(* IEC 61131-3 sources: STAR-PLC-Agent/results/raw/batch_fresh_20261114/PUB015/functional/attempt_0001, 1 file *)

(* ---- test_program.st ---- *)
PROGRAM PLC_PRG
VAR
 BenchStep : UDINT := 0;
 BenchCalls : UDINT := 0;
 BenchDone : BOOL := FALSE;
 BenchUut0 : FB_Task;
 BenchUut1 : FB_Task;
 BenchUut2 : FB_Task;
 BenchUut3 : FB_Task;
 BenchUut4 : FB_Task;
 BenchUut5 : FB_Task;
 BenchUut6 : FB_Task;
 BenchUut7 : FB_Task;
 BenchUut8 : FB_Task;
 BenchUut9 : FB_Task;
 BenchUut10 : FB_Task;
 BenchUut11 : FB_Task;
 BenchUut12 : FB_Task;
 TraceIn_estop : ARRAY[0..126] OF BOOL;
 TraceIn_opeMode : ARRAY[0..126] OF BOOL;
 TraceIn_valveAStart : ARRAY[0..126] OF BOOL;
 TraceIn_valveBStart : ARRAY[0..126] OF BOOL;
 TraceIn_valveCStart : ARRAY[0..126] OF BOOL;
 TraceIn_valveDStart : ARRAY[0..126] OF BOOL;
 TraceIn_mixMotorStart : ARRAY[0..126] OF BOOL;
 TraceIn_autoStart : ARRAY[0..126] OF BOOL;
 TraceIn_processMode : ARRAY[0..126] OF BOOL;
 TraceIn_levelSensor : ARRAY[0..126] OF INT;
 TraceIn_mixMotorComplete : ARRAY[0..126] OF BOOL;
 TraceOut_valveARun : ARRAY[0..126] OF BOOL;
 TraceOut_valveBRun : ARRAY[0..126] OF BOOL;
 TraceOut_valveCRun : ARRAY[0..126] OF BOOL;
 TraceOut_valveDRun : ARRAY[0..126] OF BOOL;
 TraceOut_mixMotorRun : ARRAY[0..126] OF BOOL;
END_VAR

IF NOT BenchDone THEN
 CASE BenchStep OF
 0:
   BenchUut0.estop := TRUE;
   BenchUut0.opeMode := FALSE;
   BenchUut0.valveAStart := FALSE;
   BenchUut0.valveBStart := FALSE;
   BenchUut0.valveCStart := FALSE;
   BenchUut0.valveDStart := FALSE;
   BenchUut0.mixMotorStart := FALSE;
   BenchUut0.autoStart := FALSE;
   BenchUut0.processMode := FALSE;
   BenchUut0.levelSensor := INT#0;
   BenchUut0.mixMotorComplete := FALSE;
   TraceIn_estop[0] := BenchUut0.estop;
   TraceIn_opeMode[0] := BenchUut0.opeMode;
   TraceIn_valveAStart[0] := BenchUut0.valveAStart;
   TraceIn_valveBStart[0] := BenchUut0.valveBStart;
   TraceIn_valveCStart[0] := BenchUut0.valveCStart;
   TraceIn_valveDStart[0] := BenchUut0.valveDStart;
   TraceIn_mixMotorStart[0] := BenchUut0.mixMotorStart;
   TraceIn_autoStart[0] := BenchUut0.autoStart;
   TraceIn_processMode[0] := BenchUut0.processMode;
   TraceIn_levelSensor[0] := BenchUut0.levelSensor;
   TraceIn_mixMotorComplete[0] := BenchUut0.mixMotorComplete;
   BenchUut0();
   TraceOut_valveARun[0] := BenchUut0.valveARun;
   TraceOut_valveBRun[0] := BenchUut0.valveBRun;
   TraceOut_valveCRun[0] := BenchUut0.valveCRun;
   TraceOut_valveDRun[0] := BenchUut0.valveDRun;
   TraceOut_mixMotorRun[0] := BenchUut0.mixMotorRun;
   BenchCalls := BenchCalls + 1;
 1:
   BenchUut0.estop := TRUE;
   BenchUut0.opeMode := FALSE;
   BenchUut0.valveAStart := TRUE;
   BenchUut0.valveBStart := FALSE;
   BenchUut0.valveCStart := FALSE;
   BenchUut0.valveDStart := FALSE;
   BenchUut0.mixMotorStart := FALSE;
   BenchUut0.autoStart := FALSE;
   BenchUut0.processMode := FALSE;
   BenchUut0.levelSensor := INT#0;
   BenchUut0.mixMotorComplete := FALSE;
   TraceIn_estop[1] := BenchUut0.estop;
   TraceIn_opeMode[1] := BenchUut0.opeMode;
   TraceIn_valveAStart[1] := BenchUut0.valveAStart;
   TraceIn_valveBStart[1] := BenchUut0.valveBStart;
   TraceIn_valveCStart[1] := BenchUut0.valveCStart;
   TraceIn_valveDStart[1] := BenchUut0.valveDStart;
   TraceIn_mixMotorStart[1] := BenchUut0.mixMotorStart;
   TraceIn_autoStart[1] := BenchUut0.autoStart;
   TraceIn_processMode[1] := BenchUut0.processMode;
   TraceIn_levelSensor[1] := BenchUut0.levelSensor;
   TraceIn_mixMotorComplete[1] := BenchUut0.mixMotorComplete;
   BenchUut0();
   TraceOut_valveARun[1] := BenchUut0.valveARun;
   TraceOut_valveBRun[1] := BenchUut0.valveBRun;
   TraceOut_valveCRun[1] := BenchUut0.valveCRun;
   TraceOut_valveDRun[1] := BenchUut0.valveDRun;
   TraceOut_mixMotorRun[1] := BenchUut0.mixMotorRun;
   BenchCalls := BenchCalls + 1;
 2:
   BenchUut0.estop := TRUE;
   BenchUut0.opeMode := FALSE;
   BenchUut0.valveAStart := TRUE;
   BenchUut0.valveBStart := FALSE;
   BenchUut0.valveCStart := FALSE;
   BenchUut0.valveDStart := FALSE;
   BenchUut0.mixMotorStart := FALSE;
   BenchUut0.autoStart := FALSE;
   BenchUut0.processMode := FALSE;
   BenchUut0.levelSensor := INT#0;
   BenchUut0.mixMotorComplete := FALSE;
   TraceIn_estop[2] := BenchUut0.estop;
   TraceIn_opeMode[2] := BenchUut0.opeMode;
   TraceIn_valveAStart[2] := BenchUut0.valveAStart;
   TraceIn_valveBStart[2] := BenchUut0.valveBStart;
   TraceIn_valveCStart[2] := BenchUut0.valveCStart;
   TraceIn_valveDStart[2] := BenchUut0.valveDStart;
   TraceIn_mixMotorStart[2] := BenchUut0.mixMotorStart;
   TraceIn_autoStart[2] := BenchUut0.autoStart;
   TraceIn_processMode[2] := BenchUut0.processMode;
   TraceIn_levelSensor[2] := BenchUut0.levelSensor;
   TraceIn_mixMotorComplete[2] := BenchUut0.mixMotorComplete;
   BenchUut0();
   TraceOut_valveARun[2] := BenchUut0.valveARun;
   TraceOut_valveBRun[2] := BenchUut0.valveBRun;
   TraceOut_valveCRun[2] := BenchUut0.valveCRun;
   TraceOut_valveDRun[2] := BenchUut0.valveDRun;
   TraceOut_mixMotorRun[2] := BenchUut0.mixMotorRun;
   BenchCalls := BenchCalls + 1;
 3:
   BenchUut0.estop := TRUE;
   BenchUut0.opeMode := FALSE;
   BenchUut0.valveAStart := FALSE;
   BenchUut0.valveBStart := FALSE;
   BenchUut0.valveCStart := FALSE;
   BenchUut0.valveDStart := FALSE;
   BenchUut0.mixMotorStart := FALSE;
   BenchUut0.autoStart := FALSE;
   BenchUut0.processMode := FALSE;
   BenchUut0.levelSensor := INT#0;
   BenchUut0.mixMotorComplete := FALSE;
   TraceIn_estop[3] := BenchUut0.estop;
   TraceIn_opeMode[3] := BenchUut0.opeMode;
   TraceIn_valveAStart[3] := BenchUut0.valveAStart;
   TraceIn_valveBStart[3] := BenchUut0.valveBStart;
   TraceIn_valveCStart[3] := BenchUut0.valveCStart;
   TraceIn_valveDStart[3] := BenchUut0.valveDStart;
   TraceIn_mixMotorStart[3] := BenchUut0.mixMotorStart;
   TraceIn_autoStart[3] := BenchUut0.autoStart;
   TraceIn_processMode[3] := BenchUut0.processMode;
   TraceIn_levelSensor[3] := BenchUut0.levelSensor;
   TraceIn_mixMotorComplete[3] := BenchUut0.mixMotorComplete;
   BenchUut0();
   TraceOut_valveARun[3] := BenchUut0.valveARun;
   TraceOut_valveBRun[3] := BenchUut0.valveBRun;
   TraceOut_valveCRun[3] := BenchUut0.valveCRun;
   TraceOut_valveDRun[3] := BenchUut0.valveDRun;
   TraceOut_mixMotorRun[3] := BenchUut0.mixMotorRun;
   BenchCalls := BenchCalls + 1;
 4:
   BenchUut0.estop := TRUE;
   BenchUut0.opeMode := FALSE;
   BenchUut0.valveAStart := TRUE;
   BenchUut0.valveBStart := FALSE;
   BenchUut0.valveCStart := FALSE;
   BenchUut0.valveDStart := FALSE;
   BenchUut0.mixMotorStart := FALSE;
   BenchUut0.autoStart := FALSE;
   BenchUut0.processMode := FALSE;
   BenchUut0.levelSensor := INT#0;
   BenchUut0.mixMotorComplete := FALSE;
   TraceIn_estop[4] := BenchUut0.estop;
   TraceIn_opeMode[4] := BenchUut0.opeMode;
   TraceIn_valveAStart[4] := BenchUut0.valveAStart;
   TraceIn_valveBStart[4] := BenchUut0.valveBStart;
   TraceIn_valveCStart[4] := BenchUut0.valveCStart;
   TraceIn_valveDStart[4] := BenchUut0.valveDStart;
   TraceIn_mixMotorStart[4] := BenchUut0.mixMotorStart;
   TraceIn_autoStart[4] := BenchUut0.autoStart;
   TraceIn_processMode[4] := BenchUut0.processMode;
   TraceIn_levelSensor[4] := BenchUut0.levelSensor;
   TraceIn_mixMotorComplete[4] := BenchUut0.mixMotorComplete;
   BenchUut0();
   TraceOut_valveARun[4] := BenchUut0.valveARun;
   TraceOut_valveBRun[4] := BenchUut0.valveBRun;
   TraceOut_valveCRun[4] := BenchUut0.valveCRun;
   TraceOut_valveDRun[4] := BenchUut0.valveDRun;
   TraceOut_mixMotorRun[4] := BenchUut0.mixMotorRun;
   BenchCalls := BenchCalls + 1;
 5:
   BenchUut0.estop := TRUE;
   BenchUut0.opeMode := FALSE;
   BenchUut0.valveAStart := FALSE;
   BenchUut0.valveBStart := TRUE;
   BenchUut0.valveCStart := TRUE;
   BenchUut0.valveDStart := TRUE;
   BenchUut0.mixMotorStart := TRUE;
   BenchUut0.autoStart := FALSE;
   BenchUut0.processMode := FALSE;
   BenchUut0.levelSensor := INT#0;
   BenchUut0.mixMotorComplete := FALSE;
   TraceIn_estop[5] := BenchUut0.estop;
   TraceIn_opeMode[5] := BenchUut0.opeMode;
   TraceIn_valveAStart[5] := BenchUut0.valveAStart;
   TraceIn_valveBStart[5] := BenchUut0.valveBStart;
   TraceIn_valveCStart[5] := BenchUut0.valveCStart;
   TraceIn_valveDStart[5] := BenchUut0.valveDStart;
   TraceIn_mixMotorStart[5] := BenchUut0.mixMotorStart;
   TraceIn_autoStart[5] := BenchUut0.autoStart;
   TraceIn_processMode[5] := BenchUut0.processMode;
   TraceIn_levelSensor[5] := BenchUut0.levelSensor;
   TraceIn_mixMotorComplete[5] := BenchUut0.mixMotorComplete;
   BenchUut0();
   TraceOut_valveARun[5] := BenchUut0.valveARun;
   TraceOut_valveBRun[5] := BenchUut0.valveBRun;
   TraceOut_valveCRun[5] := BenchUut0.valveCRun;
   TraceOut_valveDRun[5] := BenchUut0.valveDRun;
   TraceOut_mixMotorRun[5] := BenchUut0.mixMotorRun;
   BenchCalls := BenchCalls + 1;
 6:
   BenchUut0.estop := FALSE;
   BenchUut0.opeMode := FALSE;
   BenchUut0.valveAStart := FALSE;
   BenchUut0.valveBStart := FALSE;
   BenchUut0.valveCStart := FALSE;
   BenchUut0.valveDStart := FALSE;
   BenchUut0.mixMotorStart := FALSE;
   BenchUut0.autoStart := FALSE;
   BenchUut0.processMode := FALSE;
   BenchUut0.levelSensor := INT#0;
   BenchUut0.mixMotorComplete := FALSE;
   TraceIn_estop[6] := BenchUut0.estop;
   TraceIn_opeMode[6] := BenchUut0.opeMode;
   TraceIn_valveAStart[6] := BenchUut0.valveAStart;
   TraceIn_valveBStart[6] := BenchUut0.valveBStart;
   TraceIn_valveCStart[6] := BenchUut0.valveCStart;
   TraceIn_valveDStart[6] := BenchUut0.valveDStart;
   TraceIn_mixMotorStart[6] := BenchUut0.mixMotorStart;
   TraceIn_autoStart[6] := BenchUut0.autoStart;
   TraceIn_processMode[6] := BenchUut0.processMode;
   TraceIn_levelSensor[6] := BenchUut0.levelSensor;
   TraceIn_mixMotorComplete[6] := BenchUut0.mixMotorComplete;
   BenchUut0();
   TraceOut_valveARun[6] := BenchUut0.valveARun;
   TraceOut_valveBRun[6] := BenchUut0.valveBRun;
   TraceOut_valveCRun[6] := BenchUut0.valveCRun;
   TraceOut_valveDRun[6] := BenchUut0.valveDRun;
   TraceOut_mixMotorRun[6] := BenchUut0.mixMotorRun;
   BenchCalls := BenchCalls + 1;
 7:
   BenchUut1.estop := TRUE;
   BenchUut1.opeMode := TRUE;
   BenchUut1.valveAStart := FALSE;
   BenchUut1.valveBStart := FALSE;
   BenchUut1.valveCStart := FALSE;
   BenchUut1.valveDStart := FALSE;
   BenchUut1.mixMotorStart := FALSE;
   BenchUut1.autoStart := FALSE;
   BenchUut1.processMode := FALSE;
   BenchUut1.levelSensor := INT#0;
   BenchUut1.mixMotorComplete := FALSE;
   TraceIn_estop[7] := BenchUut1.estop;
   TraceIn_opeMode[7] := BenchUut1.opeMode;
   TraceIn_valveAStart[7] := BenchUut1.valveAStart;
   TraceIn_valveBStart[7] := BenchUut1.valveBStart;
   TraceIn_valveCStart[7] := BenchUut1.valveCStart;
   TraceIn_valveDStart[7] := BenchUut1.valveDStart;
   TraceIn_mixMotorStart[7] := BenchUut1.mixMotorStart;
   TraceIn_autoStart[7] := BenchUut1.autoStart;
   TraceIn_processMode[7] := BenchUut1.processMode;
   TraceIn_levelSensor[7] := BenchUut1.levelSensor;
   TraceIn_mixMotorComplete[7] := BenchUut1.mixMotorComplete;
   BenchUut1();
   TraceOut_valveARun[7] := BenchUut1.valveARun;
   TraceOut_valveBRun[7] := BenchUut1.valveBRun;
   TraceOut_valveCRun[7] := BenchUut1.valveCRun;
   TraceOut_valveDRun[7] := BenchUut1.valveDRun;
   TraceOut_mixMotorRun[7] := BenchUut1.mixMotorRun;
   BenchCalls := BenchCalls + 1;
 8:
   BenchUut1.estop := TRUE;
   BenchUut1.opeMode := TRUE;
   BenchUut1.valveAStart := FALSE;
   BenchUut1.valveBStart := FALSE;
   BenchUut1.valveCStart := FALSE;
   BenchUut1.valveDStart := FALSE;
   BenchUut1.mixMotorStart := FALSE;
   BenchUut1.autoStart := TRUE;
   BenchUut1.processMode := FALSE;
   BenchUut1.levelSensor := INT#0;
   BenchUut1.mixMotorComplete := FALSE;
   TraceIn_estop[8] := BenchUut1.estop;
   TraceIn_opeMode[8] := BenchUut1.opeMode;
   TraceIn_valveAStart[8] := BenchUut1.valveAStart;
   TraceIn_valveBStart[8] := BenchUut1.valveBStart;
   TraceIn_valveCStart[8] := BenchUut1.valveCStart;
   TraceIn_valveDStart[8] := BenchUut1.valveDStart;
   TraceIn_mixMotorStart[8] := BenchUut1.mixMotorStart;
   TraceIn_autoStart[8] := BenchUut1.autoStart;
   TraceIn_processMode[8] := BenchUut1.processMode;
   TraceIn_levelSensor[8] := BenchUut1.levelSensor;
   TraceIn_mixMotorComplete[8] := BenchUut1.mixMotorComplete;
   BenchUut1();
   TraceOut_valveARun[8] := BenchUut1.valveARun;
   TraceOut_valveBRun[8] := BenchUut1.valveBRun;
   TraceOut_valveCRun[8] := BenchUut1.valveCRun;
   TraceOut_valveDRun[8] := BenchUut1.valveDRun;
   TraceOut_mixMotorRun[8] := BenchUut1.mixMotorRun;
   BenchCalls := BenchCalls + 1;
 9:
   BenchUut1.estop := TRUE;
   BenchUut1.opeMode := TRUE;
   BenchUut1.valveAStart := FALSE;
   BenchUut1.valveBStart := FALSE;
   BenchUut1.valveCStart := FALSE;
   BenchUut1.valveDStart := FALSE;
   BenchUut1.mixMotorStart := FALSE;
   BenchUut1.autoStart := FALSE;
   BenchUut1.processMode := FALSE;
   BenchUut1.levelSensor := INT#49;
   BenchUut1.mixMotorComplete := FALSE;
   TraceIn_estop[9] := BenchUut1.estop;
   TraceIn_opeMode[9] := BenchUut1.opeMode;
   TraceIn_valveAStart[9] := BenchUut1.valveAStart;
   TraceIn_valveBStart[9] := BenchUut1.valveBStart;
   TraceIn_valveCStart[9] := BenchUut1.valveCStart;
   TraceIn_valveDStart[9] := BenchUut1.valveDStart;
   TraceIn_mixMotorStart[9] := BenchUut1.mixMotorStart;
   TraceIn_autoStart[9] := BenchUut1.autoStart;
   TraceIn_processMode[9] := BenchUut1.processMode;
   TraceIn_levelSensor[9] := BenchUut1.levelSensor;
   TraceIn_mixMotorComplete[9] := BenchUut1.mixMotorComplete;
   BenchUut1();
   TraceOut_valveARun[9] := BenchUut1.valveARun;
   TraceOut_valveBRun[9] := BenchUut1.valveBRun;
   TraceOut_valveCRun[9] := BenchUut1.valveCRun;
   TraceOut_valveDRun[9] := BenchUut1.valveDRun;
   TraceOut_mixMotorRun[9] := BenchUut1.mixMotorRun;
   BenchCalls := BenchCalls + 1;
 10:
   BenchUut1.estop := TRUE;
   BenchUut1.opeMode := TRUE;
   BenchUut1.valveAStart := FALSE;
   BenchUut1.valveBStart := FALSE;
   BenchUut1.valveCStart := FALSE;
   BenchUut1.valveDStart := FALSE;
   BenchUut1.mixMotorStart := FALSE;
   BenchUut1.autoStart := FALSE;
   BenchUut1.processMode := FALSE;
   BenchUut1.levelSensor := INT#50;
   BenchUut1.mixMotorComplete := FALSE;
   TraceIn_estop[10] := BenchUut1.estop;
   TraceIn_opeMode[10] := BenchUut1.opeMode;
   TraceIn_valveAStart[10] := BenchUut1.valveAStart;
   TraceIn_valveBStart[10] := BenchUut1.valveBStart;
   TraceIn_valveCStart[10] := BenchUut1.valveCStart;
   TraceIn_valveDStart[10] := BenchUut1.valveDStart;
   TraceIn_mixMotorStart[10] := BenchUut1.mixMotorStart;
   TraceIn_autoStart[10] := BenchUut1.autoStart;
   TraceIn_processMode[10] := BenchUut1.processMode;
   TraceIn_levelSensor[10] := BenchUut1.levelSensor;
   TraceIn_mixMotorComplete[10] := BenchUut1.mixMotorComplete;
   BenchUut1();
   TraceOut_valveARun[10] := BenchUut1.valveARun;
   TraceOut_valveBRun[10] := BenchUut1.valveBRun;
   TraceOut_valveCRun[10] := BenchUut1.valveCRun;
   TraceOut_valveDRun[10] := BenchUut1.valveDRun;
   TraceOut_mixMotorRun[10] := BenchUut1.mixMotorRun;
   BenchCalls := BenchCalls + 1;
 11:
   BenchUut1.estop := TRUE;
   BenchUut1.opeMode := TRUE;
   BenchUut1.valveAStart := FALSE;
   BenchUut1.valveBStart := FALSE;
   BenchUut1.valveCStart := FALSE;
   BenchUut1.valveDStart := FALSE;
   BenchUut1.mixMotorStart := FALSE;
   BenchUut1.autoStart := FALSE;
   BenchUut1.processMode := FALSE;
   BenchUut1.levelSensor := INT#80;
   BenchUut1.mixMotorComplete := FALSE;
   TraceIn_estop[11] := BenchUut1.estop;
   TraceIn_opeMode[11] := BenchUut1.opeMode;
   TraceIn_valveAStart[11] := BenchUut1.valveAStart;
   TraceIn_valveBStart[11] := BenchUut1.valveBStart;
   TraceIn_valveCStart[11] := BenchUut1.valveCStart;
   TraceIn_valveDStart[11] := BenchUut1.valveDStart;
   TraceIn_mixMotorStart[11] := BenchUut1.mixMotorStart;
   TraceIn_autoStart[11] := BenchUut1.autoStart;
   TraceIn_processMode[11] := BenchUut1.processMode;
   TraceIn_levelSensor[11] := BenchUut1.levelSensor;
   TraceIn_mixMotorComplete[11] := BenchUut1.mixMotorComplete;
   BenchUut1();
   TraceOut_valveARun[11] := BenchUut1.valveARun;
   TraceOut_valveBRun[11] := BenchUut1.valveBRun;
   TraceOut_valveCRun[11] := BenchUut1.valveCRun;
   TraceOut_valveDRun[11] := BenchUut1.valveDRun;
   TraceOut_mixMotorRun[11] := BenchUut1.mixMotorRun;
   BenchCalls := BenchCalls + 1;
 12:
   BenchUut1.estop := TRUE;
   BenchUut1.opeMode := TRUE;
   BenchUut1.valveAStart := FALSE;
   BenchUut1.valveBStart := FALSE;
   BenchUut1.valveCStart := FALSE;
   BenchUut1.valveDStart := FALSE;
   BenchUut1.mixMotorStart := FALSE;
   BenchUut1.autoStart := FALSE;
   BenchUut1.processMode := FALSE;
   BenchUut1.levelSensor := INT#80;
   BenchUut1.mixMotorComplete := TRUE;
   TraceIn_estop[12] := BenchUut1.estop;
   TraceIn_opeMode[12] := BenchUut1.opeMode;
   TraceIn_valveAStart[12] := BenchUut1.valveAStart;
   TraceIn_valveBStart[12] := BenchUut1.valveBStart;
   TraceIn_valveCStart[12] := BenchUut1.valveCStart;
   TraceIn_valveDStart[12] := BenchUut1.valveDStart;
   TraceIn_mixMotorStart[12] := BenchUut1.mixMotorStart;
   TraceIn_autoStart[12] := BenchUut1.autoStart;
   TraceIn_processMode[12] := BenchUut1.processMode;
   TraceIn_levelSensor[12] := BenchUut1.levelSensor;
   TraceIn_mixMotorComplete[12] := BenchUut1.mixMotorComplete;
   BenchUut1();
   TraceOut_valveARun[12] := BenchUut1.valveARun;
   TraceOut_valveBRun[12] := BenchUut1.valveBRun;
   TraceOut_valveCRun[12] := BenchUut1.valveCRun;
   TraceOut_valveDRun[12] := BenchUut1.valveDRun;
   TraceOut_mixMotorRun[12] := BenchUut1.mixMotorRun;
   BenchCalls := BenchCalls + 1;
 13:
   BenchUut1.estop := FALSE;
   BenchUut1.opeMode := TRUE;
   BenchUut1.valveAStart := FALSE;
   BenchUut1.valveBStart := FALSE;
   BenchUut1.valveCStart := FALSE;
   BenchUut1.valveDStart := FALSE;
   BenchUut1.mixMotorStart := FALSE;
   BenchUut1.autoStart := FALSE;
   BenchUut1.processMode := FALSE;
   BenchUut1.levelSensor := INT#0;
   BenchUut1.mixMotorComplete := FALSE;
   TraceIn_estop[13] := BenchUut1.estop;
   TraceIn_opeMode[13] := BenchUut1.opeMode;
   TraceIn_valveAStart[13] := BenchUut1.valveAStart;
   TraceIn_valveBStart[13] := BenchUut1.valveBStart;
   TraceIn_valveCStart[13] := BenchUut1.valveCStart;
   TraceIn_valveDStart[13] := BenchUut1.valveDStart;
   TraceIn_mixMotorStart[13] := BenchUut1.mixMotorStart;
   TraceIn_autoStart[13] := BenchUut1.autoStart;
   TraceIn_processMode[13] := BenchUut1.processMode;
   TraceIn_levelSensor[13] := BenchUut1.levelSensor;
   TraceIn_mixMotorComplete[13] := BenchUut1.mixMotorComplete;
   BenchUut1();
   TraceOut_valveARun[13] := BenchUut1.valveARun;
   TraceOut_valveBRun[13] := BenchUut1.valveBRun;
   TraceOut_valveCRun[13] := BenchUut1.valveCRun;
   TraceOut_valveDRun[13] := BenchUut1.valveDRun;
   TraceOut_mixMotorRun[13] := BenchUut1.mixMotorRun;
   BenchCalls := BenchCalls + 1;
 14:
   BenchUut2.estop := TRUE;
   BenchUut2.opeMode := TRUE;
   BenchUut2.valveAStart := FALSE;
   BenchUut2.valveBStart := FALSE;
   BenchUut2.valveCStart := FALSE;
   BenchUut2.valveDStart := FALSE;
   BenchUut2.mixMotorStart := FALSE;
   BenchUut2.autoStart := FALSE;
   BenchUut2.processMode := FALSE;
   BenchUut2.levelSensor := INT#0;
   BenchUut2.mixMotorComplete := FALSE;
   TraceIn_estop[14] := BenchUut2.estop;
   TraceIn_opeMode[14] := BenchUut2.opeMode;
   TraceIn_valveAStart[14] := BenchUut2.valveAStart;
   TraceIn_valveBStart[14] := BenchUut2.valveBStart;
   TraceIn_valveCStart[14] := BenchUut2.valveCStart;
   TraceIn_valveDStart[14] := BenchUut2.valveDStart;
   TraceIn_mixMotorStart[14] := BenchUut2.mixMotorStart;
   TraceIn_autoStart[14] := BenchUut2.autoStart;
   TraceIn_processMode[14] := BenchUut2.processMode;
   TraceIn_levelSensor[14] := BenchUut2.levelSensor;
   TraceIn_mixMotorComplete[14] := BenchUut2.mixMotorComplete;
   BenchUut2();
   TraceOut_valveARun[14] := BenchUut2.valveARun;
   TraceOut_valveBRun[14] := BenchUut2.valveBRun;
   TraceOut_valveCRun[14] := BenchUut2.valveCRun;
   TraceOut_valveDRun[14] := BenchUut2.valveDRun;
   TraceOut_mixMotorRun[14] := BenchUut2.mixMotorRun;
   BenchCalls := BenchCalls + 1;
 15:
   BenchUut2.estop := TRUE;
   BenchUut2.opeMode := TRUE;
   BenchUut2.valveAStart := FALSE;
   BenchUut2.valveBStart := FALSE;
   BenchUut2.valveCStart := FALSE;
   BenchUut2.valveDStart := FALSE;
   BenchUut2.mixMotorStart := FALSE;
   BenchUut2.autoStart := TRUE;
   BenchUut2.processMode := TRUE;
   BenchUut2.levelSensor := INT#0;
   BenchUut2.mixMotorComplete := FALSE;
   TraceIn_estop[15] := BenchUut2.estop;
   TraceIn_opeMode[15] := BenchUut2.opeMode;
   TraceIn_valveAStart[15] := BenchUut2.valveAStart;
   TraceIn_valveBStart[15] := BenchUut2.valveBStart;
   TraceIn_valveCStart[15] := BenchUut2.valveCStart;
   TraceIn_valveDStart[15] := BenchUut2.valveDStart;
   TraceIn_mixMotorStart[15] := BenchUut2.mixMotorStart;
   TraceIn_autoStart[15] := BenchUut2.autoStart;
   TraceIn_processMode[15] := BenchUut2.processMode;
   TraceIn_levelSensor[15] := BenchUut2.levelSensor;
   TraceIn_mixMotorComplete[15] := BenchUut2.mixMotorComplete;
   BenchUut2();
   TraceOut_valveARun[15] := BenchUut2.valveARun;
   TraceOut_valveBRun[15] := BenchUut2.valveBRun;
   TraceOut_valveCRun[15] := BenchUut2.valveCRun;
   TraceOut_valveDRun[15] := BenchUut2.valveDRun;
   TraceOut_mixMotorRun[15] := BenchUut2.mixMotorRun;
   BenchCalls := BenchCalls + 1;
 16:
   BenchUut2.estop := TRUE;
   BenchUut2.opeMode := TRUE;
   BenchUut2.valveAStart := FALSE;
   BenchUut2.valveBStart := FALSE;
   BenchUut2.valveCStart := FALSE;
   BenchUut2.valveDStart := FALSE;
   BenchUut2.mixMotorStart := FALSE;
   BenchUut2.autoStart := FALSE;
   BenchUut2.processMode := TRUE;
   BenchUut2.levelSensor := INT#55;
   BenchUut2.mixMotorComplete := FALSE;
   TraceIn_estop[16] := BenchUut2.estop;
   TraceIn_opeMode[16] := BenchUut2.opeMode;
   TraceIn_valveAStart[16] := BenchUut2.valveAStart;
   TraceIn_valveBStart[16] := BenchUut2.valveBStart;
   TraceIn_valveCStart[16] := BenchUut2.valveCStart;
   TraceIn_valveDStart[16] := BenchUut2.valveDStart;
   TraceIn_mixMotorStart[16] := BenchUut2.mixMotorStart;
   TraceIn_autoStart[16] := BenchUut2.autoStart;
   TraceIn_processMode[16] := BenchUut2.processMode;
   TraceIn_levelSensor[16] := BenchUut2.levelSensor;
   TraceIn_mixMotorComplete[16] := BenchUut2.mixMotorComplete;
   BenchUut2();
   TraceOut_valveARun[16] := BenchUut2.valveARun;
   TraceOut_valveBRun[16] := BenchUut2.valveBRun;
   TraceOut_valveCRun[16] := BenchUut2.valveCRun;
   TraceOut_valveDRun[16] := BenchUut2.valveDRun;
   TraceOut_mixMotorRun[16] := BenchUut2.mixMotorRun;
   BenchCalls := BenchCalls + 1;
 17:
   BenchUut2.estop := TRUE;
   BenchUut2.opeMode := TRUE;
   BenchUut2.valveAStart := FALSE;
   BenchUut2.valveBStart := FALSE;
   BenchUut2.valveCStart := FALSE;
   BenchUut2.valveDStart := FALSE;
   BenchUut2.mixMotorStart := FALSE;
   BenchUut2.autoStart := FALSE;
   BenchUut2.processMode := TRUE;
   BenchUut2.levelSensor := INT#85;
   BenchUut2.mixMotorComplete := FALSE;
   TraceIn_estop[17] := BenchUut2.estop;
   TraceIn_opeMode[17] := BenchUut2.opeMode;
   TraceIn_valveAStart[17] := BenchUut2.valveAStart;
   TraceIn_valveBStart[17] := BenchUut2.valveBStart;
   TraceIn_valveCStart[17] := BenchUut2.valveCStart;
   TraceIn_valveDStart[17] := BenchUut2.valveDStart;
   TraceIn_mixMotorStart[17] := BenchUut2.mixMotorStart;
   TraceIn_autoStart[17] := BenchUut2.autoStart;
   TraceIn_processMode[17] := BenchUut2.processMode;
   TraceIn_levelSensor[17] := BenchUut2.levelSensor;
   TraceIn_mixMotorComplete[17] := BenchUut2.mixMotorComplete;
   BenchUut2();
   TraceOut_valveARun[17] := BenchUut2.valveARun;
   TraceOut_valveBRun[17] := BenchUut2.valveBRun;
   TraceOut_valveCRun[17] := BenchUut2.valveCRun;
   TraceOut_valveDRun[17] := BenchUut2.valveDRun;
   TraceOut_mixMotorRun[17] := BenchUut2.mixMotorRun;
   BenchCalls := BenchCalls + 1;
 18:
   BenchUut2.estop := TRUE;
   BenchUut2.opeMode := TRUE;
   BenchUut2.valveAStart := FALSE;
   BenchUut2.valveBStart := FALSE;
   BenchUut2.valveCStart := FALSE;
   BenchUut2.valveDStart := FALSE;
   BenchUut2.mixMotorStart := FALSE;
   BenchUut2.autoStart := FALSE;
   BenchUut2.processMode := TRUE;
   BenchUut2.levelSensor := INT#99;
   BenchUut2.mixMotorComplete := FALSE;
   TraceIn_estop[18] := BenchUut2.estop;
   TraceIn_opeMode[18] := BenchUut2.opeMode;
   TraceIn_valveAStart[18] := BenchUut2.valveAStart;
   TraceIn_valveBStart[18] := BenchUut2.valveBStart;
   TraceIn_valveCStart[18] := BenchUut2.valveCStart;
   TraceIn_valveDStart[18] := BenchUut2.valveDStart;
   TraceIn_mixMotorStart[18] := BenchUut2.mixMotorStart;
   TraceIn_autoStart[18] := BenchUut2.autoStart;
   TraceIn_processMode[18] := BenchUut2.processMode;
   TraceIn_levelSensor[18] := BenchUut2.levelSensor;
   TraceIn_mixMotorComplete[18] := BenchUut2.mixMotorComplete;
   BenchUut2();
   TraceOut_valveARun[18] := BenchUut2.valveARun;
   TraceOut_valveBRun[18] := BenchUut2.valveBRun;
   TraceOut_valveCRun[18] := BenchUut2.valveCRun;
   TraceOut_valveDRun[18] := BenchUut2.valveDRun;
   TraceOut_mixMotorRun[18] := BenchUut2.mixMotorRun;
   BenchCalls := BenchCalls + 1;
 19:
   BenchUut2.estop := TRUE;
   BenchUut2.opeMode := TRUE;
   BenchUut2.valveAStart := FALSE;
   BenchUut2.valveBStart := FALSE;
   BenchUut2.valveCStart := FALSE;
   BenchUut2.valveDStart := FALSE;
   BenchUut2.mixMotorStart := FALSE;
   BenchUut2.autoStart := FALSE;
   BenchUut2.processMode := TRUE;
   BenchUut2.levelSensor := INT#100;
   BenchUut2.mixMotorComplete := FALSE;
   TraceIn_estop[19] := BenchUut2.estop;
   TraceIn_opeMode[19] := BenchUut2.opeMode;
   TraceIn_valveAStart[19] := BenchUut2.valveAStart;
   TraceIn_valveBStart[19] := BenchUut2.valveBStart;
   TraceIn_valveCStart[19] := BenchUut2.valveCStart;
   TraceIn_valveDStart[19] := BenchUut2.valveDStart;
   TraceIn_mixMotorStart[19] := BenchUut2.mixMotorStart;
   TraceIn_autoStart[19] := BenchUut2.autoStart;
   TraceIn_processMode[19] := BenchUut2.processMode;
   TraceIn_levelSensor[19] := BenchUut2.levelSensor;
   TraceIn_mixMotorComplete[19] := BenchUut2.mixMotorComplete;
   BenchUut2();
   TraceOut_valveARun[19] := BenchUut2.valveARun;
   TraceOut_valveBRun[19] := BenchUut2.valveBRun;
   TraceOut_valveCRun[19] := BenchUut2.valveCRun;
   TraceOut_valveDRun[19] := BenchUut2.valveDRun;
   TraceOut_mixMotorRun[19] := BenchUut2.mixMotorRun;
   BenchCalls := BenchCalls + 1;
 20:
   BenchUut2.estop := FALSE;
   BenchUut2.opeMode := TRUE;
   BenchUut2.valveAStart := FALSE;
   BenchUut2.valveBStart := FALSE;
   BenchUut2.valveCStart := FALSE;
   BenchUut2.valveDStart := FALSE;
   BenchUut2.mixMotorStart := FALSE;
   BenchUut2.autoStart := FALSE;
   BenchUut2.processMode := TRUE;
   BenchUut2.levelSensor := INT#0;
   BenchUut2.mixMotorComplete := TRUE;
   TraceIn_estop[20] := BenchUut2.estop;
   TraceIn_opeMode[20] := BenchUut2.opeMode;
   TraceIn_valveAStart[20] := BenchUut2.valveAStart;
   TraceIn_valveBStart[20] := BenchUut2.valveBStart;
   TraceIn_valveCStart[20] := BenchUut2.valveCStart;
   TraceIn_valveDStart[20] := BenchUut2.valveDStart;
   TraceIn_mixMotorStart[20] := BenchUut2.mixMotorStart;
   TraceIn_autoStart[20] := BenchUut2.autoStart;
   TraceIn_processMode[20] := BenchUut2.processMode;
   TraceIn_levelSensor[20] := BenchUut2.levelSensor;
   TraceIn_mixMotorComplete[20] := BenchUut2.mixMotorComplete;
   BenchUut2();
   TraceOut_valveARun[20] := BenchUut2.valveARun;
   TraceOut_valveBRun[20] := BenchUut2.valveBRun;
   TraceOut_valveCRun[20] := BenchUut2.valveCRun;
   TraceOut_valveDRun[20] := BenchUut2.valveDRun;
   TraceOut_mixMotorRun[20] := BenchUut2.mixMotorRun;
   BenchCalls := BenchCalls + 1;
 21:
   BenchUut2.estop := TRUE;
   BenchUut2.opeMode := TRUE;
   BenchUut2.valveAStart := FALSE;
   BenchUut2.valveBStart := FALSE;
   BenchUut2.valveCStart := FALSE;
   BenchUut2.valveDStart := FALSE;
   BenchUut2.mixMotorStart := FALSE;
   BenchUut2.autoStart := FALSE;
   BenchUut2.processMode := TRUE;
   BenchUut2.levelSensor := INT#0;
   BenchUut2.mixMotorComplete := FALSE;
   TraceIn_estop[21] := BenchUut2.estop;
   TraceIn_opeMode[21] := BenchUut2.opeMode;
   TraceIn_valveAStart[21] := BenchUut2.valveAStart;
   TraceIn_valveBStart[21] := BenchUut2.valveBStart;
   TraceIn_valveCStart[21] := BenchUut2.valveCStart;
   TraceIn_valveDStart[21] := BenchUut2.valveDStart;
   TraceIn_mixMotorStart[21] := BenchUut2.mixMotorStart;
   TraceIn_autoStart[21] := BenchUut2.autoStart;
   TraceIn_processMode[21] := BenchUut2.processMode;
   TraceIn_levelSensor[21] := BenchUut2.levelSensor;
   TraceIn_mixMotorComplete[21] := BenchUut2.mixMotorComplete;
   BenchUut2();
   TraceOut_valveARun[21] := BenchUut2.valveARun;
   TraceOut_valveBRun[21] := BenchUut2.valveBRun;
   TraceOut_valveCRun[21] := BenchUut2.valveCRun;
   TraceOut_valveDRun[21] := BenchUut2.valveDRun;
   TraceOut_mixMotorRun[21] := BenchUut2.mixMotorRun;
   BenchCalls := BenchCalls + 1;
 22:
   BenchUut3.estop := TRUE;
   BenchUut3.opeMode := FALSE;
   BenchUut3.valveAStart := FALSE;
   BenchUut3.valveBStart := TRUE;
   BenchUut3.valveCStart := FALSE;
   BenchUut3.valveDStart := FALSE;
   BenchUut3.mixMotorStart := FALSE;
   BenchUut3.autoStart := FALSE;
   BenchUut3.processMode := FALSE;
   BenchUut3.levelSensor := INT#0;
   BenchUut3.mixMotorComplete := FALSE;
   TraceIn_estop[22] := BenchUut3.estop;
   TraceIn_opeMode[22] := BenchUut3.opeMode;
   TraceIn_valveAStart[22] := BenchUut3.valveAStart;
   TraceIn_valveBStart[22] := BenchUut3.valveBStart;
   TraceIn_valveCStart[22] := BenchUut3.valveCStart;
   TraceIn_valveDStart[22] := BenchUut3.valveDStart;
   TraceIn_mixMotorStart[22] := BenchUut3.mixMotorStart;
   TraceIn_autoStart[22] := BenchUut3.autoStart;
   TraceIn_processMode[22] := BenchUut3.processMode;
   TraceIn_levelSensor[22] := BenchUut3.levelSensor;
   TraceIn_mixMotorComplete[22] := BenchUut3.mixMotorComplete;
   BenchUut3();
   TraceOut_valveARun[22] := BenchUut3.valveARun;
   TraceOut_valveBRun[22] := BenchUut3.valveBRun;
   TraceOut_valveCRun[22] := BenchUut3.valveCRun;
   TraceOut_valveDRun[22] := BenchUut3.valveDRun;
   TraceOut_mixMotorRun[22] := BenchUut3.mixMotorRun;
   BenchCalls := BenchCalls + 1;
 23:
   BenchUut3.estop := TRUE;
   BenchUut3.opeMode := FALSE;
   BenchUut3.valveAStart := FALSE;
   BenchUut3.valveBStart := TRUE;
   BenchUut3.valveCStart := FALSE;
   BenchUut3.valveDStart := FALSE;
   BenchUut3.mixMotorStart := FALSE;
   BenchUut3.autoStart := FALSE;
   BenchUut3.processMode := FALSE;
   BenchUut3.levelSensor := INT#0;
   BenchUut3.mixMotorComplete := FALSE;
   TraceIn_estop[23] := BenchUut3.estop;
   TraceIn_opeMode[23] := BenchUut3.opeMode;
   TraceIn_valveAStart[23] := BenchUut3.valveAStart;
   TraceIn_valveBStart[23] := BenchUut3.valveBStart;
   TraceIn_valveCStart[23] := BenchUut3.valveCStart;
   TraceIn_valveDStart[23] := BenchUut3.valveDStart;
   TraceIn_mixMotorStart[23] := BenchUut3.mixMotorStart;
   TraceIn_autoStart[23] := BenchUut3.autoStart;
   TraceIn_processMode[23] := BenchUut3.processMode;
   TraceIn_levelSensor[23] := BenchUut3.levelSensor;
   TraceIn_mixMotorComplete[23] := BenchUut3.mixMotorComplete;
   BenchUut3();
   TraceOut_valveARun[23] := BenchUut3.valveARun;
   TraceOut_valveBRun[23] := BenchUut3.valveBRun;
   TraceOut_valveCRun[23] := BenchUut3.valveCRun;
   TraceOut_valveDRun[23] := BenchUut3.valveDRun;
   TraceOut_mixMotorRun[23] := BenchUut3.mixMotorRun;
   BenchCalls := BenchCalls + 1;
 24:
   BenchUut3.estop := TRUE;
   BenchUut3.opeMode := TRUE;
   BenchUut3.valveAStart := FALSE;
   BenchUut3.valveBStart := FALSE;
   BenchUut3.valveCStart := FALSE;
   BenchUut3.valveDStart := FALSE;
   BenchUut3.mixMotorStart := FALSE;
   BenchUut3.autoStart := TRUE;
   BenchUut3.processMode := FALSE;
   BenchUut3.levelSensor := INT#0;
   BenchUut3.mixMotorComplete := FALSE;
   TraceIn_estop[24] := BenchUut3.estop;
   TraceIn_opeMode[24] := BenchUut3.opeMode;
   TraceIn_valveAStart[24] := BenchUut3.valveAStart;
   TraceIn_valveBStart[24] := BenchUut3.valveBStart;
   TraceIn_valveCStart[24] := BenchUut3.valveCStart;
   TraceIn_valveDStart[24] := BenchUut3.valveDStart;
   TraceIn_mixMotorStart[24] := BenchUut3.mixMotorStart;
   TraceIn_autoStart[24] := BenchUut3.autoStart;
   TraceIn_processMode[24] := BenchUut3.processMode;
   TraceIn_levelSensor[24] := BenchUut3.levelSensor;
   TraceIn_mixMotorComplete[24] := BenchUut3.mixMotorComplete;
   BenchUut3();
   TraceOut_valveARun[24] := BenchUut3.valveARun;
   TraceOut_valveBRun[24] := BenchUut3.valveBRun;
   TraceOut_valveCRun[24] := BenchUut3.valveCRun;
   TraceOut_valveDRun[24] := BenchUut3.valveDRun;
   TraceOut_mixMotorRun[24] := BenchUut3.mixMotorRun;
   BenchCalls := BenchCalls + 1;
 25:
   BenchUut3.estop := TRUE;
   BenchUut3.opeMode := TRUE;
   BenchUut3.valveAStart := FALSE;
   BenchUut3.valveBStart := FALSE;
   BenchUut3.valveCStart := FALSE;
   BenchUut3.valveDStart := FALSE;
   BenchUut3.mixMotorStart := FALSE;
   BenchUut3.autoStart := TRUE;
   BenchUut3.processMode := FALSE;
   BenchUut3.levelSensor := INT#0;
   BenchUut3.mixMotorComplete := FALSE;
   TraceIn_estop[25] := BenchUut3.estop;
   TraceIn_opeMode[25] := BenchUut3.opeMode;
   TraceIn_valveAStart[25] := BenchUut3.valveAStart;
   TraceIn_valveBStart[25] := BenchUut3.valveBStart;
   TraceIn_valveCStart[25] := BenchUut3.valveCStart;
   TraceIn_valveDStart[25] := BenchUut3.valveDStart;
   TraceIn_mixMotorStart[25] := BenchUut3.mixMotorStart;
   TraceIn_autoStart[25] := BenchUut3.autoStart;
   TraceIn_processMode[25] := BenchUut3.processMode;
   TraceIn_levelSensor[25] := BenchUut3.levelSensor;
   TraceIn_mixMotorComplete[25] := BenchUut3.mixMotorComplete;
   BenchUut3();
   TraceOut_valveARun[25] := BenchUut3.valveARun;
   TraceOut_valveBRun[25] := BenchUut3.valveBRun;
   TraceOut_valveCRun[25] := BenchUut3.valveCRun;
   TraceOut_valveDRun[25] := BenchUut3.valveDRun;
   TraceOut_mixMotorRun[25] := BenchUut3.mixMotorRun;
   BenchCalls := BenchCalls + 1;
 26:
   BenchUut3.estop := TRUE;
   BenchUut3.opeMode := TRUE;
   BenchUut3.valveAStart := FALSE;
   BenchUut3.valveBStart := FALSE;
   BenchUut3.valveCStart := FALSE;
   BenchUut3.valveDStart := FALSE;
   BenchUut3.mixMotorStart := FALSE;
   BenchUut3.autoStart := FALSE;
   BenchUut3.processMode := FALSE;
   BenchUut3.levelSensor := INT#0;
   BenchUut3.mixMotorComplete := FALSE;
   TraceIn_estop[26] := BenchUut3.estop;
   TraceIn_opeMode[26] := BenchUut3.opeMode;
   TraceIn_valveAStart[26] := BenchUut3.valveAStart;
   TraceIn_valveBStart[26] := BenchUut3.valveBStart;
   TraceIn_valveCStart[26] := BenchUut3.valveCStart;
   TraceIn_valveDStart[26] := BenchUut3.valveDStart;
   TraceIn_mixMotorStart[26] := BenchUut3.mixMotorStart;
   TraceIn_autoStart[26] := BenchUut3.autoStart;
   TraceIn_processMode[26] := BenchUut3.processMode;
   TraceIn_levelSensor[26] := BenchUut3.levelSensor;
   TraceIn_mixMotorComplete[26] := BenchUut3.mixMotorComplete;
   BenchUut3();
   TraceOut_valveARun[26] := BenchUut3.valveARun;
   TraceOut_valveBRun[26] := BenchUut3.valveBRun;
   TraceOut_valveCRun[26] := BenchUut3.valveCRun;
   TraceOut_valveDRun[26] := BenchUut3.valveDRun;
   TraceOut_mixMotorRun[26] := BenchUut3.mixMotorRun;
   BenchCalls := BenchCalls + 1;
 27:
   BenchUut3.estop := TRUE;
   BenchUut3.opeMode := TRUE;
   BenchUut3.valveAStart := FALSE;
   BenchUut3.valveBStart := FALSE;
   BenchUut3.valveCStart := FALSE;
   BenchUut3.valveDStart := FALSE;
   BenchUut3.mixMotorStart := FALSE;
   BenchUut3.autoStart := TRUE;
   BenchUut3.processMode := FALSE;
   BenchUut3.levelSensor := INT#0;
   BenchUut3.mixMotorComplete := FALSE;
   TraceIn_estop[27] := BenchUut3.estop;
   TraceIn_opeMode[27] := BenchUut3.opeMode;
   TraceIn_valveAStart[27] := BenchUut3.valveAStart;
   TraceIn_valveBStart[27] := BenchUut3.valveBStart;
   TraceIn_valveCStart[27] := BenchUut3.valveCStart;
   TraceIn_valveDStart[27] := BenchUut3.valveDStart;
   TraceIn_mixMotorStart[27] := BenchUut3.mixMotorStart;
   TraceIn_autoStart[27] := BenchUut3.autoStart;
   TraceIn_processMode[27] := BenchUut3.processMode;
   TraceIn_levelSensor[27] := BenchUut3.levelSensor;
   TraceIn_mixMotorComplete[27] := BenchUut3.mixMotorComplete;
   BenchUut3();
   TraceOut_valveARun[27] := BenchUut3.valveARun;
   TraceOut_valveBRun[27] := BenchUut3.valveBRun;
   TraceOut_valveCRun[27] := BenchUut3.valveCRun;
   TraceOut_valveDRun[27] := BenchUut3.valveDRun;
   TraceOut_mixMotorRun[27] := BenchUut3.mixMotorRun;
   BenchCalls := BenchCalls + 1;
 28:
   BenchUut3.estop := TRUE;
   BenchUut3.opeMode := TRUE;
   BenchUut3.valveAStart := FALSE;
   BenchUut3.valveBStart := FALSE;
   BenchUut3.valveCStart := FALSE;
   BenchUut3.valveDStart := FALSE;
   BenchUut3.mixMotorStart := FALSE;
   BenchUut3.autoStart := FALSE;
   BenchUut3.processMode := FALSE;
   BenchUut3.levelSensor := INT#50;
   BenchUut3.mixMotorComplete := FALSE;
   TraceIn_estop[28] := BenchUut3.estop;
   TraceIn_opeMode[28] := BenchUut3.opeMode;
   TraceIn_valveAStart[28] := BenchUut3.valveAStart;
   TraceIn_valveBStart[28] := BenchUut3.valveBStart;
   TraceIn_valveCStart[28] := BenchUut3.valveCStart;
   TraceIn_valveDStart[28] := BenchUut3.valveDStart;
   TraceIn_mixMotorStart[28] := BenchUut3.mixMotorStart;
   TraceIn_autoStart[28] := BenchUut3.autoStart;
   TraceIn_processMode[28] := BenchUut3.processMode;
   TraceIn_levelSensor[28] := BenchUut3.levelSensor;
   TraceIn_mixMotorComplete[28] := BenchUut3.mixMotorComplete;
   BenchUut3();
   TraceOut_valveARun[28] := BenchUut3.valveARun;
   TraceOut_valveBRun[28] := BenchUut3.valveBRun;
   TraceOut_valveCRun[28] := BenchUut3.valveCRun;
   TraceOut_valveDRun[28] := BenchUut3.valveDRun;
   TraceOut_mixMotorRun[28] := BenchUut3.mixMotorRun;
   BenchCalls := BenchCalls + 1;
 29:
   BenchUut3.estop := TRUE;
   BenchUut3.opeMode := TRUE;
   BenchUut3.valveAStart := FALSE;
   BenchUut3.valveBStart := FALSE;
   BenchUut3.valveCStart := FALSE;
   BenchUut3.valveDStart := FALSE;
   BenchUut3.mixMotorStart := FALSE;
   BenchUut3.autoStart := FALSE;
   BenchUut3.processMode := FALSE;
   BenchUut3.levelSensor := INT#80;
   BenchUut3.mixMotorComplete := FALSE;
   TraceIn_estop[29] := BenchUut3.estop;
   TraceIn_opeMode[29] := BenchUut3.opeMode;
   TraceIn_valveAStart[29] := BenchUut3.valveAStart;
   TraceIn_valveBStart[29] := BenchUut3.valveBStart;
   TraceIn_valveCStart[29] := BenchUut3.valveCStart;
   TraceIn_valveDStart[29] := BenchUut3.valveDStart;
   TraceIn_mixMotorStart[29] := BenchUut3.mixMotorStart;
   TraceIn_autoStart[29] := BenchUut3.autoStart;
   TraceIn_processMode[29] := BenchUut3.processMode;
   TraceIn_levelSensor[29] := BenchUut3.levelSensor;
   TraceIn_mixMotorComplete[29] := BenchUut3.mixMotorComplete;
   BenchUut3();
   TraceOut_valveARun[29] := BenchUut3.valveARun;
   TraceOut_valveBRun[29] := BenchUut3.valveBRun;
   TraceOut_valveCRun[29] := BenchUut3.valveCRun;
   TraceOut_valveDRun[29] := BenchUut3.valveDRun;
   TraceOut_mixMotorRun[29] := BenchUut3.mixMotorRun;
   BenchCalls := BenchCalls + 1;
 30:
   BenchUut3.estop := TRUE;
   BenchUut3.opeMode := TRUE;
   BenchUut3.valveAStart := FALSE;
   BenchUut3.valveBStart := FALSE;
   BenchUut3.valveCStart := FALSE;
   BenchUut3.valveDStart := FALSE;
   BenchUut3.mixMotorStart := FALSE;
   BenchUut3.autoStart := FALSE;
   BenchUut3.processMode := FALSE;
   BenchUut3.levelSensor := INT#0;
   BenchUut3.mixMotorComplete := TRUE;
   TraceIn_estop[30] := BenchUut3.estop;
   TraceIn_opeMode[30] := BenchUut3.opeMode;
   TraceIn_valveAStart[30] := BenchUut3.valveAStart;
   TraceIn_valveBStart[30] := BenchUut3.valveBStart;
   TraceIn_valveCStart[30] := BenchUut3.valveCStart;
   TraceIn_valveDStart[30] := BenchUut3.valveDStart;
   TraceIn_mixMotorStart[30] := BenchUut3.mixMotorStart;
   TraceIn_autoStart[30] := BenchUut3.autoStart;
   TraceIn_processMode[30] := BenchUut3.processMode;
   TraceIn_levelSensor[30] := BenchUut3.levelSensor;
   TraceIn_mixMotorComplete[30] := BenchUut3.mixMotorComplete;
   BenchUut3();
   TraceOut_valveARun[30] := BenchUut3.valveARun;
   TraceOut_valveBRun[30] := BenchUut3.valveBRun;
   TraceOut_valveCRun[30] := BenchUut3.valveCRun;
   TraceOut_valveDRun[30] := BenchUut3.valveDRun;
   TraceOut_mixMotorRun[30] := BenchUut3.mixMotorRun;
   BenchCalls := BenchCalls + 1;
 31:
   BenchUut3.estop := TRUE;
   BenchUut3.opeMode := TRUE;
   BenchUut3.valveAStart := FALSE;
   BenchUut3.valveBStart := FALSE;
   BenchUut3.valveCStart := FALSE;
   BenchUut3.valveDStart := FALSE;
   BenchUut3.mixMotorStart := FALSE;
   BenchUut3.autoStart := FALSE;
   BenchUut3.processMode := FALSE;
   BenchUut3.levelSensor := INT#0;
   BenchUut3.mixMotorComplete := FALSE;
   TraceIn_estop[31] := BenchUut3.estop;
   TraceIn_opeMode[31] := BenchUut3.opeMode;
   TraceIn_valveAStart[31] := BenchUut3.valveAStart;
   TraceIn_valveBStart[31] := BenchUut3.valveBStart;
   TraceIn_valveCStart[31] := BenchUut3.valveCStart;
   TraceIn_valveDStart[31] := BenchUut3.valveDStart;
   TraceIn_mixMotorStart[31] := BenchUut3.mixMotorStart;
   TraceIn_autoStart[31] := BenchUut3.autoStart;
   TraceIn_processMode[31] := BenchUut3.processMode;
   TraceIn_levelSensor[31] := BenchUut3.levelSensor;
   TraceIn_mixMotorComplete[31] := BenchUut3.mixMotorComplete;
   BenchUut3();
   TraceOut_valveARun[31] := BenchUut3.valveARun;
   TraceOut_valveBRun[31] := BenchUut3.valveBRun;
   TraceOut_valveCRun[31] := BenchUut3.valveCRun;
   TraceOut_valveDRun[31] := BenchUut3.valveDRun;
   TraceOut_mixMotorRun[31] := BenchUut3.mixMotorRun;
   BenchCalls := BenchCalls + 1;
 32:
   BenchUut4.estop := TRUE;
   BenchUut4.opeMode := FALSE;
   BenchUut4.valveAStart := FALSE;
   BenchUut4.valveBStart := TRUE;
   BenchUut4.valveCStart := TRUE;
   BenchUut4.valveDStart := FALSE;
   BenchUut4.mixMotorStart := FALSE;
   BenchUut4.autoStart := FALSE;
   BenchUut4.processMode := FALSE;
   BenchUut4.levelSensor := INT#0;
   BenchUut4.mixMotorComplete := FALSE;
   TraceIn_estop[32] := BenchUut4.estop;
   TraceIn_opeMode[32] := BenchUut4.opeMode;
   TraceIn_valveAStart[32] := BenchUut4.valveAStart;
   TraceIn_valveBStart[32] := BenchUut4.valveBStart;
   TraceIn_valveCStart[32] := BenchUut4.valveCStart;
   TraceIn_valveDStart[32] := BenchUut4.valveDStart;
   TraceIn_mixMotorStart[32] := BenchUut4.mixMotorStart;
   TraceIn_autoStart[32] := BenchUut4.autoStart;
   TraceIn_processMode[32] := BenchUut4.processMode;
   TraceIn_levelSensor[32] := BenchUut4.levelSensor;
   TraceIn_mixMotorComplete[32] := BenchUut4.mixMotorComplete;
   BenchUut4();
   TraceOut_valveARun[32] := BenchUut4.valveARun;
   TraceOut_valveBRun[32] := BenchUut4.valveBRun;
   TraceOut_valveCRun[32] := BenchUut4.valveCRun;
   TraceOut_valveDRun[32] := BenchUut4.valveDRun;
   TraceOut_mixMotorRun[32] := BenchUut4.mixMotorRun;
   BenchCalls := BenchCalls + 1;
 33:
   BenchUut4.estop := TRUE;
   BenchUut4.opeMode := FALSE;
   BenchUut4.valveAStart := FALSE;
   BenchUut4.valveBStart := TRUE;
   BenchUut4.valveCStart := FALSE;
   BenchUut4.valveDStart := TRUE;
   BenchUut4.mixMotorStart := FALSE;
   BenchUut4.autoStart := FALSE;
   BenchUut4.processMode := FALSE;
   BenchUut4.levelSensor := INT#0;
   BenchUut4.mixMotorComplete := FALSE;
   TraceIn_estop[33] := BenchUut4.estop;
   TraceIn_opeMode[33] := BenchUut4.opeMode;
   TraceIn_valveAStart[33] := BenchUut4.valveAStart;
   TraceIn_valveBStart[33] := BenchUut4.valveBStart;
   TraceIn_valveCStart[33] := BenchUut4.valveCStart;
   TraceIn_valveDStart[33] := BenchUut4.valveDStart;
   TraceIn_mixMotorStart[33] := BenchUut4.mixMotorStart;
   TraceIn_autoStart[33] := BenchUut4.autoStart;
   TraceIn_processMode[33] := BenchUut4.processMode;
   TraceIn_levelSensor[33] := BenchUut4.levelSensor;
   TraceIn_mixMotorComplete[33] := BenchUut4.mixMotorComplete;
   BenchUut4();
   TraceOut_valveARun[33] := BenchUut4.valveARun;
   TraceOut_valveBRun[33] := BenchUut4.valveBRun;
   TraceOut_valveCRun[33] := BenchUut4.valveCRun;
   TraceOut_valveDRun[33] := BenchUut4.valveDRun;
   TraceOut_mixMotorRun[33] := BenchUut4.mixMotorRun;
   BenchCalls := BenchCalls + 1;
 34:
   BenchUut4.estop := TRUE;
   BenchUut4.opeMode := FALSE;
   BenchUut4.valveAStart := FALSE;
   BenchUut4.valveBStart := FALSE;
   BenchUut4.valveCStart := FALSE;
   BenchUut4.valveDStart := TRUE;
   BenchUut4.mixMotorStart := TRUE;
   BenchUut4.autoStart := FALSE;
   BenchUut4.processMode := FALSE;
   BenchUut4.levelSensor := INT#0;
   BenchUut4.mixMotorComplete := FALSE;
   TraceIn_estop[34] := BenchUut4.estop;
   TraceIn_opeMode[34] := BenchUut4.opeMode;
   TraceIn_valveAStart[34] := BenchUut4.valveAStart;
   TraceIn_valveBStart[34] := BenchUut4.valveBStart;
   TraceIn_valveCStart[34] := BenchUut4.valveCStart;
   TraceIn_valveDStart[34] := BenchUut4.valveDStart;
   TraceIn_mixMotorStart[34] := BenchUut4.mixMotorStart;
   TraceIn_autoStart[34] := BenchUut4.autoStart;
   TraceIn_processMode[34] := BenchUut4.processMode;
   TraceIn_levelSensor[34] := BenchUut4.levelSensor;
   TraceIn_mixMotorComplete[34] := BenchUut4.mixMotorComplete;
   BenchUut4();
   TraceOut_valveARun[34] := BenchUut4.valveARun;
   TraceOut_valveBRun[34] := BenchUut4.valveBRun;
   TraceOut_valveCRun[34] := BenchUut4.valveCRun;
   TraceOut_valveDRun[34] := BenchUut4.valveDRun;
   TraceOut_mixMotorRun[34] := BenchUut4.mixMotorRun;
   BenchCalls := BenchCalls + 1;
 35:
   BenchUut4.estop := TRUE;
   BenchUut4.opeMode := FALSE;
   BenchUut4.valveAStart := FALSE;
   BenchUut4.valveBStart := TRUE;
   BenchUut4.valveCStart := FALSE;
   BenchUut4.valveDStart := FALSE;
   BenchUut4.mixMotorStart := FALSE;
   BenchUut4.autoStart := FALSE;
   BenchUut4.processMode := FALSE;
   BenchUut4.levelSensor := INT#0;
   BenchUut4.mixMotorComplete := FALSE;
   TraceIn_estop[35] := BenchUut4.estop;
   TraceIn_opeMode[35] := BenchUut4.opeMode;
   TraceIn_valveAStart[35] := BenchUut4.valveAStart;
   TraceIn_valveBStart[35] := BenchUut4.valveBStart;
   TraceIn_valveCStart[35] := BenchUut4.valveCStart;
   TraceIn_valveDStart[35] := BenchUut4.valveDStart;
   TraceIn_mixMotorStart[35] := BenchUut4.mixMotorStart;
   TraceIn_autoStart[35] := BenchUut4.autoStart;
   TraceIn_processMode[35] := BenchUut4.processMode;
   TraceIn_levelSensor[35] := BenchUut4.levelSensor;
   TraceIn_mixMotorComplete[35] := BenchUut4.mixMotorComplete;
   BenchUut4();
   TraceOut_valveARun[35] := BenchUut4.valveARun;
   TraceOut_valveBRun[35] := BenchUut4.valveBRun;
   TraceOut_valveCRun[35] := BenchUut4.valveCRun;
   TraceOut_valveDRun[35] := BenchUut4.valveDRun;
   TraceOut_mixMotorRun[35] := BenchUut4.mixMotorRun;
   BenchCalls := BenchCalls + 1;
 36:
   BenchUut4.estop := TRUE;
   BenchUut4.opeMode := TRUE;
   BenchUut4.valveAStart := FALSE;
   BenchUut4.valveBStart := FALSE;
   BenchUut4.valveCStart := FALSE;
   BenchUut4.valveDStart := FALSE;
   BenchUut4.mixMotorStart := FALSE;
   BenchUut4.autoStart := FALSE;
   BenchUut4.processMode := TRUE;
   BenchUut4.levelSensor := INT#0;
   BenchUut4.mixMotorComplete := FALSE;
   TraceIn_estop[36] := BenchUut4.estop;
   TraceIn_opeMode[36] := BenchUut4.opeMode;
   TraceIn_valveAStart[36] := BenchUut4.valveAStart;
   TraceIn_valveBStart[36] := BenchUut4.valveBStart;
   TraceIn_valveCStart[36] := BenchUut4.valveCStart;
   TraceIn_valveDStart[36] := BenchUut4.valveDStart;
   TraceIn_mixMotorStart[36] := BenchUut4.mixMotorStart;
   TraceIn_autoStart[36] := BenchUut4.autoStart;
   TraceIn_processMode[36] := BenchUut4.processMode;
   TraceIn_levelSensor[36] := BenchUut4.levelSensor;
   TraceIn_mixMotorComplete[36] := BenchUut4.mixMotorComplete;
   BenchUut4();
   TraceOut_valveARun[36] := BenchUut4.valveARun;
   TraceOut_valveBRun[36] := BenchUut4.valveBRun;
   TraceOut_valveCRun[36] := BenchUut4.valveCRun;
   TraceOut_valveDRun[36] := BenchUut4.valveDRun;
   TraceOut_mixMotorRun[36] := BenchUut4.mixMotorRun;
   BenchCalls := BenchCalls + 1;
 37:
   BenchUut4.estop := TRUE;
   BenchUut4.opeMode := TRUE;
   BenchUut4.valveAStart := FALSE;
   BenchUut4.valveBStart := FALSE;
   BenchUut4.valveCStart := FALSE;
   BenchUut4.valveDStart := FALSE;
   BenchUut4.mixMotorStart := FALSE;
   BenchUut4.autoStart := TRUE;
   BenchUut4.processMode := TRUE;
   BenchUut4.levelSensor := INT#120;
   BenchUut4.mixMotorComplete := FALSE;
   TraceIn_estop[37] := BenchUut4.estop;
   TraceIn_opeMode[37] := BenchUut4.opeMode;
   TraceIn_valveAStart[37] := BenchUut4.valveAStart;
   TraceIn_valveBStart[37] := BenchUut4.valveBStart;
   TraceIn_valveCStart[37] := BenchUut4.valveCStart;
   TraceIn_valveDStart[37] := BenchUut4.valveDStart;
   TraceIn_mixMotorStart[37] := BenchUut4.mixMotorStart;
   TraceIn_autoStart[37] := BenchUut4.autoStart;
   TraceIn_processMode[37] := BenchUut4.processMode;
   TraceIn_levelSensor[37] := BenchUut4.levelSensor;
   TraceIn_mixMotorComplete[37] := BenchUut4.mixMotorComplete;
   BenchUut4();
   TraceOut_valveARun[37] := BenchUut4.valveARun;
   TraceOut_valveBRun[37] := BenchUut4.valveBRun;
   TraceOut_valveCRun[37] := BenchUut4.valveCRun;
   TraceOut_valveDRun[37] := BenchUut4.valveDRun;
   TraceOut_mixMotorRun[37] := BenchUut4.mixMotorRun;
   BenchCalls := BenchCalls + 1;
 38:
   BenchUut4.estop := TRUE;
   BenchUut4.opeMode := TRUE;
   BenchUut4.valveAStart := FALSE;
   BenchUut4.valveBStart := FALSE;
   BenchUut4.valveCStart := FALSE;
   BenchUut4.valveDStart := FALSE;
   BenchUut4.mixMotorStart := FALSE;
   BenchUut4.autoStart := TRUE;
   BenchUut4.processMode := TRUE;
   BenchUut4.levelSensor := INT#120;
   BenchUut4.mixMotorComplete := FALSE;
   TraceIn_estop[38] := BenchUut4.estop;
   TraceIn_opeMode[38] := BenchUut4.opeMode;
   TraceIn_valveAStart[38] := BenchUut4.valveAStart;
   TraceIn_valveBStart[38] := BenchUut4.valveBStart;
   TraceIn_valveCStart[38] := BenchUut4.valveCStart;
   TraceIn_valveDStart[38] := BenchUut4.valveDStart;
   TraceIn_mixMotorStart[38] := BenchUut4.mixMotorStart;
   TraceIn_autoStart[38] := BenchUut4.autoStart;
   TraceIn_processMode[38] := BenchUut4.processMode;
   TraceIn_levelSensor[38] := BenchUut4.levelSensor;
   TraceIn_mixMotorComplete[38] := BenchUut4.mixMotorComplete;
   BenchUut4();
   TraceOut_valveARun[38] := BenchUut4.valveARun;
   TraceOut_valveBRun[38] := BenchUut4.valveBRun;
   TraceOut_valveCRun[38] := BenchUut4.valveCRun;
   TraceOut_valveDRun[38] := BenchUut4.valveDRun;
   TraceOut_mixMotorRun[38] := BenchUut4.mixMotorRun;
   BenchCalls := BenchCalls + 1;
 39:
   BenchUut4.estop := TRUE;
   BenchUut4.opeMode := TRUE;
   BenchUut4.valveAStart := FALSE;
   BenchUut4.valveBStart := FALSE;
   BenchUut4.valveCStart := FALSE;
   BenchUut4.valveDStart := FALSE;
   BenchUut4.mixMotorStart := FALSE;
   BenchUut4.autoStart := FALSE;
   BenchUut4.processMode := TRUE;
   BenchUut4.levelSensor := INT#120;
   BenchUut4.mixMotorComplete := FALSE;
   TraceIn_estop[39] := BenchUut4.estop;
   TraceIn_opeMode[39] := BenchUut4.opeMode;
   TraceIn_valveAStart[39] := BenchUut4.valveAStart;
   TraceIn_valveBStart[39] := BenchUut4.valveBStart;
   TraceIn_valveCStart[39] := BenchUut4.valveCStart;
   TraceIn_valveDStart[39] := BenchUut4.valveDStart;
   TraceIn_mixMotorStart[39] := BenchUut4.mixMotorStart;
   TraceIn_autoStart[39] := BenchUut4.autoStart;
   TraceIn_processMode[39] := BenchUut4.processMode;
   TraceIn_levelSensor[39] := BenchUut4.levelSensor;
   TraceIn_mixMotorComplete[39] := BenchUut4.mixMotorComplete;
   BenchUut4();
   TraceOut_valveARun[39] := BenchUut4.valveARun;
   TraceOut_valveBRun[39] := BenchUut4.valveBRun;
   TraceOut_valveCRun[39] := BenchUut4.valveCRun;
   TraceOut_valveDRun[39] := BenchUut4.valveDRun;
   TraceOut_mixMotorRun[39] := BenchUut4.mixMotorRun;
   BenchCalls := BenchCalls + 1;
 40:
   BenchUut4.estop := TRUE;
   BenchUut4.opeMode := TRUE;
   BenchUut4.valveAStart := FALSE;
   BenchUut4.valveBStart := FALSE;
   BenchUut4.valveCStart := FALSE;
   BenchUut4.valveDStart := FALSE;
   BenchUut4.mixMotorStart := FALSE;
   BenchUut4.autoStart := FALSE;
   BenchUut4.processMode := TRUE;
   BenchUut4.levelSensor := INT#120;
   BenchUut4.mixMotorComplete := FALSE;
   TraceIn_estop[40] := BenchUut4.estop;
   TraceIn_opeMode[40] := BenchUut4.opeMode;
   TraceIn_valveAStart[40] := BenchUut4.valveAStart;
   TraceIn_valveBStart[40] := BenchUut4.valveBStart;
   TraceIn_valveCStart[40] := BenchUut4.valveCStart;
   TraceIn_valveDStart[40] := BenchUut4.valveDStart;
   TraceIn_mixMotorStart[40] := BenchUut4.mixMotorStart;
   TraceIn_autoStart[40] := BenchUut4.autoStart;
   TraceIn_processMode[40] := BenchUut4.processMode;
   TraceIn_levelSensor[40] := BenchUut4.levelSensor;
   TraceIn_mixMotorComplete[40] := BenchUut4.mixMotorComplete;
   BenchUut4();
   TraceOut_valveARun[40] := BenchUut4.valveARun;
   TraceOut_valveBRun[40] := BenchUut4.valveBRun;
   TraceOut_valveCRun[40] := BenchUut4.valveCRun;
   TraceOut_valveDRun[40] := BenchUut4.valveDRun;
   TraceOut_mixMotorRun[40] := BenchUut4.mixMotorRun;
   BenchCalls := BenchCalls + 1;
 41:
   BenchUut4.estop := TRUE;
   BenchUut4.opeMode := TRUE;
   BenchUut4.valveAStart := FALSE;
   BenchUut4.valveBStart := FALSE;
   BenchUut4.valveCStart := FALSE;
   BenchUut4.valveDStart := FALSE;
   BenchUut4.mixMotorStart := FALSE;
   BenchUut4.autoStart := FALSE;
   BenchUut4.processMode := TRUE;
   BenchUut4.levelSensor := INT#120;
   BenchUut4.mixMotorComplete := TRUE;
   TraceIn_estop[41] := BenchUut4.estop;
   TraceIn_opeMode[41] := BenchUut4.opeMode;
   TraceIn_valveAStart[41] := BenchUut4.valveAStart;
   TraceIn_valveBStart[41] := BenchUut4.valveBStart;
   TraceIn_valveCStart[41] := BenchUut4.valveCStart;
   TraceIn_valveDStart[41] := BenchUut4.valveDStart;
   TraceIn_mixMotorStart[41] := BenchUut4.mixMotorStart;
   TraceIn_autoStart[41] := BenchUut4.autoStart;
   TraceIn_processMode[41] := BenchUut4.processMode;
   TraceIn_levelSensor[41] := BenchUut4.levelSensor;
   TraceIn_mixMotorComplete[41] := BenchUut4.mixMotorComplete;
   BenchUut4();
   TraceOut_valveARun[41] := BenchUut4.valveARun;
   TraceOut_valveBRun[41] := BenchUut4.valveBRun;
   TraceOut_valveCRun[41] := BenchUut4.valveCRun;
   TraceOut_valveDRun[41] := BenchUut4.valveDRun;
   TraceOut_mixMotorRun[41] := BenchUut4.mixMotorRun;
   BenchCalls := BenchCalls + 1;
 42:
   BenchUut4.estop := TRUE;
   BenchUut4.opeMode := TRUE;
   BenchUut4.valveAStart := FALSE;
   BenchUut4.valveBStart := FALSE;
   BenchUut4.valveCStart := FALSE;
   BenchUut4.valveDStart := FALSE;
   BenchUut4.mixMotorStart := FALSE;
   BenchUut4.autoStart := FALSE;
   BenchUut4.processMode := TRUE;
   BenchUut4.levelSensor := INT#0;
   BenchUut4.mixMotorComplete := FALSE;
   TraceIn_estop[42] := BenchUut4.estop;
   TraceIn_opeMode[42] := BenchUut4.opeMode;
   TraceIn_valveAStart[42] := BenchUut4.valveAStart;
   TraceIn_valveBStart[42] := BenchUut4.valveBStart;
   TraceIn_valveCStart[42] := BenchUut4.valveCStart;
   TraceIn_valveDStart[42] := BenchUut4.valveDStart;
   TraceIn_mixMotorStart[42] := BenchUut4.mixMotorStart;
   TraceIn_autoStart[42] := BenchUut4.autoStart;
   TraceIn_processMode[42] := BenchUut4.processMode;
   TraceIn_levelSensor[42] := BenchUut4.levelSensor;
   TraceIn_mixMotorComplete[42] := BenchUut4.mixMotorComplete;
   BenchUut4();
   TraceOut_valveARun[42] := BenchUut4.valveARun;
   TraceOut_valveBRun[42] := BenchUut4.valveBRun;
   TraceOut_valveCRun[42] := BenchUut4.valveCRun;
   TraceOut_valveDRun[42] := BenchUut4.valveDRun;
   TraceOut_mixMotorRun[42] := BenchUut4.mixMotorRun;
   BenchCalls := BenchCalls + 1;
 43:
   BenchUut4.estop := TRUE;
   BenchUut4.opeMode := TRUE;
   BenchUut4.valveAStart := FALSE;
   BenchUut4.valveBStart := FALSE;
   BenchUut4.valveCStart := FALSE;
   BenchUut4.valveDStart := FALSE;
   BenchUut4.mixMotorStart := FALSE;
   BenchUut4.autoStart := TRUE;
   BenchUut4.processMode := FALSE;
   BenchUut4.levelSensor := INT#0;
   BenchUut4.mixMotorComplete := FALSE;
   TraceIn_estop[43] := BenchUut4.estop;
   TraceIn_opeMode[43] := BenchUut4.opeMode;
   TraceIn_valveAStart[43] := BenchUut4.valveAStart;
   TraceIn_valveBStart[43] := BenchUut4.valveBStart;
   TraceIn_valveCStart[43] := BenchUut4.valveCStart;
   TraceIn_valveDStart[43] := BenchUut4.valveDStart;
   TraceIn_mixMotorStart[43] := BenchUut4.mixMotorStart;
   TraceIn_autoStart[43] := BenchUut4.autoStart;
   TraceIn_processMode[43] := BenchUut4.processMode;
   TraceIn_levelSensor[43] := BenchUut4.levelSensor;
   TraceIn_mixMotorComplete[43] := BenchUut4.mixMotorComplete;
   BenchUut4();
   TraceOut_valveARun[43] := BenchUut4.valveARun;
   TraceOut_valveBRun[43] := BenchUut4.valveBRun;
   TraceOut_valveCRun[43] := BenchUut4.valveCRun;
   TraceOut_valveDRun[43] := BenchUut4.valveDRun;
   TraceOut_mixMotorRun[43] := BenchUut4.mixMotorRun;
   BenchCalls := BenchCalls + 1;
 44:
   BenchUut4.estop := FALSE;
   BenchUut4.opeMode := TRUE;
   BenchUut4.valveAStart := FALSE;
   BenchUut4.valveBStart := FALSE;
   BenchUut4.valveCStart := FALSE;
   BenchUut4.valveDStart := FALSE;
   BenchUut4.mixMotorStart := FALSE;
   BenchUut4.autoStart := FALSE;
   BenchUut4.processMode := FALSE;
   BenchUut4.levelSensor := INT#50;
   BenchUut4.mixMotorComplete := FALSE;
   TraceIn_estop[44] := BenchUut4.estop;
   TraceIn_opeMode[44] := BenchUut4.opeMode;
   TraceIn_valveAStart[44] := BenchUut4.valveAStart;
   TraceIn_valveBStart[44] := BenchUut4.valveBStart;
   TraceIn_valveCStart[44] := BenchUut4.valveCStart;
   TraceIn_valveDStart[44] := BenchUut4.valveDStart;
   TraceIn_mixMotorStart[44] := BenchUut4.mixMotorStart;
   TraceIn_autoStart[44] := BenchUut4.autoStart;
   TraceIn_processMode[44] := BenchUut4.processMode;
   TraceIn_levelSensor[44] := BenchUut4.levelSensor;
   TraceIn_mixMotorComplete[44] := BenchUut4.mixMotorComplete;
   BenchUut4();
   TraceOut_valveARun[44] := BenchUut4.valveARun;
   TraceOut_valveBRun[44] := BenchUut4.valveBRun;
   TraceOut_valveCRun[44] := BenchUut4.valveCRun;
   TraceOut_valveDRun[44] := BenchUut4.valveDRun;
   TraceOut_mixMotorRun[44] := BenchUut4.mixMotorRun;
   BenchCalls := BenchCalls + 1;
 45:
   BenchUut4.estop := TRUE;
   BenchUut4.opeMode := TRUE;
   BenchUut4.valveAStart := FALSE;
   BenchUut4.valveBStart := FALSE;
   BenchUut4.valveCStart := FALSE;
   BenchUut4.valveDStart := FALSE;
   BenchUut4.mixMotorStart := FALSE;
   BenchUut4.autoStart := FALSE;
   BenchUut4.processMode := FALSE;
   BenchUut4.levelSensor := INT#0;
   BenchUut4.mixMotorComplete := FALSE;
   TraceIn_estop[45] := BenchUut4.estop;
   TraceIn_opeMode[45] := BenchUut4.opeMode;
   TraceIn_valveAStart[45] := BenchUut4.valveAStart;
   TraceIn_valveBStart[45] := BenchUut4.valveBStart;
   TraceIn_valveCStart[45] := BenchUut4.valveCStart;
   TraceIn_valveDStart[45] := BenchUut4.valveDStart;
   TraceIn_mixMotorStart[45] := BenchUut4.mixMotorStart;
   TraceIn_autoStart[45] := BenchUut4.autoStart;
   TraceIn_processMode[45] := BenchUut4.processMode;
   TraceIn_levelSensor[45] := BenchUut4.levelSensor;
   TraceIn_mixMotorComplete[45] := BenchUut4.mixMotorComplete;
   BenchUut4();
   TraceOut_valveARun[45] := BenchUut4.valveARun;
   TraceOut_valveBRun[45] := BenchUut4.valveBRun;
   TraceOut_valveCRun[45] := BenchUut4.valveCRun;
   TraceOut_valveDRun[45] := BenchUut4.valveDRun;
   TraceOut_mixMotorRun[45] := BenchUut4.mixMotorRun;
   BenchCalls := BenchCalls + 1;
 46:
   BenchUut5.estop := TRUE;
   BenchUut5.opeMode := FALSE;
   BenchUut5.valveAStart := FALSE;
   BenchUut5.valveBStart := FALSE;
   BenchUut5.valveCStart := FALSE;
   BenchUut5.valveDStart := FALSE;
   BenchUut5.mixMotorStart := FALSE;
   BenchUut5.autoStart := FALSE;
   BenchUut5.processMode := FALSE;
   BenchUut5.levelSensor := INT#0;
   BenchUut5.mixMotorComplete := FALSE;
   TraceIn_estop[46] := BenchUut5.estop;
   TraceIn_opeMode[46] := BenchUut5.opeMode;
   TraceIn_valveAStart[46] := BenchUut5.valveAStart;
   TraceIn_valveBStart[46] := BenchUut5.valveBStart;
   TraceIn_valveCStart[46] := BenchUut5.valveCStart;
   TraceIn_valveDStart[46] := BenchUut5.valveDStart;
   TraceIn_mixMotorStart[46] := BenchUut5.mixMotorStart;
   TraceIn_autoStart[46] := BenchUut5.autoStart;
   TraceIn_processMode[46] := BenchUut5.processMode;
   TraceIn_levelSensor[46] := BenchUut5.levelSensor;
   TraceIn_mixMotorComplete[46] := BenchUut5.mixMotorComplete;
   BenchUut5();
   TraceOut_valveARun[46] := BenchUut5.valveARun;
   TraceOut_valveBRun[46] := BenchUut5.valveBRun;
   TraceOut_valveCRun[46] := BenchUut5.valveCRun;
   TraceOut_valveDRun[46] := BenchUut5.valveDRun;
   TraceOut_mixMotorRun[46] := BenchUut5.mixMotorRun;
   BenchCalls := BenchCalls + 1;
 47:
   BenchUut5.estop := TRUE;
   BenchUut5.opeMode := FALSE;
   BenchUut5.valveAStart := TRUE;
   BenchUut5.valveBStart := FALSE;
   BenchUut5.valveCStart := FALSE;
   BenchUut5.valveDStart := FALSE;
   BenchUut5.mixMotorStart := FALSE;
   BenchUut5.autoStart := FALSE;
   BenchUut5.processMode := FALSE;
   BenchUut5.levelSensor := INT#0;
   BenchUut5.mixMotorComplete := FALSE;
   TraceIn_estop[47] := BenchUut5.estop;
   TraceIn_opeMode[47] := BenchUut5.opeMode;
   TraceIn_valveAStart[47] := BenchUut5.valveAStart;
   TraceIn_valveBStart[47] := BenchUut5.valveBStart;
   TraceIn_valveCStart[47] := BenchUut5.valveCStart;
   TraceIn_valveDStart[47] := BenchUut5.valveDStart;
   TraceIn_mixMotorStart[47] := BenchUut5.mixMotorStart;
   TraceIn_autoStart[47] := BenchUut5.autoStart;
   TraceIn_processMode[47] := BenchUut5.processMode;
   TraceIn_levelSensor[47] := BenchUut5.levelSensor;
   TraceIn_mixMotorComplete[47] := BenchUut5.mixMotorComplete;
   BenchUut5();
   TraceOut_valveARun[47] := BenchUut5.valveARun;
   TraceOut_valveBRun[47] := BenchUut5.valveBRun;
   TraceOut_valveCRun[47] := BenchUut5.valveCRun;
   TraceOut_valveDRun[47] := BenchUut5.valveDRun;
   TraceOut_mixMotorRun[47] := BenchUut5.mixMotorRun;
   BenchCalls := BenchCalls + 1;
 48:
   BenchUut5.estop := TRUE;
   BenchUut5.opeMode := FALSE;
   BenchUut5.valveAStart := TRUE;
   BenchUut5.valveBStart := FALSE;
   BenchUut5.valveCStart := FALSE;
   BenchUut5.valveDStart := FALSE;
   BenchUut5.mixMotorStart := FALSE;
   BenchUut5.autoStart := FALSE;
   BenchUut5.processMode := FALSE;
   BenchUut5.levelSensor := INT#0;
   BenchUut5.mixMotorComplete := FALSE;
   TraceIn_estop[48] := BenchUut5.estop;
   TraceIn_opeMode[48] := BenchUut5.opeMode;
   TraceIn_valveAStart[48] := BenchUut5.valveAStart;
   TraceIn_valveBStart[48] := BenchUut5.valveBStart;
   TraceIn_valveCStart[48] := BenchUut5.valveCStart;
   TraceIn_valveDStart[48] := BenchUut5.valveDStart;
   TraceIn_mixMotorStart[48] := BenchUut5.mixMotorStart;
   TraceIn_autoStart[48] := BenchUut5.autoStart;
   TraceIn_processMode[48] := BenchUut5.processMode;
   TraceIn_levelSensor[48] := BenchUut5.levelSensor;
   TraceIn_mixMotorComplete[48] := BenchUut5.mixMotorComplete;
   BenchUut5();
   TraceOut_valveARun[48] := BenchUut5.valveARun;
   TraceOut_valveBRun[48] := BenchUut5.valveBRun;
   TraceOut_valveCRun[48] := BenchUut5.valveCRun;
   TraceOut_valveDRun[48] := BenchUut5.valveDRun;
   TraceOut_mixMotorRun[48] := BenchUut5.mixMotorRun;
   BenchCalls := BenchCalls + 1;
 49:
   BenchUut5.estop := TRUE;
   BenchUut5.opeMode := FALSE;
   BenchUut5.valveAStart := FALSE;
   BenchUut5.valveBStart := FALSE;
   BenchUut5.valveCStart := FALSE;
   BenchUut5.valveDStart := FALSE;
   BenchUut5.mixMotorStart := FALSE;
   BenchUut5.autoStart := FALSE;
   BenchUut5.processMode := FALSE;
   BenchUut5.levelSensor := INT#0;
   BenchUut5.mixMotorComplete := FALSE;
   TraceIn_estop[49] := BenchUut5.estop;
   TraceIn_opeMode[49] := BenchUut5.opeMode;
   TraceIn_valveAStart[49] := BenchUut5.valveAStart;
   TraceIn_valveBStart[49] := BenchUut5.valveBStart;
   TraceIn_valveCStart[49] := BenchUut5.valveCStart;
   TraceIn_valveDStart[49] := BenchUut5.valveDStart;
   TraceIn_mixMotorStart[49] := BenchUut5.mixMotorStart;
   TraceIn_autoStart[49] := BenchUut5.autoStart;
   TraceIn_processMode[49] := BenchUut5.processMode;
   TraceIn_levelSensor[49] := BenchUut5.levelSensor;
   TraceIn_mixMotorComplete[49] := BenchUut5.mixMotorComplete;
   BenchUut5();
   TraceOut_valveARun[49] := BenchUut5.valveARun;
   TraceOut_valveBRun[49] := BenchUut5.valveBRun;
   TraceOut_valveCRun[49] := BenchUut5.valveCRun;
   TraceOut_valveDRun[49] := BenchUut5.valveDRun;
   TraceOut_mixMotorRun[49] := BenchUut5.mixMotorRun;
   BenchCalls := BenchCalls + 1;
 50:
   BenchUut5.estop := TRUE;
   BenchUut5.opeMode := FALSE;
   BenchUut5.valveAStart := TRUE;
   BenchUut5.valveBStart := FALSE;
   BenchUut5.valveCStart := FALSE;
   BenchUut5.valveDStart := FALSE;
   BenchUut5.mixMotorStart := FALSE;
   BenchUut5.autoStart := FALSE;
   BenchUut5.processMode := FALSE;
   BenchUut5.levelSensor := INT#0;
   BenchUut5.mixMotorComplete := FALSE;
   TraceIn_estop[50] := BenchUut5.estop;
   TraceIn_opeMode[50] := BenchUut5.opeMode;
   TraceIn_valveAStart[50] := BenchUut5.valveAStart;
   TraceIn_valveBStart[50] := BenchUut5.valveBStart;
   TraceIn_valveCStart[50] := BenchUut5.valveCStart;
   TraceIn_valveDStart[50] := BenchUut5.valveDStart;
   TraceIn_mixMotorStart[50] := BenchUut5.mixMotorStart;
   TraceIn_autoStart[50] := BenchUut5.autoStart;
   TraceIn_processMode[50] := BenchUut5.processMode;
   TraceIn_levelSensor[50] := BenchUut5.levelSensor;
   TraceIn_mixMotorComplete[50] := BenchUut5.mixMotorComplete;
   BenchUut5();
   TraceOut_valveARun[50] := BenchUut5.valveARun;
   TraceOut_valveBRun[50] := BenchUut5.valveBRun;
   TraceOut_valveCRun[50] := BenchUut5.valveCRun;
   TraceOut_valveDRun[50] := BenchUut5.valveDRun;
   TraceOut_mixMotorRun[50] := BenchUut5.mixMotorRun;
   BenchCalls := BenchCalls + 1;
 51:
   BenchUut5.estop := TRUE;
   BenchUut5.opeMode := FALSE;
   BenchUut5.valveAStart := FALSE;
   BenchUut5.valveBStart := TRUE;
   BenchUut5.valveCStart := TRUE;
   BenchUut5.valveDStart := TRUE;
   BenchUut5.mixMotorStart := TRUE;
   BenchUut5.autoStart := FALSE;
   BenchUut5.processMode := FALSE;
   BenchUut5.levelSensor := INT#0;
   BenchUut5.mixMotorComplete := FALSE;
   TraceIn_estop[51] := BenchUut5.estop;
   TraceIn_opeMode[51] := BenchUut5.opeMode;
   TraceIn_valveAStart[51] := BenchUut5.valveAStart;
   TraceIn_valveBStart[51] := BenchUut5.valveBStart;
   TraceIn_valveCStart[51] := BenchUut5.valveCStart;
   TraceIn_valveDStart[51] := BenchUut5.valveDStart;
   TraceIn_mixMotorStart[51] := BenchUut5.mixMotorStart;
   TraceIn_autoStart[51] := BenchUut5.autoStart;
   TraceIn_processMode[51] := BenchUut5.processMode;
   TraceIn_levelSensor[51] := BenchUut5.levelSensor;
   TraceIn_mixMotorComplete[51] := BenchUut5.mixMotorComplete;
   BenchUut5();
   TraceOut_valveARun[51] := BenchUut5.valveARun;
   TraceOut_valveBRun[51] := BenchUut5.valveBRun;
   TraceOut_valveCRun[51] := BenchUut5.valveCRun;
   TraceOut_valveDRun[51] := BenchUut5.valveDRun;
   TraceOut_mixMotorRun[51] := BenchUut5.mixMotorRun;
   BenchCalls := BenchCalls + 1;
 52:
   BenchUut5.estop := TRUE;
   BenchUut5.opeMode := FALSE;
   BenchUut5.valveAStart := FALSE;
   BenchUut5.valveBStart := TRUE;
   BenchUut5.valveCStart := TRUE;
   BenchUut5.valveDStart := TRUE;
   BenchUut5.mixMotorStart := TRUE;
   BenchUut5.autoStart := FALSE;
   BenchUut5.processMode := FALSE;
   BenchUut5.levelSensor := INT#0;
   BenchUut5.mixMotorComplete := FALSE;
   TraceIn_estop[52] := BenchUut5.estop;
   TraceIn_opeMode[52] := BenchUut5.opeMode;
   TraceIn_valveAStart[52] := BenchUut5.valveAStart;
   TraceIn_valveBStart[52] := BenchUut5.valveBStart;
   TraceIn_valveCStart[52] := BenchUut5.valveCStart;
   TraceIn_valveDStart[52] := BenchUut5.valveDStart;
   TraceIn_mixMotorStart[52] := BenchUut5.mixMotorStart;
   TraceIn_autoStart[52] := BenchUut5.autoStart;
   TraceIn_processMode[52] := BenchUut5.processMode;
   TraceIn_levelSensor[52] := BenchUut5.levelSensor;
   TraceIn_mixMotorComplete[52] := BenchUut5.mixMotorComplete;
   BenchUut5();
   TraceOut_valveARun[52] := BenchUut5.valveARun;
   TraceOut_valveBRun[52] := BenchUut5.valveBRun;
   TraceOut_valveCRun[52] := BenchUut5.valveCRun;
   TraceOut_valveDRun[52] := BenchUut5.valveDRun;
   TraceOut_mixMotorRun[52] := BenchUut5.mixMotorRun;
   BenchCalls := BenchCalls + 1;
 53:
   BenchUut6.estop := TRUE;
   BenchUut6.opeMode := FALSE;
   BenchUut6.valveAStart := FALSE;
   BenchUut6.valveBStart := FALSE;
   BenchUut6.valveCStart := FALSE;
   BenchUut6.valveDStart := FALSE;
   BenchUut6.mixMotorStart := FALSE;
   BenchUut6.autoStart := FALSE;
   BenchUut6.processMode := FALSE;
   BenchUut6.levelSensor := INT#0;
   BenchUut6.mixMotorComplete := FALSE;
   TraceIn_estop[53] := BenchUut6.estop;
   TraceIn_opeMode[53] := BenchUut6.opeMode;
   TraceIn_valveAStart[53] := BenchUut6.valveAStart;
   TraceIn_valveBStart[53] := BenchUut6.valveBStart;
   TraceIn_valveCStart[53] := BenchUut6.valveCStart;
   TraceIn_valveDStart[53] := BenchUut6.valveDStart;
   TraceIn_mixMotorStart[53] := BenchUut6.mixMotorStart;
   TraceIn_autoStart[53] := BenchUut6.autoStart;
   TraceIn_processMode[53] := BenchUut6.processMode;
   TraceIn_levelSensor[53] := BenchUut6.levelSensor;
   TraceIn_mixMotorComplete[53] := BenchUut6.mixMotorComplete;
   BenchUut6();
   TraceOut_valveARun[53] := BenchUut6.valveARun;
   TraceOut_valveBRun[53] := BenchUut6.valveBRun;
   TraceOut_valveCRun[53] := BenchUut6.valveCRun;
   TraceOut_valveDRun[53] := BenchUut6.valveDRun;
   TraceOut_mixMotorRun[53] := BenchUut6.mixMotorRun;
   BenchCalls := BenchCalls + 1;
 54:
   BenchUut6.estop := TRUE;
   BenchUut6.opeMode := FALSE;
   BenchUut6.valveAStart := TRUE;
   BenchUut6.valveBStart := FALSE;
   BenchUut6.valveCStart := FALSE;
   BenchUut6.valveDStart := FALSE;
   BenchUut6.mixMotorStart := FALSE;
   BenchUut6.autoStart := FALSE;
   BenchUut6.processMode := FALSE;
   BenchUut6.levelSensor := INT#0;
   BenchUut6.mixMotorComplete := FALSE;
   TraceIn_estop[54] := BenchUut6.estop;
   TraceIn_opeMode[54] := BenchUut6.opeMode;
   TraceIn_valveAStart[54] := BenchUut6.valveAStart;
   TraceIn_valveBStart[54] := BenchUut6.valveBStart;
   TraceIn_valveCStart[54] := BenchUut6.valveCStart;
   TraceIn_valveDStart[54] := BenchUut6.valveDStart;
   TraceIn_mixMotorStart[54] := BenchUut6.mixMotorStart;
   TraceIn_autoStart[54] := BenchUut6.autoStart;
   TraceIn_processMode[54] := BenchUut6.processMode;
   TraceIn_levelSensor[54] := BenchUut6.levelSensor;
   TraceIn_mixMotorComplete[54] := BenchUut6.mixMotorComplete;
   BenchUut6();
   TraceOut_valveARun[54] := BenchUut6.valveARun;
   TraceOut_valveBRun[54] := BenchUut6.valveBRun;
   TraceOut_valveCRun[54] := BenchUut6.valveCRun;
   TraceOut_valveDRun[54] := BenchUut6.valveDRun;
   TraceOut_mixMotorRun[54] := BenchUut6.mixMotorRun;
   BenchCalls := BenchCalls + 1;
 55:
   BenchUut6.estop := TRUE;
   BenchUut6.opeMode := FALSE;
   BenchUut6.valveAStart := TRUE;
   BenchUut6.valveBStart := FALSE;
   BenchUut6.valveCStart := FALSE;
   BenchUut6.valveDStart := FALSE;
   BenchUut6.mixMotorStart := FALSE;
   BenchUut6.autoStart := FALSE;
   BenchUut6.processMode := FALSE;
   BenchUut6.levelSensor := INT#0;
   BenchUut6.mixMotorComplete := FALSE;
   TraceIn_estop[55] := BenchUut6.estop;
   TraceIn_opeMode[55] := BenchUut6.opeMode;
   TraceIn_valveAStart[55] := BenchUut6.valveAStart;
   TraceIn_valveBStart[55] := BenchUut6.valveBStart;
   TraceIn_valveCStart[55] := BenchUut6.valveCStart;
   TraceIn_valveDStart[55] := BenchUut6.valveDStart;
   TraceIn_mixMotorStart[55] := BenchUut6.mixMotorStart;
   TraceIn_autoStart[55] := BenchUut6.autoStart;
   TraceIn_processMode[55] := BenchUut6.processMode;
   TraceIn_levelSensor[55] := BenchUut6.levelSensor;
   TraceIn_mixMotorComplete[55] := BenchUut6.mixMotorComplete;
   BenchUut6();
   TraceOut_valveARun[55] := BenchUut6.valveARun;
   TraceOut_valveBRun[55] := BenchUut6.valveBRun;
   TraceOut_valveCRun[55] := BenchUut6.valveCRun;
   TraceOut_valveDRun[55] := BenchUut6.valveDRun;
   TraceOut_mixMotorRun[55] := BenchUut6.mixMotorRun;
   BenchCalls := BenchCalls + 1;
 56:
   BenchUut6.estop := TRUE;
   BenchUut6.opeMode := FALSE;
   BenchUut6.valveAStart := FALSE;
   BenchUut6.valveBStart := FALSE;
   BenchUut6.valveCStart := FALSE;
   BenchUut6.valveDStart := FALSE;
   BenchUut6.mixMotorStart := FALSE;
   BenchUut6.autoStart := FALSE;
   BenchUut6.processMode := FALSE;
   BenchUut6.levelSensor := INT#0;
   BenchUut6.mixMotorComplete := FALSE;
   TraceIn_estop[56] := BenchUut6.estop;
   TraceIn_opeMode[56] := BenchUut6.opeMode;
   TraceIn_valveAStart[56] := BenchUut6.valveAStart;
   TraceIn_valveBStart[56] := BenchUut6.valveBStart;
   TraceIn_valveCStart[56] := BenchUut6.valveCStart;
   TraceIn_valveDStart[56] := BenchUut6.valveDStart;
   TraceIn_mixMotorStart[56] := BenchUut6.mixMotorStart;
   TraceIn_autoStart[56] := BenchUut6.autoStart;
   TraceIn_processMode[56] := BenchUut6.processMode;
   TraceIn_levelSensor[56] := BenchUut6.levelSensor;
   TraceIn_mixMotorComplete[56] := BenchUut6.mixMotorComplete;
   BenchUut6();
   TraceOut_valveARun[56] := BenchUut6.valveARun;
   TraceOut_valveBRun[56] := BenchUut6.valveBRun;
   TraceOut_valveCRun[56] := BenchUut6.valveCRun;
   TraceOut_valveDRun[56] := BenchUut6.valveDRun;
   TraceOut_mixMotorRun[56] := BenchUut6.mixMotorRun;
   BenchCalls := BenchCalls + 1;
 57:
   BenchUut6.estop := TRUE;
   BenchUut6.opeMode := FALSE;
   BenchUut6.valveAStart := FALSE;
   BenchUut6.valveBStart := FALSE;
   BenchUut6.valveCStart := FALSE;
   BenchUut6.valveDStart := FALSE;
   BenchUut6.mixMotorStart := FALSE;
   BenchUut6.autoStart := FALSE;
   BenchUut6.processMode := FALSE;
   BenchUut6.levelSensor := INT#0;
   BenchUut6.mixMotorComplete := FALSE;
   TraceIn_estop[57] := BenchUut6.estop;
   TraceIn_opeMode[57] := BenchUut6.opeMode;
   TraceIn_valveAStart[57] := BenchUut6.valveAStart;
   TraceIn_valveBStart[57] := BenchUut6.valveBStart;
   TraceIn_valveCStart[57] := BenchUut6.valveCStart;
   TraceIn_valveDStart[57] := BenchUut6.valveDStart;
   TraceIn_mixMotorStart[57] := BenchUut6.mixMotorStart;
   TraceIn_autoStart[57] := BenchUut6.autoStart;
   TraceIn_processMode[57] := BenchUut6.processMode;
   TraceIn_levelSensor[57] := BenchUut6.levelSensor;
   TraceIn_mixMotorComplete[57] := BenchUut6.mixMotorComplete;
   BenchUut6();
   TraceOut_valveARun[57] := BenchUut6.valveARun;
   TraceOut_valveBRun[57] := BenchUut6.valveBRun;
   TraceOut_valveCRun[57] := BenchUut6.valveCRun;
   TraceOut_valveDRun[57] := BenchUut6.valveDRun;
   TraceOut_mixMotorRun[57] := BenchUut6.mixMotorRun;
   BenchCalls := BenchCalls + 1;
 58:
   BenchUut6.estop := TRUE;
   BenchUut6.opeMode := FALSE;
   BenchUut6.valveAStart := TRUE;
   BenchUut6.valveBStart := FALSE;
   BenchUut6.valveCStart := FALSE;
   BenchUut6.valveDStart := FALSE;
   BenchUut6.mixMotorStart := FALSE;
   BenchUut6.autoStart := FALSE;
   BenchUut6.processMode := FALSE;
   BenchUut6.levelSensor := INT#0;
   BenchUut6.mixMotorComplete := FALSE;
   TraceIn_estop[58] := BenchUut6.estop;
   TraceIn_opeMode[58] := BenchUut6.opeMode;
   TraceIn_valveAStart[58] := BenchUut6.valveAStart;
   TraceIn_valveBStart[58] := BenchUut6.valveBStart;
   TraceIn_valveCStart[58] := BenchUut6.valveCStart;
   TraceIn_valveDStart[58] := BenchUut6.valveDStart;
   TraceIn_mixMotorStart[58] := BenchUut6.mixMotorStart;
   TraceIn_autoStart[58] := BenchUut6.autoStart;
   TraceIn_processMode[58] := BenchUut6.processMode;
   TraceIn_levelSensor[58] := BenchUut6.levelSensor;
   TraceIn_mixMotorComplete[58] := BenchUut6.mixMotorComplete;
   BenchUut6();
   TraceOut_valveARun[58] := BenchUut6.valveARun;
   TraceOut_valveBRun[58] := BenchUut6.valveBRun;
   TraceOut_valveCRun[58] := BenchUut6.valveCRun;
   TraceOut_valveDRun[58] := BenchUut6.valveDRun;
   TraceOut_mixMotorRun[58] := BenchUut6.mixMotorRun;
   BenchCalls := BenchCalls + 1;
 59:
   BenchUut6.estop := TRUE;
   BenchUut6.opeMode := FALSE;
   BenchUut6.valveAStart := TRUE;
   BenchUut6.valveBStart := FALSE;
   BenchUut6.valveCStart := FALSE;
   BenchUut6.valveDStart := FALSE;
   BenchUut6.mixMotorStart := FALSE;
   BenchUut6.autoStart := FALSE;
   BenchUut6.processMode := FALSE;
   BenchUut6.levelSensor := INT#0;
   BenchUut6.mixMotorComplete := FALSE;
   TraceIn_estop[59] := BenchUut6.estop;
   TraceIn_opeMode[59] := BenchUut6.opeMode;
   TraceIn_valveAStart[59] := BenchUut6.valveAStart;
   TraceIn_valveBStart[59] := BenchUut6.valveBStart;
   TraceIn_valveCStart[59] := BenchUut6.valveCStart;
   TraceIn_valveDStart[59] := BenchUut6.valveDStart;
   TraceIn_mixMotorStart[59] := BenchUut6.mixMotorStart;
   TraceIn_autoStart[59] := BenchUut6.autoStart;
   TraceIn_processMode[59] := BenchUut6.processMode;
   TraceIn_levelSensor[59] := BenchUut6.levelSensor;
   TraceIn_mixMotorComplete[59] := BenchUut6.mixMotorComplete;
   BenchUut6();
   TraceOut_valveARun[59] := BenchUut6.valveARun;
   TraceOut_valveBRun[59] := BenchUut6.valveBRun;
   TraceOut_valveCRun[59] := BenchUut6.valveCRun;
   TraceOut_valveDRun[59] := BenchUut6.valveDRun;
   TraceOut_mixMotorRun[59] := BenchUut6.mixMotorRun;
   BenchCalls := BenchCalls + 1;
 60:
   BenchUut6.estop := TRUE;
   BenchUut6.opeMode := FALSE;
   BenchUut6.valveAStart := FALSE;
   BenchUut6.valveBStart := FALSE;
   BenchUut6.valveCStart := FALSE;
   BenchUut6.valveDStart := FALSE;
   BenchUut6.mixMotorStart := FALSE;
   BenchUut6.autoStart := FALSE;
   BenchUut6.processMode := FALSE;
   BenchUut6.levelSensor := INT#0;
   BenchUut6.mixMotorComplete := FALSE;
   TraceIn_estop[60] := BenchUut6.estop;
   TraceIn_opeMode[60] := BenchUut6.opeMode;
   TraceIn_valveAStart[60] := BenchUut6.valveAStart;
   TraceIn_valveBStart[60] := BenchUut6.valveBStart;
   TraceIn_valveCStart[60] := BenchUut6.valveCStart;
   TraceIn_valveDStart[60] := BenchUut6.valveDStart;
   TraceIn_mixMotorStart[60] := BenchUut6.mixMotorStart;
   TraceIn_autoStart[60] := BenchUut6.autoStart;
   TraceIn_processMode[60] := BenchUut6.processMode;
   TraceIn_levelSensor[60] := BenchUut6.levelSensor;
   TraceIn_mixMotorComplete[60] := BenchUut6.mixMotorComplete;
   BenchUut6();
   TraceOut_valveARun[60] := BenchUut6.valveARun;
   TraceOut_valveBRun[60] := BenchUut6.valveBRun;
   TraceOut_valveCRun[60] := BenchUut6.valveCRun;
   TraceOut_valveDRun[60] := BenchUut6.valveDRun;
   TraceOut_mixMotorRun[60] := BenchUut6.mixMotorRun;
   BenchCalls := BenchCalls + 1;
 61:
   BenchUut7.estop := TRUE;
   BenchUut7.opeMode := FALSE;
   BenchUut7.valveAStart := FALSE;
   BenchUut7.valveBStart := FALSE;
   BenchUut7.valveCStart := FALSE;
   BenchUut7.valveDStart := FALSE;
   BenchUut7.mixMotorStart := FALSE;
   BenchUut7.autoStart := FALSE;
   BenchUut7.processMode := FALSE;
   BenchUut7.levelSensor := INT#0;
   BenchUut7.mixMotorComplete := FALSE;
   TraceIn_estop[61] := BenchUut7.estop;
   TraceIn_opeMode[61] := BenchUut7.opeMode;
   TraceIn_valveAStart[61] := BenchUut7.valveAStart;
   TraceIn_valveBStart[61] := BenchUut7.valveBStart;
   TraceIn_valveCStart[61] := BenchUut7.valveCStart;
   TraceIn_valveDStart[61] := BenchUut7.valveDStart;
   TraceIn_mixMotorStart[61] := BenchUut7.mixMotorStart;
   TraceIn_autoStart[61] := BenchUut7.autoStart;
   TraceIn_processMode[61] := BenchUut7.processMode;
   TraceIn_levelSensor[61] := BenchUut7.levelSensor;
   TraceIn_mixMotorComplete[61] := BenchUut7.mixMotorComplete;
   BenchUut7();
   TraceOut_valveARun[61] := BenchUut7.valveARun;
   TraceOut_valveBRun[61] := BenchUut7.valveBRun;
   TraceOut_valveCRun[61] := BenchUut7.valveCRun;
   TraceOut_valveDRun[61] := BenchUut7.valveDRun;
   TraceOut_mixMotorRun[61] := BenchUut7.mixMotorRun;
   BenchCalls := BenchCalls + 1;
 62:
   BenchUut7.estop := TRUE;
   BenchUut7.opeMode := FALSE;
   BenchUut7.valveAStart := FALSE;
   BenchUut7.valveBStart := TRUE;
   BenchUut7.valveCStart := FALSE;
   BenchUut7.valveDStart := FALSE;
   BenchUut7.mixMotorStart := FALSE;
   BenchUut7.autoStart := FALSE;
   BenchUut7.processMode := FALSE;
   BenchUut7.levelSensor := INT#0;
   BenchUut7.mixMotorComplete := FALSE;
   TraceIn_estop[62] := BenchUut7.estop;
   TraceIn_opeMode[62] := BenchUut7.opeMode;
   TraceIn_valveAStart[62] := BenchUut7.valveAStart;
   TraceIn_valveBStart[62] := BenchUut7.valveBStart;
   TraceIn_valveCStart[62] := BenchUut7.valveCStart;
   TraceIn_valveDStart[62] := BenchUut7.valveDStart;
   TraceIn_mixMotorStart[62] := BenchUut7.mixMotorStart;
   TraceIn_autoStart[62] := BenchUut7.autoStart;
   TraceIn_processMode[62] := BenchUut7.processMode;
   TraceIn_levelSensor[62] := BenchUut7.levelSensor;
   TraceIn_mixMotorComplete[62] := BenchUut7.mixMotorComplete;
   BenchUut7();
   TraceOut_valveARun[62] := BenchUut7.valveARun;
   TraceOut_valveBRun[62] := BenchUut7.valveBRun;
   TraceOut_valveCRun[62] := BenchUut7.valveCRun;
   TraceOut_valveDRun[62] := BenchUut7.valveDRun;
   TraceOut_mixMotorRun[62] := BenchUut7.mixMotorRun;
   BenchCalls := BenchCalls + 1;
 63:
   BenchUut7.estop := TRUE;
   BenchUut7.opeMode := FALSE;
   BenchUut7.valveAStart := FALSE;
   BenchUut7.valveBStart := TRUE;
   BenchUut7.valveCStart := FALSE;
   BenchUut7.valveDStart := FALSE;
   BenchUut7.mixMotorStart := FALSE;
   BenchUut7.autoStart := FALSE;
   BenchUut7.processMode := FALSE;
   BenchUut7.levelSensor := INT#0;
   BenchUut7.mixMotorComplete := FALSE;
   TraceIn_estop[63] := BenchUut7.estop;
   TraceIn_opeMode[63] := BenchUut7.opeMode;
   TraceIn_valveAStart[63] := BenchUut7.valveAStart;
   TraceIn_valveBStart[63] := BenchUut7.valveBStart;
   TraceIn_valveCStart[63] := BenchUut7.valveCStart;
   TraceIn_valveDStart[63] := BenchUut7.valveDStart;
   TraceIn_mixMotorStart[63] := BenchUut7.mixMotorStart;
   TraceIn_autoStart[63] := BenchUut7.autoStart;
   TraceIn_processMode[63] := BenchUut7.processMode;
   TraceIn_levelSensor[63] := BenchUut7.levelSensor;
   TraceIn_mixMotorComplete[63] := BenchUut7.mixMotorComplete;
   BenchUut7();
   TraceOut_valveARun[63] := BenchUut7.valveARun;
   TraceOut_valveBRun[63] := BenchUut7.valveBRun;
   TraceOut_valveCRun[63] := BenchUut7.valveCRun;
   TraceOut_valveDRun[63] := BenchUut7.valveDRun;
   TraceOut_mixMotorRun[63] := BenchUut7.mixMotorRun;
   BenchCalls := BenchCalls + 1;
 64:
   BenchUut7.estop := TRUE;
   BenchUut7.opeMode := FALSE;
   BenchUut7.valveAStart := FALSE;
   BenchUut7.valveBStart := FALSE;
   BenchUut7.valveCStart := FALSE;
   BenchUut7.valveDStart := FALSE;
   BenchUut7.mixMotorStart := FALSE;
   BenchUut7.autoStart := FALSE;
   BenchUut7.processMode := FALSE;
   BenchUut7.levelSensor := INT#0;
   BenchUut7.mixMotorComplete := FALSE;
   TraceIn_estop[64] := BenchUut7.estop;
   TraceIn_opeMode[64] := BenchUut7.opeMode;
   TraceIn_valveAStart[64] := BenchUut7.valveAStart;
   TraceIn_valveBStart[64] := BenchUut7.valveBStart;
   TraceIn_valveCStart[64] := BenchUut7.valveCStart;
   TraceIn_valveDStart[64] := BenchUut7.valveDStart;
   TraceIn_mixMotorStart[64] := BenchUut7.mixMotorStart;
   TraceIn_autoStart[64] := BenchUut7.autoStart;
   TraceIn_processMode[64] := BenchUut7.processMode;
   TraceIn_levelSensor[64] := BenchUut7.levelSensor;
   TraceIn_mixMotorComplete[64] := BenchUut7.mixMotorComplete;
   BenchUut7();
   TraceOut_valveARun[64] := BenchUut7.valveARun;
   TraceOut_valveBRun[64] := BenchUut7.valveBRun;
   TraceOut_valveCRun[64] := BenchUut7.valveCRun;
   TraceOut_valveDRun[64] := BenchUut7.valveDRun;
   TraceOut_mixMotorRun[64] := BenchUut7.mixMotorRun;
   BenchCalls := BenchCalls + 1;
 65:
   BenchUut7.estop := TRUE;
   BenchUut7.opeMode := FALSE;
   BenchUut7.valveAStart := FALSE;
   BenchUut7.valveBStart := FALSE;
   BenchUut7.valveCStart := FALSE;
   BenchUut7.valveDStart := FALSE;
   BenchUut7.mixMotorStart := FALSE;
   BenchUut7.autoStart := FALSE;
   BenchUut7.processMode := FALSE;
   BenchUut7.levelSensor := INT#0;
   BenchUut7.mixMotorComplete := FALSE;
   TraceIn_estop[65] := BenchUut7.estop;
   TraceIn_opeMode[65] := BenchUut7.opeMode;
   TraceIn_valveAStart[65] := BenchUut7.valveAStart;
   TraceIn_valveBStart[65] := BenchUut7.valveBStart;
   TraceIn_valveCStart[65] := BenchUut7.valveCStart;
   TraceIn_valveDStart[65] := BenchUut7.valveDStart;
   TraceIn_mixMotorStart[65] := BenchUut7.mixMotorStart;
   TraceIn_autoStart[65] := BenchUut7.autoStart;
   TraceIn_processMode[65] := BenchUut7.processMode;
   TraceIn_levelSensor[65] := BenchUut7.levelSensor;
   TraceIn_mixMotorComplete[65] := BenchUut7.mixMotorComplete;
   BenchUut7();
   TraceOut_valveARun[65] := BenchUut7.valveARun;
   TraceOut_valveBRun[65] := BenchUut7.valveBRun;
   TraceOut_valveCRun[65] := BenchUut7.valveCRun;
   TraceOut_valveDRun[65] := BenchUut7.valveDRun;
   TraceOut_mixMotorRun[65] := BenchUut7.mixMotorRun;
   BenchCalls := BenchCalls + 1;
 66:
   BenchUut7.estop := TRUE;
   BenchUut7.opeMode := FALSE;
   BenchUut7.valveAStart := FALSE;
   BenchUut7.valveBStart := TRUE;
   BenchUut7.valveCStart := FALSE;
   BenchUut7.valveDStart := FALSE;
   BenchUut7.mixMotorStart := FALSE;
   BenchUut7.autoStart := FALSE;
   BenchUut7.processMode := FALSE;
   BenchUut7.levelSensor := INT#0;
   BenchUut7.mixMotorComplete := FALSE;
   TraceIn_estop[66] := BenchUut7.estop;
   TraceIn_opeMode[66] := BenchUut7.opeMode;
   TraceIn_valveAStart[66] := BenchUut7.valveAStart;
   TraceIn_valveBStart[66] := BenchUut7.valveBStart;
   TraceIn_valveCStart[66] := BenchUut7.valveCStart;
   TraceIn_valveDStart[66] := BenchUut7.valveDStart;
   TraceIn_mixMotorStart[66] := BenchUut7.mixMotorStart;
   TraceIn_autoStart[66] := BenchUut7.autoStart;
   TraceIn_processMode[66] := BenchUut7.processMode;
   TraceIn_levelSensor[66] := BenchUut7.levelSensor;
   TraceIn_mixMotorComplete[66] := BenchUut7.mixMotorComplete;
   BenchUut7();
   TraceOut_valveARun[66] := BenchUut7.valveARun;
   TraceOut_valveBRun[66] := BenchUut7.valveBRun;
   TraceOut_valveCRun[66] := BenchUut7.valveCRun;
   TraceOut_valveDRun[66] := BenchUut7.valveDRun;
   TraceOut_mixMotorRun[66] := BenchUut7.mixMotorRun;
   BenchCalls := BenchCalls + 1;
 67:
   BenchUut7.estop := TRUE;
   BenchUut7.opeMode := FALSE;
   BenchUut7.valveAStart := FALSE;
   BenchUut7.valveBStart := TRUE;
   BenchUut7.valveCStart := FALSE;
   BenchUut7.valveDStart := FALSE;
   BenchUut7.mixMotorStart := FALSE;
   BenchUut7.autoStart := FALSE;
   BenchUut7.processMode := FALSE;
   BenchUut7.levelSensor := INT#0;
   BenchUut7.mixMotorComplete := FALSE;
   TraceIn_estop[67] := BenchUut7.estop;
   TraceIn_opeMode[67] := BenchUut7.opeMode;
   TraceIn_valveAStart[67] := BenchUut7.valveAStart;
   TraceIn_valveBStart[67] := BenchUut7.valveBStart;
   TraceIn_valveCStart[67] := BenchUut7.valveCStart;
   TraceIn_valveDStart[67] := BenchUut7.valveDStart;
   TraceIn_mixMotorStart[67] := BenchUut7.mixMotorStart;
   TraceIn_autoStart[67] := BenchUut7.autoStart;
   TraceIn_processMode[67] := BenchUut7.processMode;
   TraceIn_levelSensor[67] := BenchUut7.levelSensor;
   TraceIn_mixMotorComplete[67] := BenchUut7.mixMotorComplete;
   BenchUut7();
   TraceOut_valveARun[67] := BenchUut7.valveARun;
   TraceOut_valveBRun[67] := BenchUut7.valveBRun;
   TraceOut_valveCRun[67] := BenchUut7.valveCRun;
   TraceOut_valveDRun[67] := BenchUut7.valveDRun;
   TraceOut_mixMotorRun[67] := BenchUut7.mixMotorRun;
   BenchCalls := BenchCalls + 1;
 68:
   BenchUut7.estop := TRUE;
   BenchUut7.opeMode := FALSE;
   BenchUut7.valveAStart := FALSE;
   BenchUut7.valveBStart := FALSE;
   BenchUut7.valveCStart := FALSE;
   BenchUut7.valveDStart := FALSE;
   BenchUut7.mixMotorStart := FALSE;
   BenchUut7.autoStart := FALSE;
   BenchUut7.processMode := FALSE;
   BenchUut7.levelSensor := INT#0;
   BenchUut7.mixMotorComplete := FALSE;
   TraceIn_estop[68] := BenchUut7.estop;
   TraceIn_opeMode[68] := BenchUut7.opeMode;
   TraceIn_valveAStart[68] := BenchUut7.valveAStart;
   TraceIn_valveBStart[68] := BenchUut7.valveBStart;
   TraceIn_valveCStart[68] := BenchUut7.valveCStart;
   TraceIn_valveDStart[68] := BenchUut7.valveDStart;
   TraceIn_mixMotorStart[68] := BenchUut7.mixMotorStart;
   TraceIn_autoStart[68] := BenchUut7.autoStart;
   TraceIn_processMode[68] := BenchUut7.processMode;
   TraceIn_levelSensor[68] := BenchUut7.levelSensor;
   TraceIn_mixMotorComplete[68] := BenchUut7.mixMotorComplete;
   BenchUut7();
   TraceOut_valveARun[68] := BenchUut7.valveARun;
   TraceOut_valveBRun[68] := BenchUut7.valveBRun;
   TraceOut_valveCRun[68] := BenchUut7.valveCRun;
   TraceOut_valveDRun[68] := BenchUut7.valveDRun;
   TraceOut_mixMotorRun[68] := BenchUut7.mixMotorRun;
   BenchCalls := BenchCalls + 1;
 69:
   BenchUut8.estop := TRUE;
   BenchUut8.opeMode := FALSE;
   BenchUut8.valveAStart := FALSE;
   BenchUut8.valveBStart := FALSE;
   BenchUut8.valveCStart := FALSE;
   BenchUut8.valveDStart := FALSE;
   BenchUut8.mixMotorStart := FALSE;
   BenchUut8.autoStart := FALSE;
   BenchUut8.processMode := FALSE;
   BenchUut8.levelSensor := INT#0;
   BenchUut8.mixMotorComplete := FALSE;
   TraceIn_estop[69] := BenchUut8.estop;
   TraceIn_opeMode[69] := BenchUut8.opeMode;
   TraceIn_valveAStart[69] := BenchUut8.valveAStart;
   TraceIn_valveBStart[69] := BenchUut8.valveBStart;
   TraceIn_valveCStart[69] := BenchUut8.valveCStart;
   TraceIn_valveDStart[69] := BenchUut8.valveDStart;
   TraceIn_mixMotorStart[69] := BenchUut8.mixMotorStart;
   TraceIn_autoStart[69] := BenchUut8.autoStart;
   TraceIn_processMode[69] := BenchUut8.processMode;
   TraceIn_levelSensor[69] := BenchUut8.levelSensor;
   TraceIn_mixMotorComplete[69] := BenchUut8.mixMotorComplete;
   BenchUut8();
   TraceOut_valveARun[69] := BenchUut8.valveARun;
   TraceOut_valveBRun[69] := BenchUut8.valveBRun;
   TraceOut_valveCRun[69] := BenchUut8.valveCRun;
   TraceOut_valveDRun[69] := BenchUut8.valveDRun;
   TraceOut_mixMotorRun[69] := BenchUut8.mixMotorRun;
   BenchCalls := BenchCalls + 1;
 70:
   BenchUut8.estop := TRUE;
   BenchUut8.opeMode := FALSE;
   BenchUut8.valveAStart := FALSE;
   BenchUut8.valveBStart := FALSE;
   BenchUut8.valveCStart := TRUE;
   BenchUut8.valveDStart := FALSE;
   BenchUut8.mixMotorStart := FALSE;
   BenchUut8.autoStart := FALSE;
   BenchUut8.processMode := FALSE;
   BenchUut8.levelSensor := INT#0;
   BenchUut8.mixMotorComplete := FALSE;
   TraceIn_estop[70] := BenchUut8.estop;
   TraceIn_opeMode[70] := BenchUut8.opeMode;
   TraceIn_valveAStart[70] := BenchUut8.valveAStart;
   TraceIn_valveBStart[70] := BenchUut8.valveBStart;
   TraceIn_valveCStart[70] := BenchUut8.valveCStart;
   TraceIn_valveDStart[70] := BenchUut8.valveDStart;
   TraceIn_mixMotorStart[70] := BenchUut8.mixMotorStart;
   TraceIn_autoStart[70] := BenchUut8.autoStart;
   TraceIn_processMode[70] := BenchUut8.processMode;
   TraceIn_levelSensor[70] := BenchUut8.levelSensor;
   TraceIn_mixMotorComplete[70] := BenchUut8.mixMotorComplete;
   BenchUut8();
   TraceOut_valveARun[70] := BenchUut8.valveARun;
   TraceOut_valveBRun[70] := BenchUut8.valveBRun;
   TraceOut_valveCRun[70] := BenchUut8.valveCRun;
   TraceOut_valveDRun[70] := BenchUut8.valveDRun;
   TraceOut_mixMotorRun[70] := BenchUut8.mixMotorRun;
   BenchCalls := BenchCalls + 1;
 71:
   BenchUut8.estop := TRUE;
   BenchUut8.opeMode := FALSE;
   BenchUut8.valveAStart := FALSE;
   BenchUut8.valveBStart := FALSE;
   BenchUut8.valveCStart := TRUE;
   BenchUut8.valveDStart := FALSE;
   BenchUut8.mixMotorStart := FALSE;
   BenchUut8.autoStart := FALSE;
   BenchUut8.processMode := FALSE;
   BenchUut8.levelSensor := INT#0;
   BenchUut8.mixMotorComplete := FALSE;
   TraceIn_estop[71] := BenchUut8.estop;
   TraceIn_opeMode[71] := BenchUut8.opeMode;
   TraceIn_valveAStart[71] := BenchUut8.valveAStart;
   TraceIn_valveBStart[71] := BenchUut8.valveBStart;
   TraceIn_valveCStart[71] := BenchUut8.valveCStart;
   TraceIn_valveDStart[71] := BenchUut8.valveDStart;
   TraceIn_mixMotorStart[71] := BenchUut8.mixMotorStart;
   TraceIn_autoStart[71] := BenchUut8.autoStart;
   TraceIn_processMode[71] := BenchUut8.processMode;
   TraceIn_levelSensor[71] := BenchUut8.levelSensor;
   TraceIn_mixMotorComplete[71] := BenchUut8.mixMotorComplete;
   BenchUut8();
   TraceOut_valveARun[71] := BenchUut8.valveARun;
   TraceOut_valveBRun[71] := BenchUut8.valveBRun;
   TraceOut_valveCRun[71] := BenchUut8.valveCRun;
   TraceOut_valveDRun[71] := BenchUut8.valveDRun;
   TraceOut_mixMotorRun[71] := BenchUut8.mixMotorRun;
   BenchCalls := BenchCalls + 1;
 72:
   BenchUut8.estop := TRUE;
   BenchUut8.opeMode := FALSE;
   BenchUut8.valveAStart := FALSE;
   BenchUut8.valveBStart := FALSE;
   BenchUut8.valveCStart := FALSE;
   BenchUut8.valveDStart := FALSE;
   BenchUut8.mixMotorStart := FALSE;
   BenchUut8.autoStart := FALSE;
   BenchUut8.processMode := FALSE;
   BenchUut8.levelSensor := INT#0;
   BenchUut8.mixMotorComplete := FALSE;
   TraceIn_estop[72] := BenchUut8.estop;
   TraceIn_opeMode[72] := BenchUut8.opeMode;
   TraceIn_valveAStart[72] := BenchUut8.valveAStart;
   TraceIn_valveBStart[72] := BenchUut8.valveBStart;
   TraceIn_valveCStart[72] := BenchUut8.valveCStart;
   TraceIn_valveDStart[72] := BenchUut8.valveDStart;
   TraceIn_mixMotorStart[72] := BenchUut8.mixMotorStart;
   TraceIn_autoStart[72] := BenchUut8.autoStart;
   TraceIn_processMode[72] := BenchUut8.processMode;
   TraceIn_levelSensor[72] := BenchUut8.levelSensor;
   TraceIn_mixMotorComplete[72] := BenchUut8.mixMotorComplete;
   BenchUut8();
   TraceOut_valveARun[72] := BenchUut8.valveARun;
   TraceOut_valveBRun[72] := BenchUut8.valveBRun;
   TraceOut_valveCRun[72] := BenchUut8.valveCRun;
   TraceOut_valveDRun[72] := BenchUut8.valveDRun;
   TraceOut_mixMotorRun[72] := BenchUut8.mixMotorRun;
   BenchCalls := BenchCalls + 1;
 73:
   BenchUut8.estop := TRUE;
   BenchUut8.opeMode := FALSE;
   BenchUut8.valveAStart := FALSE;
   BenchUut8.valveBStart := FALSE;
   BenchUut8.valveCStart := FALSE;
   BenchUut8.valveDStart := FALSE;
   BenchUut8.mixMotorStart := FALSE;
   BenchUut8.autoStart := FALSE;
   BenchUut8.processMode := FALSE;
   BenchUut8.levelSensor := INT#0;
   BenchUut8.mixMotorComplete := FALSE;
   TraceIn_estop[73] := BenchUut8.estop;
   TraceIn_opeMode[73] := BenchUut8.opeMode;
   TraceIn_valveAStart[73] := BenchUut8.valveAStart;
   TraceIn_valveBStart[73] := BenchUut8.valveBStart;
   TraceIn_valveCStart[73] := BenchUut8.valveCStart;
   TraceIn_valveDStart[73] := BenchUut8.valveDStart;
   TraceIn_mixMotorStart[73] := BenchUut8.mixMotorStart;
   TraceIn_autoStart[73] := BenchUut8.autoStart;
   TraceIn_processMode[73] := BenchUut8.processMode;
   TraceIn_levelSensor[73] := BenchUut8.levelSensor;
   TraceIn_mixMotorComplete[73] := BenchUut8.mixMotorComplete;
   BenchUut8();
   TraceOut_valveARun[73] := BenchUut8.valveARun;
   TraceOut_valveBRun[73] := BenchUut8.valveBRun;
   TraceOut_valveCRun[73] := BenchUut8.valveCRun;
   TraceOut_valveDRun[73] := BenchUut8.valveDRun;
   TraceOut_mixMotorRun[73] := BenchUut8.mixMotorRun;
   BenchCalls := BenchCalls + 1;
 74:
   BenchUut8.estop := TRUE;
   BenchUut8.opeMode := FALSE;
   BenchUut8.valveAStart := FALSE;
   BenchUut8.valveBStart := FALSE;
   BenchUut8.valveCStart := TRUE;
   BenchUut8.valveDStart := FALSE;
   BenchUut8.mixMotorStart := FALSE;
   BenchUut8.autoStart := FALSE;
   BenchUut8.processMode := FALSE;
   BenchUut8.levelSensor := INT#0;
   BenchUut8.mixMotorComplete := FALSE;
   TraceIn_estop[74] := BenchUut8.estop;
   TraceIn_opeMode[74] := BenchUut8.opeMode;
   TraceIn_valveAStart[74] := BenchUut8.valveAStart;
   TraceIn_valveBStart[74] := BenchUut8.valveBStart;
   TraceIn_valveCStart[74] := BenchUut8.valveCStart;
   TraceIn_valveDStart[74] := BenchUut8.valveDStart;
   TraceIn_mixMotorStart[74] := BenchUut8.mixMotorStart;
   TraceIn_autoStart[74] := BenchUut8.autoStart;
   TraceIn_processMode[74] := BenchUut8.processMode;
   TraceIn_levelSensor[74] := BenchUut8.levelSensor;
   TraceIn_mixMotorComplete[74] := BenchUut8.mixMotorComplete;
   BenchUut8();
   TraceOut_valveARun[74] := BenchUut8.valveARun;
   TraceOut_valveBRun[74] := BenchUut8.valveBRun;
   TraceOut_valveCRun[74] := BenchUut8.valveCRun;
   TraceOut_valveDRun[74] := BenchUut8.valveDRun;
   TraceOut_mixMotorRun[74] := BenchUut8.mixMotorRun;
   BenchCalls := BenchCalls + 1;
 75:
   BenchUut8.estop := TRUE;
   BenchUut8.opeMode := FALSE;
   BenchUut8.valveAStart := FALSE;
   BenchUut8.valveBStart := FALSE;
   BenchUut8.valveCStart := TRUE;
   BenchUut8.valveDStart := FALSE;
   BenchUut8.mixMotorStart := FALSE;
   BenchUut8.autoStart := FALSE;
   BenchUut8.processMode := FALSE;
   BenchUut8.levelSensor := INT#0;
   BenchUut8.mixMotorComplete := FALSE;
   TraceIn_estop[75] := BenchUut8.estop;
   TraceIn_opeMode[75] := BenchUut8.opeMode;
   TraceIn_valveAStart[75] := BenchUut8.valveAStart;
   TraceIn_valveBStart[75] := BenchUut8.valveBStart;
   TraceIn_valveCStart[75] := BenchUut8.valveCStart;
   TraceIn_valveDStart[75] := BenchUut8.valveDStart;
   TraceIn_mixMotorStart[75] := BenchUut8.mixMotorStart;
   TraceIn_autoStart[75] := BenchUut8.autoStart;
   TraceIn_processMode[75] := BenchUut8.processMode;
   TraceIn_levelSensor[75] := BenchUut8.levelSensor;
   TraceIn_mixMotorComplete[75] := BenchUut8.mixMotorComplete;
   BenchUut8();
   TraceOut_valveARun[75] := BenchUut8.valveARun;
   TraceOut_valveBRun[75] := BenchUut8.valveBRun;
   TraceOut_valveCRun[75] := BenchUut8.valveCRun;
   TraceOut_valveDRun[75] := BenchUut8.valveDRun;
   TraceOut_mixMotorRun[75] := BenchUut8.mixMotorRun;
   BenchCalls := BenchCalls + 1;
 76:
   BenchUut8.estop := TRUE;
   BenchUut8.opeMode := FALSE;
   BenchUut8.valveAStart := FALSE;
   BenchUut8.valveBStart := FALSE;
   BenchUut8.valveCStart := FALSE;
   BenchUut8.valveDStart := FALSE;
   BenchUut8.mixMotorStart := FALSE;
   BenchUut8.autoStart := FALSE;
   BenchUut8.processMode := FALSE;
   BenchUut8.levelSensor := INT#0;
   BenchUut8.mixMotorComplete := FALSE;
   TraceIn_estop[76] := BenchUut8.estop;
   TraceIn_opeMode[76] := BenchUut8.opeMode;
   TraceIn_valveAStart[76] := BenchUut8.valveAStart;
   TraceIn_valveBStart[76] := BenchUut8.valveBStart;
   TraceIn_valveCStart[76] := BenchUut8.valveCStart;
   TraceIn_valveDStart[76] := BenchUut8.valveDStart;
   TraceIn_mixMotorStart[76] := BenchUut8.mixMotorStart;
   TraceIn_autoStart[76] := BenchUut8.autoStart;
   TraceIn_processMode[76] := BenchUut8.processMode;
   TraceIn_levelSensor[76] := BenchUut8.levelSensor;
   TraceIn_mixMotorComplete[76] := BenchUut8.mixMotorComplete;
   BenchUut8();
   TraceOut_valveARun[76] := BenchUut8.valveARun;
   TraceOut_valveBRun[76] := BenchUut8.valveBRun;
   TraceOut_valveCRun[76] := BenchUut8.valveCRun;
   TraceOut_valveDRun[76] := BenchUut8.valveDRun;
   TraceOut_mixMotorRun[76] := BenchUut8.mixMotorRun;
   BenchCalls := BenchCalls + 1;
 77:
   BenchUut9.estop := TRUE;
   BenchUut9.opeMode := FALSE;
   BenchUut9.valveAStart := FALSE;
   BenchUut9.valveBStart := FALSE;
   BenchUut9.valveCStart := FALSE;
   BenchUut9.valveDStart := FALSE;
   BenchUut9.mixMotorStart := FALSE;
   BenchUut9.autoStart := FALSE;
   BenchUut9.processMode := FALSE;
   BenchUut9.levelSensor := INT#0;
   BenchUut9.mixMotorComplete := FALSE;
   TraceIn_estop[77] := BenchUut9.estop;
   TraceIn_opeMode[77] := BenchUut9.opeMode;
   TraceIn_valveAStart[77] := BenchUut9.valveAStart;
   TraceIn_valveBStart[77] := BenchUut9.valveBStart;
   TraceIn_valveCStart[77] := BenchUut9.valveCStart;
   TraceIn_valveDStart[77] := BenchUut9.valveDStart;
   TraceIn_mixMotorStart[77] := BenchUut9.mixMotorStart;
   TraceIn_autoStart[77] := BenchUut9.autoStart;
   TraceIn_processMode[77] := BenchUut9.processMode;
   TraceIn_levelSensor[77] := BenchUut9.levelSensor;
   TraceIn_mixMotorComplete[77] := BenchUut9.mixMotorComplete;
   BenchUut9();
   TraceOut_valveARun[77] := BenchUut9.valveARun;
   TraceOut_valveBRun[77] := BenchUut9.valveBRun;
   TraceOut_valveCRun[77] := BenchUut9.valveCRun;
   TraceOut_valveDRun[77] := BenchUut9.valveDRun;
   TraceOut_mixMotorRun[77] := BenchUut9.mixMotorRun;
   BenchCalls := BenchCalls + 1;
 78:
   BenchUut9.estop := TRUE;
   BenchUut9.opeMode := FALSE;
   BenchUut9.valveAStart := FALSE;
   BenchUut9.valveBStart := FALSE;
   BenchUut9.valveCStart := FALSE;
   BenchUut9.valveDStart := TRUE;
   BenchUut9.mixMotorStart := FALSE;
   BenchUut9.autoStart := FALSE;
   BenchUut9.processMode := FALSE;
   BenchUut9.levelSensor := INT#0;
   BenchUut9.mixMotorComplete := FALSE;
   TraceIn_estop[78] := BenchUut9.estop;
   TraceIn_opeMode[78] := BenchUut9.opeMode;
   TraceIn_valveAStart[78] := BenchUut9.valveAStart;
   TraceIn_valveBStart[78] := BenchUut9.valveBStart;
   TraceIn_valveCStart[78] := BenchUut9.valveCStart;
   TraceIn_valveDStart[78] := BenchUut9.valveDStart;
   TraceIn_mixMotorStart[78] := BenchUut9.mixMotorStart;
   TraceIn_autoStart[78] := BenchUut9.autoStart;
   TraceIn_processMode[78] := BenchUut9.processMode;
   TraceIn_levelSensor[78] := BenchUut9.levelSensor;
   TraceIn_mixMotorComplete[78] := BenchUut9.mixMotorComplete;
   BenchUut9();
   TraceOut_valveARun[78] := BenchUut9.valveARun;
   TraceOut_valveBRun[78] := BenchUut9.valveBRun;
   TraceOut_valveCRun[78] := BenchUut9.valveCRun;
   TraceOut_valveDRun[78] := BenchUut9.valveDRun;
   TraceOut_mixMotorRun[78] := BenchUut9.mixMotorRun;
   BenchCalls := BenchCalls + 1;
 79:
   BenchUut9.estop := TRUE;
   BenchUut9.opeMode := FALSE;
   BenchUut9.valveAStart := FALSE;
   BenchUut9.valveBStart := FALSE;
   BenchUut9.valveCStart := FALSE;
   BenchUut9.valveDStart := TRUE;
   BenchUut9.mixMotorStart := FALSE;
   BenchUut9.autoStart := FALSE;
   BenchUut9.processMode := FALSE;
   BenchUut9.levelSensor := INT#0;
   BenchUut9.mixMotorComplete := FALSE;
   TraceIn_estop[79] := BenchUut9.estop;
   TraceIn_opeMode[79] := BenchUut9.opeMode;
   TraceIn_valveAStart[79] := BenchUut9.valveAStart;
   TraceIn_valveBStart[79] := BenchUut9.valveBStart;
   TraceIn_valveCStart[79] := BenchUut9.valveCStart;
   TraceIn_valveDStart[79] := BenchUut9.valveDStart;
   TraceIn_mixMotorStart[79] := BenchUut9.mixMotorStart;
   TraceIn_autoStart[79] := BenchUut9.autoStart;
   TraceIn_processMode[79] := BenchUut9.processMode;
   TraceIn_levelSensor[79] := BenchUut9.levelSensor;
   TraceIn_mixMotorComplete[79] := BenchUut9.mixMotorComplete;
   BenchUut9();
   TraceOut_valveARun[79] := BenchUut9.valveARun;
   TraceOut_valveBRun[79] := BenchUut9.valveBRun;
   TraceOut_valveCRun[79] := BenchUut9.valveCRun;
   TraceOut_valveDRun[79] := BenchUut9.valveDRun;
   TraceOut_mixMotorRun[79] := BenchUut9.mixMotorRun;
   BenchCalls := BenchCalls + 1;
 80:
   BenchUut9.estop := TRUE;
   BenchUut9.opeMode := FALSE;
   BenchUut9.valveAStart := FALSE;
   BenchUut9.valveBStart := FALSE;
   BenchUut9.valveCStart := FALSE;
   BenchUut9.valveDStart := FALSE;
   BenchUut9.mixMotorStart := FALSE;
   BenchUut9.autoStart := FALSE;
   BenchUut9.processMode := FALSE;
   BenchUut9.levelSensor := INT#0;
   BenchUut9.mixMotorComplete := FALSE;
   TraceIn_estop[80] := BenchUut9.estop;
   TraceIn_opeMode[80] := BenchUut9.opeMode;
   TraceIn_valveAStart[80] := BenchUut9.valveAStart;
   TraceIn_valveBStart[80] := BenchUut9.valveBStart;
   TraceIn_valveCStart[80] := BenchUut9.valveCStart;
   TraceIn_valveDStart[80] := BenchUut9.valveDStart;
   TraceIn_mixMotorStart[80] := BenchUut9.mixMotorStart;
   TraceIn_autoStart[80] := BenchUut9.autoStart;
   TraceIn_processMode[80] := BenchUut9.processMode;
   TraceIn_levelSensor[80] := BenchUut9.levelSensor;
   TraceIn_mixMotorComplete[80] := BenchUut9.mixMotorComplete;
   BenchUut9();
   TraceOut_valveARun[80] := BenchUut9.valveARun;
   TraceOut_valveBRun[80] := BenchUut9.valveBRun;
   TraceOut_valveCRun[80] := BenchUut9.valveCRun;
   TraceOut_valveDRun[80] := BenchUut9.valveDRun;
   TraceOut_mixMotorRun[80] := BenchUut9.mixMotorRun;
   BenchCalls := BenchCalls + 1;
 81:
   BenchUut9.estop := TRUE;
   BenchUut9.opeMode := FALSE;
   BenchUut9.valveAStart := FALSE;
   BenchUut9.valveBStart := FALSE;
   BenchUut9.valveCStart := FALSE;
   BenchUut9.valveDStart := FALSE;
   BenchUut9.mixMotorStart := FALSE;
   BenchUut9.autoStart := FALSE;
   BenchUut9.processMode := FALSE;
   BenchUut9.levelSensor := INT#0;
   BenchUut9.mixMotorComplete := FALSE;
   TraceIn_estop[81] := BenchUut9.estop;
   TraceIn_opeMode[81] := BenchUut9.opeMode;
   TraceIn_valveAStart[81] := BenchUut9.valveAStart;
   TraceIn_valveBStart[81] := BenchUut9.valveBStart;
   TraceIn_valveCStart[81] := BenchUut9.valveCStart;
   TraceIn_valveDStart[81] := BenchUut9.valveDStart;
   TraceIn_mixMotorStart[81] := BenchUut9.mixMotorStart;
   TraceIn_autoStart[81] := BenchUut9.autoStart;
   TraceIn_processMode[81] := BenchUut9.processMode;
   TraceIn_levelSensor[81] := BenchUut9.levelSensor;
   TraceIn_mixMotorComplete[81] := BenchUut9.mixMotorComplete;
   BenchUut9();
   TraceOut_valveARun[81] := BenchUut9.valveARun;
   TraceOut_valveBRun[81] := BenchUut9.valveBRun;
   TraceOut_valveCRun[81] := BenchUut9.valveCRun;
   TraceOut_valveDRun[81] := BenchUut9.valveDRun;
   TraceOut_mixMotorRun[81] := BenchUut9.mixMotorRun;
   BenchCalls := BenchCalls + 1;
 82:
   BenchUut9.estop := TRUE;
   BenchUut9.opeMode := FALSE;
   BenchUut9.valveAStart := FALSE;
   BenchUut9.valveBStart := FALSE;
   BenchUut9.valveCStart := FALSE;
   BenchUut9.valveDStart := TRUE;
   BenchUut9.mixMotorStart := FALSE;
   BenchUut9.autoStart := FALSE;
   BenchUut9.processMode := FALSE;
   BenchUut9.levelSensor := INT#0;
   BenchUut9.mixMotorComplete := FALSE;
   TraceIn_estop[82] := BenchUut9.estop;
   TraceIn_opeMode[82] := BenchUut9.opeMode;
   TraceIn_valveAStart[82] := BenchUut9.valveAStart;
   TraceIn_valveBStart[82] := BenchUut9.valveBStart;
   TraceIn_valveCStart[82] := BenchUut9.valveCStart;
   TraceIn_valveDStart[82] := BenchUut9.valveDStart;
   TraceIn_mixMotorStart[82] := BenchUut9.mixMotorStart;
   TraceIn_autoStart[82] := BenchUut9.autoStart;
   TraceIn_processMode[82] := BenchUut9.processMode;
   TraceIn_levelSensor[82] := BenchUut9.levelSensor;
   TraceIn_mixMotorComplete[82] := BenchUut9.mixMotorComplete;
   BenchUut9();
   TraceOut_valveARun[82] := BenchUut9.valveARun;
   TraceOut_valveBRun[82] := BenchUut9.valveBRun;
   TraceOut_valveCRun[82] := BenchUut9.valveCRun;
   TraceOut_valveDRun[82] := BenchUut9.valveDRun;
   TraceOut_mixMotorRun[82] := BenchUut9.mixMotorRun;
   BenchCalls := BenchCalls + 1;
 83:
   BenchUut9.estop := TRUE;
   BenchUut9.opeMode := FALSE;
   BenchUut9.valveAStart := FALSE;
   BenchUut9.valveBStart := FALSE;
   BenchUut9.valveCStart := FALSE;
   BenchUut9.valveDStart := TRUE;
   BenchUut9.mixMotorStart := FALSE;
   BenchUut9.autoStart := FALSE;
   BenchUut9.processMode := FALSE;
   BenchUut9.levelSensor := INT#0;
   BenchUut9.mixMotorComplete := FALSE;
   TraceIn_estop[83] := BenchUut9.estop;
   TraceIn_opeMode[83] := BenchUut9.opeMode;
   TraceIn_valveAStart[83] := BenchUut9.valveAStart;
   TraceIn_valveBStart[83] := BenchUut9.valveBStart;
   TraceIn_valveCStart[83] := BenchUut9.valveCStart;
   TraceIn_valveDStart[83] := BenchUut9.valveDStart;
   TraceIn_mixMotorStart[83] := BenchUut9.mixMotorStart;
   TraceIn_autoStart[83] := BenchUut9.autoStart;
   TraceIn_processMode[83] := BenchUut9.processMode;
   TraceIn_levelSensor[83] := BenchUut9.levelSensor;
   TraceIn_mixMotorComplete[83] := BenchUut9.mixMotorComplete;
   BenchUut9();
   TraceOut_valveARun[83] := BenchUut9.valveARun;
   TraceOut_valveBRun[83] := BenchUut9.valveBRun;
   TraceOut_valveCRun[83] := BenchUut9.valveCRun;
   TraceOut_valveDRun[83] := BenchUut9.valveDRun;
   TraceOut_mixMotorRun[83] := BenchUut9.mixMotorRun;
   BenchCalls := BenchCalls + 1;
 84:
   BenchUut9.estop := TRUE;
   BenchUut9.opeMode := FALSE;
   BenchUut9.valveAStart := FALSE;
   BenchUut9.valveBStart := FALSE;
   BenchUut9.valveCStart := FALSE;
   BenchUut9.valveDStart := FALSE;
   BenchUut9.mixMotorStart := FALSE;
   BenchUut9.autoStart := FALSE;
   BenchUut9.processMode := FALSE;
   BenchUut9.levelSensor := INT#0;
   BenchUut9.mixMotorComplete := FALSE;
   TraceIn_estop[84] := BenchUut9.estop;
   TraceIn_opeMode[84] := BenchUut9.opeMode;
   TraceIn_valveAStart[84] := BenchUut9.valveAStart;
   TraceIn_valveBStart[84] := BenchUut9.valveBStart;
   TraceIn_valveCStart[84] := BenchUut9.valveCStart;
   TraceIn_valveDStart[84] := BenchUut9.valveDStart;
   TraceIn_mixMotorStart[84] := BenchUut9.mixMotorStart;
   TraceIn_autoStart[84] := BenchUut9.autoStart;
   TraceIn_processMode[84] := BenchUut9.processMode;
   TraceIn_levelSensor[84] := BenchUut9.levelSensor;
   TraceIn_mixMotorComplete[84] := BenchUut9.mixMotorComplete;
   BenchUut9();
   TraceOut_valveARun[84] := BenchUut9.valveARun;
   TraceOut_valveBRun[84] := BenchUut9.valveBRun;
   TraceOut_valveCRun[84] := BenchUut9.valveCRun;
   TraceOut_valveDRun[84] := BenchUut9.valveDRun;
   TraceOut_mixMotorRun[84] := BenchUut9.mixMotorRun;
   BenchCalls := BenchCalls + 1;
 85:
   BenchUut10.estop := TRUE;
   BenchUut10.opeMode := FALSE;
   BenchUut10.valveAStart := FALSE;
   BenchUut10.valveBStart := FALSE;
   BenchUut10.valveCStart := FALSE;
   BenchUut10.valveDStart := FALSE;
   BenchUut10.mixMotorStart := FALSE;
   BenchUut10.autoStart := FALSE;
   BenchUut10.processMode := FALSE;
   BenchUut10.levelSensor := INT#0;
   BenchUut10.mixMotorComplete := FALSE;
   TraceIn_estop[85] := BenchUut10.estop;
   TraceIn_opeMode[85] := BenchUut10.opeMode;
   TraceIn_valveAStart[85] := BenchUut10.valveAStart;
   TraceIn_valveBStart[85] := BenchUut10.valveBStart;
   TraceIn_valveCStart[85] := BenchUut10.valveCStart;
   TraceIn_valveDStart[85] := BenchUut10.valveDStart;
   TraceIn_mixMotorStart[85] := BenchUut10.mixMotorStart;
   TraceIn_autoStart[85] := BenchUut10.autoStart;
   TraceIn_processMode[85] := BenchUut10.processMode;
   TraceIn_levelSensor[85] := BenchUut10.levelSensor;
   TraceIn_mixMotorComplete[85] := BenchUut10.mixMotorComplete;
   BenchUut10();
   TraceOut_valveARun[85] := BenchUut10.valveARun;
   TraceOut_valveBRun[85] := BenchUut10.valveBRun;
   TraceOut_valveCRun[85] := BenchUut10.valveCRun;
   TraceOut_valveDRun[85] := BenchUut10.valveDRun;
   TraceOut_mixMotorRun[85] := BenchUut10.mixMotorRun;
   BenchCalls := BenchCalls + 1;
 86:
   BenchUut10.estop := TRUE;
   BenchUut10.opeMode := FALSE;
   BenchUut10.valveAStart := FALSE;
   BenchUut10.valveBStart := FALSE;
   BenchUut10.valveCStart := FALSE;
   BenchUut10.valveDStart := FALSE;
   BenchUut10.mixMotorStart := TRUE;
   BenchUut10.autoStart := FALSE;
   BenchUut10.processMode := FALSE;
   BenchUut10.levelSensor := INT#0;
   BenchUut10.mixMotorComplete := FALSE;
   TraceIn_estop[86] := BenchUut10.estop;
   TraceIn_opeMode[86] := BenchUut10.opeMode;
   TraceIn_valveAStart[86] := BenchUut10.valveAStart;
   TraceIn_valveBStart[86] := BenchUut10.valveBStart;
   TraceIn_valveCStart[86] := BenchUut10.valveCStart;
   TraceIn_valveDStart[86] := BenchUut10.valveDStart;
   TraceIn_mixMotorStart[86] := BenchUut10.mixMotorStart;
   TraceIn_autoStart[86] := BenchUut10.autoStart;
   TraceIn_processMode[86] := BenchUut10.processMode;
   TraceIn_levelSensor[86] := BenchUut10.levelSensor;
   TraceIn_mixMotorComplete[86] := BenchUut10.mixMotorComplete;
   BenchUut10();
   TraceOut_valveARun[86] := BenchUut10.valveARun;
   TraceOut_valveBRun[86] := BenchUut10.valveBRun;
   TraceOut_valveCRun[86] := BenchUut10.valveCRun;
   TraceOut_valveDRun[86] := BenchUut10.valveDRun;
   TraceOut_mixMotorRun[86] := BenchUut10.mixMotorRun;
   BenchCalls := BenchCalls + 1;
 87:
   BenchUut10.estop := TRUE;
   BenchUut10.opeMode := FALSE;
   BenchUut10.valveAStart := FALSE;
   BenchUut10.valveBStart := FALSE;
   BenchUut10.valveCStart := FALSE;
   BenchUut10.valveDStart := FALSE;
   BenchUut10.mixMotorStart := TRUE;
   BenchUut10.autoStart := FALSE;
   BenchUut10.processMode := FALSE;
   BenchUut10.levelSensor := INT#0;
   BenchUut10.mixMotorComplete := FALSE;
   TraceIn_estop[87] := BenchUut10.estop;
   TraceIn_opeMode[87] := BenchUut10.opeMode;
   TraceIn_valveAStart[87] := BenchUut10.valveAStart;
   TraceIn_valveBStart[87] := BenchUut10.valveBStart;
   TraceIn_valveCStart[87] := BenchUut10.valveCStart;
   TraceIn_valveDStart[87] := BenchUut10.valveDStart;
   TraceIn_mixMotorStart[87] := BenchUut10.mixMotorStart;
   TraceIn_autoStart[87] := BenchUut10.autoStart;
   TraceIn_processMode[87] := BenchUut10.processMode;
   TraceIn_levelSensor[87] := BenchUut10.levelSensor;
   TraceIn_mixMotorComplete[87] := BenchUut10.mixMotorComplete;
   BenchUut10();
   TraceOut_valveARun[87] := BenchUut10.valveARun;
   TraceOut_valveBRun[87] := BenchUut10.valveBRun;
   TraceOut_valveCRun[87] := BenchUut10.valveCRun;
   TraceOut_valveDRun[87] := BenchUut10.valveDRun;
   TraceOut_mixMotorRun[87] := BenchUut10.mixMotorRun;
   BenchCalls := BenchCalls + 1;
 88:
   BenchUut10.estop := TRUE;
   BenchUut10.opeMode := FALSE;
   BenchUut10.valveAStart := FALSE;
   BenchUut10.valveBStart := FALSE;
   BenchUut10.valveCStart := FALSE;
   BenchUut10.valveDStart := FALSE;
   BenchUut10.mixMotorStart := FALSE;
   BenchUut10.autoStart := FALSE;
   BenchUut10.processMode := FALSE;
   BenchUut10.levelSensor := INT#0;
   BenchUut10.mixMotorComplete := FALSE;
   TraceIn_estop[88] := BenchUut10.estop;
   TraceIn_opeMode[88] := BenchUut10.opeMode;
   TraceIn_valveAStart[88] := BenchUut10.valveAStart;
   TraceIn_valveBStart[88] := BenchUut10.valveBStart;
   TraceIn_valveCStart[88] := BenchUut10.valveCStart;
   TraceIn_valveDStart[88] := BenchUut10.valveDStart;
   TraceIn_mixMotorStart[88] := BenchUut10.mixMotorStart;
   TraceIn_autoStart[88] := BenchUut10.autoStart;
   TraceIn_processMode[88] := BenchUut10.processMode;
   TraceIn_levelSensor[88] := BenchUut10.levelSensor;
   TraceIn_mixMotorComplete[88] := BenchUut10.mixMotorComplete;
   BenchUut10();
   TraceOut_valveARun[88] := BenchUut10.valveARun;
   TraceOut_valveBRun[88] := BenchUut10.valveBRun;
   TraceOut_valveCRun[88] := BenchUut10.valveCRun;
   TraceOut_valveDRun[88] := BenchUut10.valveDRun;
   TraceOut_mixMotorRun[88] := BenchUut10.mixMotorRun;
   BenchCalls := BenchCalls + 1;
 89:
   BenchUut10.estop := TRUE;
   BenchUut10.opeMode := FALSE;
   BenchUut10.valveAStart := FALSE;
   BenchUut10.valveBStart := FALSE;
   BenchUut10.valveCStart := FALSE;
   BenchUut10.valveDStart := FALSE;
   BenchUut10.mixMotorStart := FALSE;
   BenchUut10.autoStart := FALSE;
   BenchUut10.processMode := FALSE;
   BenchUut10.levelSensor := INT#0;
   BenchUut10.mixMotorComplete := FALSE;
   TraceIn_estop[89] := BenchUut10.estop;
   TraceIn_opeMode[89] := BenchUut10.opeMode;
   TraceIn_valveAStart[89] := BenchUut10.valveAStart;
   TraceIn_valveBStart[89] := BenchUut10.valveBStart;
   TraceIn_valveCStart[89] := BenchUut10.valveCStart;
   TraceIn_valveDStart[89] := BenchUut10.valveDStart;
   TraceIn_mixMotorStart[89] := BenchUut10.mixMotorStart;
   TraceIn_autoStart[89] := BenchUut10.autoStart;
   TraceIn_processMode[89] := BenchUut10.processMode;
   TraceIn_levelSensor[89] := BenchUut10.levelSensor;
   TraceIn_mixMotorComplete[89] := BenchUut10.mixMotorComplete;
   BenchUut10();
   TraceOut_valveARun[89] := BenchUut10.valveARun;
   TraceOut_valveBRun[89] := BenchUut10.valveBRun;
   TraceOut_valveCRun[89] := BenchUut10.valveCRun;
   TraceOut_valveDRun[89] := BenchUut10.valveDRun;
   TraceOut_mixMotorRun[89] := BenchUut10.mixMotorRun;
   BenchCalls := BenchCalls + 1;
 90:
   BenchUut10.estop := TRUE;
   BenchUut10.opeMode := FALSE;
   BenchUut10.valveAStart := FALSE;
   BenchUut10.valveBStart := FALSE;
   BenchUut10.valveCStart := FALSE;
   BenchUut10.valveDStart := FALSE;
   BenchUut10.mixMotorStart := TRUE;
   BenchUut10.autoStart := FALSE;
   BenchUut10.processMode := FALSE;
   BenchUut10.levelSensor := INT#0;
   BenchUut10.mixMotorComplete := FALSE;
   TraceIn_estop[90] := BenchUut10.estop;
   TraceIn_opeMode[90] := BenchUut10.opeMode;
   TraceIn_valveAStart[90] := BenchUut10.valveAStart;
   TraceIn_valveBStart[90] := BenchUut10.valveBStart;
   TraceIn_valveCStart[90] := BenchUut10.valveCStart;
   TraceIn_valveDStart[90] := BenchUut10.valveDStart;
   TraceIn_mixMotorStart[90] := BenchUut10.mixMotorStart;
   TraceIn_autoStart[90] := BenchUut10.autoStart;
   TraceIn_processMode[90] := BenchUut10.processMode;
   TraceIn_levelSensor[90] := BenchUut10.levelSensor;
   TraceIn_mixMotorComplete[90] := BenchUut10.mixMotorComplete;
   BenchUut10();
   TraceOut_valveARun[90] := BenchUut10.valveARun;
   TraceOut_valveBRun[90] := BenchUut10.valveBRun;
   TraceOut_valveCRun[90] := BenchUut10.valveCRun;
   TraceOut_valveDRun[90] := BenchUut10.valveDRun;
   TraceOut_mixMotorRun[90] := BenchUut10.mixMotorRun;
   BenchCalls := BenchCalls + 1;
 91:
   BenchUut10.estop := TRUE;
   BenchUut10.opeMode := FALSE;
   BenchUut10.valveAStart := FALSE;
   BenchUut10.valveBStart := FALSE;
   BenchUut10.valveCStart := FALSE;
   BenchUut10.valveDStart := FALSE;
   BenchUut10.mixMotorStart := TRUE;
   BenchUut10.autoStart := FALSE;
   BenchUut10.processMode := FALSE;
   BenchUut10.levelSensor := INT#0;
   BenchUut10.mixMotorComplete := FALSE;
   TraceIn_estop[91] := BenchUut10.estop;
   TraceIn_opeMode[91] := BenchUut10.opeMode;
   TraceIn_valveAStart[91] := BenchUut10.valveAStart;
   TraceIn_valveBStart[91] := BenchUut10.valveBStart;
   TraceIn_valveCStart[91] := BenchUut10.valveCStart;
   TraceIn_valveDStart[91] := BenchUut10.valveDStart;
   TraceIn_mixMotorStart[91] := BenchUut10.mixMotorStart;
   TraceIn_autoStart[91] := BenchUut10.autoStart;
   TraceIn_processMode[91] := BenchUut10.processMode;
   TraceIn_levelSensor[91] := BenchUut10.levelSensor;
   TraceIn_mixMotorComplete[91] := BenchUut10.mixMotorComplete;
   BenchUut10();
   TraceOut_valveARun[91] := BenchUut10.valveARun;
   TraceOut_valveBRun[91] := BenchUut10.valveBRun;
   TraceOut_valveCRun[91] := BenchUut10.valveCRun;
   TraceOut_valveDRun[91] := BenchUut10.valveDRun;
   TraceOut_mixMotorRun[91] := BenchUut10.mixMotorRun;
   BenchCalls := BenchCalls + 1;
 92:
   BenchUut10.estop := TRUE;
   BenchUut10.opeMode := FALSE;
   BenchUut10.valveAStart := FALSE;
   BenchUut10.valveBStart := FALSE;
   BenchUut10.valveCStart := FALSE;
   BenchUut10.valveDStart := FALSE;
   BenchUut10.mixMotorStart := FALSE;
   BenchUut10.autoStart := FALSE;
   BenchUut10.processMode := FALSE;
   BenchUut10.levelSensor := INT#0;
   BenchUut10.mixMotorComplete := FALSE;
   TraceIn_estop[92] := BenchUut10.estop;
   TraceIn_opeMode[92] := BenchUut10.opeMode;
   TraceIn_valveAStart[92] := BenchUut10.valveAStart;
   TraceIn_valveBStart[92] := BenchUut10.valveBStart;
   TraceIn_valveCStart[92] := BenchUut10.valveCStart;
   TraceIn_valveDStart[92] := BenchUut10.valveDStart;
   TraceIn_mixMotorStart[92] := BenchUut10.mixMotorStart;
   TraceIn_autoStart[92] := BenchUut10.autoStart;
   TraceIn_processMode[92] := BenchUut10.processMode;
   TraceIn_levelSensor[92] := BenchUut10.levelSensor;
   TraceIn_mixMotorComplete[92] := BenchUut10.mixMotorComplete;
   BenchUut10();
   TraceOut_valveARun[92] := BenchUut10.valveARun;
   TraceOut_valveBRun[92] := BenchUut10.valveBRun;
   TraceOut_valveCRun[92] := BenchUut10.valveCRun;
   TraceOut_valveDRun[92] := BenchUut10.valveDRun;
   TraceOut_mixMotorRun[92] := BenchUut10.mixMotorRun;
   BenchCalls := BenchCalls + 1;
 93:
   BenchUut11.estop := TRUE;
   BenchUut11.opeMode := TRUE;
   BenchUut11.valveAStart := FALSE;
   BenchUut11.valveBStart := FALSE;
   BenchUut11.valveCStart := FALSE;
   BenchUut11.valveDStart := FALSE;
   BenchUut11.mixMotorStart := FALSE;
   BenchUut11.autoStart := FALSE;
   BenchUut11.processMode := FALSE;
   BenchUut11.levelSensor := INT#0;
   BenchUut11.mixMotorComplete := FALSE;
   TraceIn_estop[93] := BenchUut11.estop;
   TraceIn_opeMode[93] := BenchUut11.opeMode;
   TraceIn_valveAStart[93] := BenchUut11.valveAStart;
   TraceIn_valveBStart[93] := BenchUut11.valveBStart;
   TraceIn_valveCStart[93] := BenchUut11.valveCStart;
   TraceIn_valveDStart[93] := BenchUut11.valveDStart;
   TraceIn_mixMotorStart[93] := BenchUut11.mixMotorStart;
   TraceIn_autoStart[93] := BenchUut11.autoStart;
   TraceIn_processMode[93] := BenchUut11.processMode;
   TraceIn_levelSensor[93] := BenchUut11.levelSensor;
   TraceIn_mixMotorComplete[93] := BenchUut11.mixMotorComplete;
   BenchUut11();
   TraceOut_valveARun[93] := BenchUut11.valveARun;
   TraceOut_valveBRun[93] := BenchUut11.valveBRun;
   TraceOut_valveCRun[93] := BenchUut11.valveCRun;
   TraceOut_valveDRun[93] := BenchUut11.valveDRun;
   TraceOut_mixMotorRun[93] := BenchUut11.mixMotorRun;
   BenchCalls := BenchCalls + 1;
 94:
   BenchUut11.estop := TRUE;
   BenchUut11.opeMode := TRUE;
   BenchUut11.valveAStart := FALSE;
   BenchUut11.valveBStart := FALSE;
   BenchUut11.valveCStart := FALSE;
   BenchUut11.valveDStart := FALSE;
   BenchUut11.mixMotorStart := FALSE;
   BenchUut11.autoStart := TRUE;
   BenchUut11.processMode := FALSE;
   BenchUut11.levelSensor := INT#0;
   BenchUut11.mixMotorComplete := FALSE;
   TraceIn_estop[94] := BenchUut11.estop;
   TraceIn_opeMode[94] := BenchUut11.opeMode;
   TraceIn_valveAStart[94] := BenchUut11.valveAStart;
   TraceIn_valveBStart[94] := BenchUut11.valveBStart;
   TraceIn_valveCStart[94] := BenchUut11.valveCStart;
   TraceIn_valveDStart[94] := BenchUut11.valveDStart;
   TraceIn_mixMotorStart[94] := BenchUut11.mixMotorStart;
   TraceIn_autoStart[94] := BenchUut11.autoStart;
   TraceIn_processMode[94] := BenchUut11.processMode;
   TraceIn_levelSensor[94] := BenchUut11.levelSensor;
   TraceIn_mixMotorComplete[94] := BenchUut11.mixMotorComplete;
   BenchUut11();
   TraceOut_valveARun[94] := BenchUut11.valveARun;
   TraceOut_valveBRun[94] := BenchUut11.valveBRun;
   TraceOut_valveCRun[94] := BenchUut11.valveCRun;
   TraceOut_valveDRun[94] := BenchUut11.valveDRun;
   TraceOut_mixMotorRun[94] := BenchUut11.mixMotorRun;
   BenchCalls := BenchCalls + 1;
 95:
   BenchUut11.estop := TRUE;
   BenchUut11.opeMode := TRUE;
   BenchUut11.valveAStart := FALSE;
   BenchUut11.valveBStart := FALSE;
   BenchUut11.valveCStart := FALSE;
   BenchUut11.valveDStart := FALSE;
   BenchUut11.mixMotorStart := FALSE;
   BenchUut11.autoStart := FALSE;
   BenchUut11.processMode := FALSE;
   BenchUut11.levelSensor := INT#0;
   BenchUut11.mixMotorComplete := FALSE;
   TraceIn_estop[95] := BenchUut11.estop;
   TraceIn_opeMode[95] := BenchUut11.opeMode;
   TraceIn_valveAStart[95] := BenchUut11.valveAStart;
   TraceIn_valveBStart[95] := BenchUut11.valveBStart;
   TraceIn_valveCStart[95] := BenchUut11.valveCStart;
   TraceIn_valveDStart[95] := BenchUut11.valveDStart;
   TraceIn_mixMotorStart[95] := BenchUut11.mixMotorStart;
   TraceIn_autoStart[95] := BenchUut11.autoStart;
   TraceIn_processMode[95] := BenchUut11.processMode;
   TraceIn_levelSensor[95] := BenchUut11.levelSensor;
   TraceIn_mixMotorComplete[95] := BenchUut11.mixMotorComplete;
   BenchUut11();
   TraceOut_valveARun[95] := BenchUut11.valveARun;
   TraceOut_valveBRun[95] := BenchUut11.valveBRun;
   TraceOut_valveCRun[95] := BenchUut11.valveCRun;
   TraceOut_valveDRun[95] := BenchUut11.valveDRun;
   TraceOut_mixMotorRun[95] := BenchUut11.mixMotorRun;
   BenchCalls := BenchCalls + 1;
 96:
   BenchUut11.estop := TRUE;
   BenchUut11.opeMode := TRUE;
   BenchUut11.valveAStart := FALSE;
   BenchUut11.valveBStart := FALSE;
   BenchUut11.valveCStart := FALSE;
   BenchUut11.valveDStart := FALSE;
   BenchUut11.mixMotorStart := FALSE;
   BenchUut11.autoStart := FALSE;
   BenchUut11.processMode := FALSE;
   BenchUut11.levelSensor := INT#0;
   BenchUut11.mixMotorComplete := FALSE;
   TraceIn_estop[96] := BenchUut11.estop;
   TraceIn_opeMode[96] := BenchUut11.opeMode;
   TraceIn_valveAStart[96] := BenchUut11.valveAStart;
   TraceIn_valveBStart[96] := BenchUut11.valveBStart;
   TraceIn_valveCStart[96] := BenchUut11.valveCStart;
   TraceIn_valveDStart[96] := BenchUut11.valveDStart;
   TraceIn_mixMotorStart[96] := BenchUut11.mixMotorStart;
   TraceIn_autoStart[96] := BenchUut11.autoStart;
   TraceIn_processMode[96] := BenchUut11.processMode;
   TraceIn_levelSensor[96] := BenchUut11.levelSensor;
   TraceIn_mixMotorComplete[96] := BenchUut11.mixMotorComplete;
   BenchUut11();
   TraceOut_valveARun[96] := BenchUut11.valveARun;
   TraceOut_valveBRun[96] := BenchUut11.valveBRun;
   TraceOut_valveCRun[96] := BenchUut11.valveCRun;
   TraceOut_valveDRun[96] := BenchUut11.valveDRun;
   TraceOut_mixMotorRun[96] := BenchUut11.mixMotorRun;
   BenchCalls := BenchCalls + 1;
 97:
   BenchUut11.estop := TRUE;
   BenchUut11.opeMode := TRUE;
   BenchUut11.valveAStart := FALSE;
   BenchUut11.valveBStart := FALSE;
   BenchUut11.valveCStart := FALSE;
   BenchUut11.valveDStart := FALSE;
   BenchUut11.mixMotorStart := FALSE;
   BenchUut11.autoStart := FALSE;
   BenchUut11.processMode := FALSE;
   BenchUut11.levelSensor := INT#50;
   BenchUut11.mixMotorComplete := FALSE;
   TraceIn_estop[97] := BenchUut11.estop;
   TraceIn_opeMode[97] := BenchUut11.opeMode;
   TraceIn_valveAStart[97] := BenchUut11.valveAStart;
   TraceIn_valveBStart[97] := BenchUut11.valveBStart;
   TraceIn_valveCStart[97] := BenchUut11.valveCStart;
   TraceIn_valveDStart[97] := BenchUut11.valveDStart;
   TraceIn_mixMotorStart[97] := BenchUut11.mixMotorStart;
   TraceIn_autoStart[97] := BenchUut11.autoStart;
   TraceIn_processMode[97] := BenchUut11.processMode;
   TraceIn_levelSensor[97] := BenchUut11.levelSensor;
   TraceIn_mixMotorComplete[97] := BenchUut11.mixMotorComplete;
   BenchUut11();
   TraceOut_valveARun[97] := BenchUut11.valveARun;
   TraceOut_valveBRun[97] := BenchUut11.valveBRun;
   TraceOut_valveCRun[97] := BenchUut11.valveCRun;
   TraceOut_valveDRun[97] := BenchUut11.valveDRun;
   TraceOut_mixMotorRun[97] := BenchUut11.mixMotorRun;
   BenchCalls := BenchCalls + 1;
 98:
   BenchUut11.estop := TRUE;
   BenchUut11.opeMode := TRUE;
   BenchUut11.valveAStart := FALSE;
   BenchUut11.valveBStart := FALSE;
   BenchUut11.valveCStart := FALSE;
   BenchUut11.valveDStart := FALSE;
   BenchUut11.mixMotorStart := FALSE;
   BenchUut11.autoStart := FALSE;
   BenchUut11.processMode := FALSE;
   BenchUut11.levelSensor := INT#50;
   BenchUut11.mixMotorComplete := FALSE;
   TraceIn_estop[98] := BenchUut11.estop;
   TraceIn_opeMode[98] := BenchUut11.opeMode;
   TraceIn_valveAStart[98] := BenchUut11.valveAStart;
   TraceIn_valveBStart[98] := BenchUut11.valveBStart;
   TraceIn_valveCStart[98] := BenchUut11.valveCStart;
   TraceIn_valveDStart[98] := BenchUut11.valveDStart;
   TraceIn_mixMotorStart[98] := BenchUut11.mixMotorStart;
   TraceIn_autoStart[98] := BenchUut11.autoStart;
   TraceIn_processMode[98] := BenchUut11.processMode;
   TraceIn_levelSensor[98] := BenchUut11.levelSensor;
   TraceIn_mixMotorComplete[98] := BenchUut11.mixMotorComplete;
   BenchUut11();
   TraceOut_valveARun[98] := BenchUut11.valveARun;
   TraceOut_valveBRun[98] := BenchUut11.valveBRun;
   TraceOut_valveCRun[98] := BenchUut11.valveCRun;
   TraceOut_valveDRun[98] := BenchUut11.valveDRun;
   TraceOut_mixMotorRun[98] := BenchUut11.mixMotorRun;
   BenchCalls := BenchCalls + 1;
 99:
   BenchUut11.estop := TRUE;
   BenchUut11.opeMode := TRUE;
   BenchUut11.valveAStart := FALSE;
   BenchUut11.valveBStart := FALSE;
   BenchUut11.valveCStart := FALSE;
   BenchUut11.valveDStart := FALSE;
   BenchUut11.mixMotorStart := FALSE;
   BenchUut11.autoStart := FALSE;
   BenchUut11.processMode := FALSE;
   BenchUut11.levelSensor := INT#80;
   BenchUut11.mixMotorComplete := FALSE;
   TraceIn_estop[99] := BenchUut11.estop;
   TraceIn_opeMode[99] := BenchUut11.opeMode;
   TraceIn_valveAStart[99] := BenchUut11.valveAStart;
   TraceIn_valveBStart[99] := BenchUut11.valveBStart;
   TraceIn_valveCStart[99] := BenchUut11.valveCStart;
   TraceIn_valveDStart[99] := BenchUut11.valveDStart;
   TraceIn_mixMotorStart[99] := BenchUut11.mixMotorStart;
   TraceIn_autoStart[99] := BenchUut11.autoStart;
   TraceIn_processMode[99] := BenchUut11.processMode;
   TraceIn_levelSensor[99] := BenchUut11.levelSensor;
   TraceIn_mixMotorComplete[99] := BenchUut11.mixMotorComplete;
   BenchUut11();
   TraceOut_valveARun[99] := BenchUut11.valveARun;
   TraceOut_valveBRun[99] := BenchUut11.valveBRun;
   TraceOut_valveCRun[99] := BenchUut11.valveCRun;
   TraceOut_valveDRun[99] := BenchUut11.valveDRun;
   TraceOut_mixMotorRun[99] := BenchUut11.mixMotorRun;
   BenchCalls := BenchCalls + 1;
 100:
   BenchUut11.estop := TRUE;
   BenchUut11.opeMode := TRUE;
   BenchUut11.valveAStart := FALSE;
   BenchUut11.valveBStart := FALSE;
   BenchUut11.valveCStart := FALSE;
   BenchUut11.valveDStart := FALSE;
   BenchUut11.mixMotorStart := FALSE;
   BenchUut11.autoStart := FALSE;
   BenchUut11.processMode := FALSE;
   BenchUut11.levelSensor := INT#80;
   BenchUut11.mixMotorComplete := FALSE;
   TraceIn_estop[100] := BenchUut11.estop;
   TraceIn_opeMode[100] := BenchUut11.opeMode;
   TraceIn_valveAStart[100] := BenchUut11.valveAStart;
   TraceIn_valveBStart[100] := BenchUut11.valveBStart;
   TraceIn_valveCStart[100] := BenchUut11.valveCStart;
   TraceIn_valveDStart[100] := BenchUut11.valveDStart;
   TraceIn_mixMotorStart[100] := BenchUut11.mixMotorStart;
   TraceIn_autoStart[100] := BenchUut11.autoStart;
   TraceIn_processMode[100] := BenchUut11.processMode;
   TraceIn_levelSensor[100] := BenchUut11.levelSensor;
   TraceIn_mixMotorComplete[100] := BenchUut11.mixMotorComplete;
   BenchUut11();
   TraceOut_valveARun[100] := BenchUut11.valveARun;
   TraceOut_valveBRun[100] := BenchUut11.valveBRun;
   TraceOut_valveCRun[100] := BenchUut11.valveCRun;
   TraceOut_valveDRun[100] := BenchUut11.valveDRun;
   TraceOut_mixMotorRun[100] := BenchUut11.mixMotorRun;
   BenchCalls := BenchCalls + 1;
 101:
   BenchUut11.estop := TRUE;
   BenchUut11.opeMode := TRUE;
   BenchUut11.valveAStart := FALSE;
   BenchUut11.valveBStart := FALSE;
   BenchUut11.valveCStart := FALSE;
   BenchUut11.valveDStart := FALSE;
   BenchUut11.mixMotorStart := FALSE;
   BenchUut11.autoStart := FALSE;
   BenchUut11.processMode := FALSE;
   BenchUut11.levelSensor := INT#80;
   BenchUut11.mixMotorComplete := FALSE;
   TraceIn_estop[101] := BenchUut11.estop;
   TraceIn_opeMode[101] := BenchUut11.opeMode;
   TraceIn_valveAStart[101] := BenchUut11.valveAStart;
   TraceIn_valveBStart[101] := BenchUut11.valveBStart;
   TraceIn_valveCStart[101] := BenchUut11.valveCStart;
   TraceIn_valveDStart[101] := BenchUut11.valveDStart;
   TraceIn_mixMotorStart[101] := BenchUut11.mixMotorStart;
   TraceIn_autoStart[101] := BenchUut11.autoStart;
   TraceIn_processMode[101] := BenchUut11.processMode;
   TraceIn_levelSensor[101] := BenchUut11.levelSensor;
   TraceIn_mixMotorComplete[101] := BenchUut11.mixMotorComplete;
   BenchUut11();
   TraceOut_valveARun[101] := BenchUut11.valveARun;
   TraceOut_valveBRun[101] := BenchUut11.valveBRun;
   TraceOut_valveCRun[101] := BenchUut11.valveCRun;
   TraceOut_valveDRun[101] := BenchUut11.valveDRun;
   TraceOut_mixMotorRun[101] := BenchUut11.mixMotorRun;
   BenchCalls := BenchCalls + 1;
 102:
   BenchUut11.estop := TRUE;
   BenchUut11.opeMode := TRUE;
   BenchUut11.valveAStart := FALSE;
   BenchUut11.valveBStart := FALSE;
   BenchUut11.valveCStart := FALSE;
   BenchUut11.valveDStart := FALSE;
   BenchUut11.mixMotorStart := FALSE;
   BenchUut11.autoStart := FALSE;
   BenchUut11.processMode := FALSE;
   BenchUut11.levelSensor := INT#80;
   BenchUut11.mixMotorComplete := TRUE;
   TraceIn_estop[102] := BenchUut11.estop;
   TraceIn_opeMode[102] := BenchUut11.opeMode;
   TraceIn_valveAStart[102] := BenchUut11.valveAStart;
   TraceIn_valveBStart[102] := BenchUut11.valveBStart;
   TraceIn_valveCStart[102] := BenchUut11.valveCStart;
   TraceIn_valveDStart[102] := BenchUut11.valveDStart;
   TraceIn_mixMotorStart[102] := BenchUut11.mixMotorStart;
   TraceIn_autoStart[102] := BenchUut11.autoStart;
   TraceIn_processMode[102] := BenchUut11.processMode;
   TraceIn_levelSensor[102] := BenchUut11.levelSensor;
   TraceIn_mixMotorComplete[102] := BenchUut11.mixMotorComplete;
   BenchUut11();
   TraceOut_valveARun[102] := BenchUut11.valveARun;
   TraceOut_valveBRun[102] := BenchUut11.valveBRun;
   TraceOut_valveCRun[102] := BenchUut11.valveCRun;
   TraceOut_valveDRun[102] := BenchUut11.valveDRun;
   TraceOut_mixMotorRun[102] := BenchUut11.mixMotorRun;
   BenchCalls := BenchCalls + 1;
 103:
   BenchUut11.estop := TRUE;
   BenchUut11.opeMode := TRUE;
   BenchUut11.valveAStart := FALSE;
   BenchUut11.valveBStart := FALSE;
   BenchUut11.valveCStart := FALSE;
   BenchUut11.valveDStart := FALSE;
   BenchUut11.mixMotorStart := FALSE;
   BenchUut11.autoStart := FALSE;
   BenchUut11.processMode := FALSE;
   BenchUut11.levelSensor := INT#80;
   BenchUut11.mixMotorComplete := FALSE;
   TraceIn_estop[103] := BenchUut11.estop;
   TraceIn_opeMode[103] := BenchUut11.opeMode;
   TraceIn_valveAStart[103] := BenchUut11.valveAStart;
   TraceIn_valveBStart[103] := BenchUut11.valveBStart;
   TraceIn_valveCStart[103] := BenchUut11.valveCStart;
   TraceIn_valveDStart[103] := BenchUut11.valveDStart;
   TraceIn_mixMotorStart[103] := BenchUut11.mixMotorStart;
   TraceIn_autoStart[103] := BenchUut11.autoStart;
   TraceIn_processMode[103] := BenchUut11.processMode;
   TraceIn_levelSensor[103] := BenchUut11.levelSensor;
   TraceIn_mixMotorComplete[103] := BenchUut11.mixMotorComplete;
   BenchUut11();
   TraceOut_valveARun[103] := BenchUut11.valveARun;
   TraceOut_valveBRun[103] := BenchUut11.valveBRun;
   TraceOut_valveCRun[103] := BenchUut11.valveCRun;
   TraceOut_valveDRun[103] := BenchUut11.valveDRun;
   TraceOut_mixMotorRun[103] := BenchUut11.mixMotorRun;
   BenchCalls := BenchCalls + 1;
 104:
   BenchUut11.estop := TRUE;
   BenchUut11.opeMode := TRUE;
   BenchUut11.valveAStart := FALSE;
   BenchUut11.valveBStart := FALSE;
   BenchUut11.valveCStart := FALSE;
   BenchUut11.valveDStart := FALSE;
   BenchUut11.mixMotorStart := FALSE;
   BenchUut11.autoStart := FALSE;
   BenchUut11.processMode := FALSE;
   BenchUut11.levelSensor := INT#80;
   BenchUut11.mixMotorComplete := FALSE;
   TraceIn_estop[104] := BenchUut11.estop;
   TraceIn_opeMode[104] := BenchUut11.opeMode;
   TraceIn_valveAStart[104] := BenchUut11.valveAStart;
   TraceIn_valveBStart[104] := BenchUut11.valveBStart;
   TraceIn_valveCStart[104] := BenchUut11.valveCStart;
   TraceIn_valveDStart[104] := BenchUut11.valveDStart;
   TraceIn_mixMotorStart[104] := BenchUut11.mixMotorStart;
   TraceIn_autoStart[104] := BenchUut11.autoStart;
   TraceIn_processMode[104] := BenchUut11.processMode;
   TraceIn_levelSensor[104] := BenchUut11.levelSensor;
   TraceIn_mixMotorComplete[104] := BenchUut11.mixMotorComplete;
   BenchUut11();
   TraceOut_valveARun[104] := BenchUut11.valveARun;
   TraceOut_valveBRun[104] := BenchUut11.valveBRun;
   TraceOut_valveCRun[104] := BenchUut11.valveCRun;
   TraceOut_valveDRun[104] := BenchUut11.valveDRun;
   TraceOut_mixMotorRun[104] := BenchUut11.mixMotorRun;
   BenchCalls := BenchCalls + 1;
 105:
   BenchUut11.estop := TRUE;
   BenchUut11.opeMode := FALSE;
   BenchUut11.valveAStart := FALSE;
   BenchUut11.valveBStart := FALSE;
   BenchUut11.valveCStart := FALSE;
   BenchUut11.valveDStart := FALSE;
   BenchUut11.mixMotorStart := FALSE;
   BenchUut11.autoStart := FALSE;
   BenchUut11.processMode := FALSE;
   BenchUut11.levelSensor := INT#80;
   BenchUut11.mixMotorComplete := FALSE;
   TraceIn_estop[105] := BenchUut11.estop;
   TraceIn_opeMode[105] := BenchUut11.opeMode;
   TraceIn_valveAStart[105] := BenchUut11.valveAStart;
   TraceIn_valveBStart[105] := BenchUut11.valveBStart;
   TraceIn_valveCStart[105] := BenchUut11.valveCStart;
   TraceIn_valveDStart[105] := BenchUut11.valveDStart;
   TraceIn_mixMotorStart[105] := BenchUut11.mixMotorStart;
   TraceIn_autoStart[105] := BenchUut11.autoStart;
   TraceIn_processMode[105] := BenchUut11.processMode;
   TraceIn_levelSensor[105] := BenchUut11.levelSensor;
   TraceIn_mixMotorComplete[105] := BenchUut11.mixMotorComplete;
   BenchUut11();
   TraceOut_valveARun[105] := BenchUut11.valveARun;
   TraceOut_valveBRun[105] := BenchUut11.valveBRun;
   TraceOut_valveCRun[105] := BenchUut11.valveCRun;
   TraceOut_valveDRun[105] := BenchUut11.valveDRun;
   TraceOut_mixMotorRun[105] := BenchUut11.mixMotorRun;
   BenchCalls := BenchCalls + 1;
 106:
   BenchUut11.estop := TRUE;
   BenchUut11.opeMode := TRUE;
   BenchUut11.valveAStart := FALSE;
   BenchUut11.valveBStart := FALSE;
   BenchUut11.valveCStart := FALSE;
   BenchUut11.valveDStart := FALSE;
   BenchUut11.mixMotorStart := FALSE;
   BenchUut11.autoStart := FALSE;
   BenchUut11.processMode := FALSE;
   BenchUut11.levelSensor := INT#0;
   BenchUut11.mixMotorComplete := FALSE;
   TraceIn_estop[106] := BenchUut11.estop;
   TraceIn_opeMode[106] := BenchUut11.opeMode;
   TraceIn_valveAStart[106] := BenchUut11.valveAStart;
   TraceIn_valveBStart[106] := BenchUut11.valveBStart;
   TraceIn_valveCStart[106] := BenchUut11.valveCStart;
   TraceIn_valveDStart[106] := BenchUut11.valveDStart;
   TraceIn_mixMotorStart[106] := BenchUut11.mixMotorStart;
   TraceIn_autoStart[106] := BenchUut11.autoStart;
   TraceIn_processMode[106] := BenchUut11.processMode;
   TraceIn_levelSensor[106] := BenchUut11.levelSensor;
   TraceIn_mixMotorComplete[106] := BenchUut11.mixMotorComplete;
   BenchUut11();
   TraceOut_valveARun[106] := BenchUut11.valveARun;
   TraceOut_valveBRun[106] := BenchUut11.valveBRun;
   TraceOut_valveCRun[106] := BenchUut11.valveCRun;
   TraceOut_valveDRun[106] := BenchUut11.valveDRun;
   TraceOut_mixMotorRun[106] := BenchUut11.mixMotorRun;
   BenchCalls := BenchCalls + 1;
 107:
   BenchUut11.estop := TRUE;
   BenchUut11.opeMode := TRUE;
   BenchUut11.valveAStart := FALSE;
   BenchUut11.valveBStart := FALSE;
   BenchUut11.valveCStart := FALSE;
   BenchUut11.valveDStart := FALSE;
   BenchUut11.mixMotorStart := FALSE;
   BenchUut11.autoStart := TRUE;
   BenchUut11.processMode := FALSE;
   BenchUut11.levelSensor := INT#0;
   BenchUut11.mixMotorComplete := FALSE;
   TraceIn_estop[107] := BenchUut11.estop;
   TraceIn_opeMode[107] := BenchUut11.opeMode;
   TraceIn_valveAStart[107] := BenchUut11.valveAStart;
   TraceIn_valveBStart[107] := BenchUut11.valveBStart;
   TraceIn_valveCStart[107] := BenchUut11.valveCStart;
   TraceIn_valveDStart[107] := BenchUut11.valveDStart;
   TraceIn_mixMotorStart[107] := BenchUut11.mixMotorStart;
   TraceIn_autoStart[107] := BenchUut11.autoStart;
   TraceIn_processMode[107] := BenchUut11.processMode;
   TraceIn_levelSensor[107] := BenchUut11.levelSensor;
   TraceIn_mixMotorComplete[107] := BenchUut11.mixMotorComplete;
   BenchUut11();
   TraceOut_valveARun[107] := BenchUut11.valveARun;
   TraceOut_valveBRun[107] := BenchUut11.valveBRun;
   TraceOut_valveCRun[107] := BenchUut11.valveCRun;
   TraceOut_valveDRun[107] := BenchUut11.valveDRun;
   TraceOut_mixMotorRun[107] := BenchUut11.mixMotorRun;
   BenchCalls := BenchCalls + 1;
 108:
   BenchUut11.estop := TRUE;
   BenchUut11.opeMode := TRUE;
   BenchUut11.valveAStart := FALSE;
   BenchUut11.valveBStart := FALSE;
   BenchUut11.valveCStart := FALSE;
   BenchUut11.valveDStart := FALSE;
   BenchUut11.mixMotorStart := FALSE;
   BenchUut11.autoStart := FALSE;
   BenchUut11.processMode := FALSE;
   BenchUut11.levelSensor := INT#0;
   BenchUut11.mixMotorComplete := FALSE;
   TraceIn_estop[108] := BenchUut11.estop;
   TraceIn_opeMode[108] := BenchUut11.opeMode;
   TraceIn_valveAStart[108] := BenchUut11.valveAStart;
   TraceIn_valveBStart[108] := BenchUut11.valveBStart;
   TraceIn_valveCStart[108] := BenchUut11.valveCStart;
   TraceIn_valveDStart[108] := BenchUut11.valveDStart;
   TraceIn_mixMotorStart[108] := BenchUut11.mixMotorStart;
   TraceIn_autoStart[108] := BenchUut11.autoStart;
   TraceIn_processMode[108] := BenchUut11.processMode;
   TraceIn_levelSensor[108] := BenchUut11.levelSensor;
   TraceIn_mixMotorComplete[108] := BenchUut11.mixMotorComplete;
   BenchUut11();
   TraceOut_valveARun[108] := BenchUut11.valveARun;
   TraceOut_valveBRun[108] := BenchUut11.valveBRun;
   TraceOut_valveCRun[108] := BenchUut11.valveCRun;
   TraceOut_valveDRun[108] := BenchUut11.valveDRun;
   TraceOut_mixMotorRun[108] := BenchUut11.mixMotorRun;
   BenchCalls := BenchCalls + 1;
 109:
   BenchUut12.estop := TRUE;
   BenchUut12.opeMode := TRUE;
   BenchUut12.valveAStart := FALSE;
   BenchUut12.valveBStart := FALSE;
   BenchUut12.valveCStart := FALSE;
   BenchUut12.valveDStart := FALSE;
   BenchUut12.mixMotorStart := FALSE;
   BenchUut12.autoStart := FALSE;
   BenchUut12.processMode := TRUE;
   BenchUut12.levelSensor := INT#0;
   BenchUut12.mixMotorComplete := FALSE;
   TraceIn_estop[109] := BenchUut12.estop;
   TraceIn_opeMode[109] := BenchUut12.opeMode;
   TraceIn_valveAStart[109] := BenchUut12.valveAStart;
   TraceIn_valveBStart[109] := BenchUut12.valveBStart;
   TraceIn_valveCStart[109] := BenchUut12.valveCStart;
   TraceIn_valveDStart[109] := BenchUut12.valveDStart;
   TraceIn_mixMotorStart[109] := BenchUut12.mixMotorStart;
   TraceIn_autoStart[109] := BenchUut12.autoStart;
   TraceIn_processMode[109] := BenchUut12.processMode;
   TraceIn_levelSensor[109] := BenchUut12.levelSensor;
   TraceIn_mixMotorComplete[109] := BenchUut12.mixMotorComplete;
   BenchUut12();
   TraceOut_valveARun[109] := BenchUut12.valveARun;
   TraceOut_valveBRun[109] := BenchUut12.valveBRun;
   TraceOut_valveCRun[109] := BenchUut12.valveCRun;
   TraceOut_valveDRun[109] := BenchUut12.valveDRun;
   TraceOut_mixMotorRun[109] := BenchUut12.mixMotorRun;
   BenchCalls := BenchCalls + 1;
 110:
   BenchUut12.estop := TRUE;
   BenchUut12.opeMode := TRUE;
   BenchUut12.valveAStart := FALSE;
   BenchUut12.valveBStart := FALSE;
   BenchUut12.valveCStart := FALSE;
   BenchUut12.valveDStart := FALSE;
   BenchUut12.mixMotorStart := FALSE;
   BenchUut12.autoStart := TRUE;
   BenchUut12.processMode := TRUE;
   BenchUut12.levelSensor := INT#0;
   BenchUut12.mixMotorComplete := FALSE;
   TraceIn_estop[110] := BenchUut12.estop;
   TraceIn_opeMode[110] := BenchUut12.opeMode;
   TraceIn_valveAStart[110] := BenchUut12.valveAStart;
   TraceIn_valveBStart[110] := BenchUut12.valveBStart;
   TraceIn_valveCStart[110] := BenchUut12.valveCStart;
   TraceIn_valveDStart[110] := BenchUut12.valveDStart;
   TraceIn_mixMotorStart[110] := BenchUut12.mixMotorStart;
   TraceIn_autoStart[110] := BenchUut12.autoStart;
   TraceIn_processMode[110] := BenchUut12.processMode;
   TraceIn_levelSensor[110] := BenchUut12.levelSensor;
   TraceIn_mixMotorComplete[110] := BenchUut12.mixMotorComplete;
   BenchUut12();
   TraceOut_valveARun[110] := BenchUut12.valveARun;
   TraceOut_valveBRun[110] := BenchUut12.valveBRun;
   TraceOut_valveCRun[110] := BenchUut12.valveCRun;
   TraceOut_valveDRun[110] := BenchUut12.valveDRun;
   TraceOut_mixMotorRun[110] := BenchUut12.mixMotorRun;
   BenchCalls := BenchCalls + 1;
 111:
   BenchUut12.estop := TRUE;
   BenchUut12.opeMode := TRUE;
   BenchUut12.valveAStart := FALSE;
   BenchUut12.valveBStart := FALSE;
   BenchUut12.valveCStart := FALSE;
   BenchUut12.valveDStart := FALSE;
   BenchUut12.mixMotorStart := FALSE;
   BenchUut12.autoStart := FALSE;
   BenchUut12.processMode := TRUE;
   BenchUut12.levelSensor := INT#0;
   BenchUut12.mixMotorComplete := FALSE;
   TraceIn_estop[111] := BenchUut12.estop;
   TraceIn_opeMode[111] := BenchUut12.opeMode;
   TraceIn_valveAStart[111] := BenchUut12.valveAStart;
   TraceIn_valveBStart[111] := BenchUut12.valveBStart;
   TraceIn_valveCStart[111] := BenchUut12.valveCStart;
   TraceIn_valveDStart[111] := BenchUut12.valveDStart;
   TraceIn_mixMotorStart[111] := BenchUut12.mixMotorStart;
   TraceIn_autoStart[111] := BenchUut12.autoStart;
   TraceIn_processMode[111] := BenchUut12.processMode;
   TraceIn_levelSensor[111] := BenchUut12.levelSensor;
   TraceIn_mixMotorComplete[111] := BenchUut12.mixMotorComplete;
   BenchUut12();
   TraceOut_valveARun[111] := BenchUut12.valveARun;
   TraceOut_valveBRun[111] := BenchUut12.valveBRun;
   TraceOut_valveCRun[111] := BenchUut12.valveCRun;
   TraceOut_valveDRun[111] := BenchUut12.valveDRun;
   TraceOut_mixMotorRun[111] := BenchUut12.mixMotorRun;
   BenchCalls := BenchCalls + 1;
 112:
   BenchUut12.estop := TRUE;
   BenchUut12.opeMode := TRUE;
   BenchUut12.valveAStart := FALSE;
   BenchUut12.valveBStart := FALSE;
   BenchUut12.valveCStart := FALSE;
   BenchUut12.valveDStart := FALSE;
   BenchUut12.mixMotorStart := FALSE;
   BenchUut12.autoStart := FALSE;
   BenchUut12.processMode := TRUE;
   BenchUut12.levelSensor := INT#0;
   BenchUut12.mixMotorComplete := FALSE;
   TraceIn_estop[112] := BenchUut12.estop;
   TraceIn_opeMode[112] := BenchUut12.opeMode;
   TraceIn_valveAStart[112] := BenchUut12.valveAStart;
   TraceIn_valveBStart[112] := BenchUut12.valveBStart;
   TraceIn_valveCStart[112] := BenchUut12.valveCStart;
   TraceIn_valveDStart[112] := BenchUut12.valveDStart;
   TraceIn_mixMotorStart[112] := BenchUut12.mixMotorStart;
   TraceIn_autoStart[112] := BenchUut12.autoStart;
   TraceIn_processMode[112] := BenchUut12.processMode;
   TraceIn_levelSensor[112] := BenchUut12.levelSensor;
   TraceIn_mixMotorComplete[112] := BenchUut12.mixMotorComplete;
   BenchUut12();
   TraceOut_valveARun[112] := BenchUut12.valveARun;
   TraceOut_valveBRun[112] := BenchUut12.valveBRun;
   TraceOut_valveCRun[112] := BenchUut12.valveCRun;
   TraceOut_valveDRun[112] := BenchUut12.valveDRun;
   TraceOut_mixMotorRun[112] := BenchUut12.mixMotorRun;
   BenchCalls := BenchCalls + 1;
 113:
   BenchUut12.estop := TRUE;
   BenchUut12.opeMode := TRUE;
   BenchUut12.valveAStart := FALSE;
   BenchUut12.valveBStart := FALSE;
   BenchUut12.valveCStart := FALSE;
   BenchUut12.valveDStart := FALSE;
   BenchUut12.mixMotorStart := FALSE;
   BenchUut12.autoStart := FALSE;
   BenchUut12.processMode := TRUE;
   BenchUut12.levelSensor := INT#50;
   BenchUut12.mixMotorComplete := FALSE;
   TraceIn_estop[113] := BenchUut12.estop;
   TraceIn_opeMode[113] := BenchUut12.opeMode;
   TraceIn_valveAStart[113] := BenchUut12.valveAStart;
   TraceIn_valveBStart[113] := BenchUut12.valveBStart;
   TraceIn_valveCStart[113] := BenchUut12.valveCStart;
   TraceIn_valveDStart[113] := BenchUut12.valveDStart;
   TraceIn_mixMotorStart[113] := BenchUut12.mixMotorStart;
   TraceIn_autoStart[113] := BenchUut12.autoStart;
   TraceIn_processMode[113] := BenchUut12.processMode;
   TraceIn_levelSensor[113] := BenchUut12.levelSensor;
   TraceIn_mixMotorComplete[113] := BenchUut12.mixMotorComplete;
   BenchUut12();
   TraceOut_valveARun[113] := BenchUut12.valveARun;
   TraceOut_valveBRun[113] := BenchUut12.valveBRun;
   TraceOut_valveCRun[113] := BenchUut12.valveCRun;
   TraceOut_valveDRun[113] := BenchUut12.valveDRun;
   TraceOut_mixMotorRun[113] := BenchUut12.mixMotorRun;
   BenchCalls := BenchCalls + 1;
 114:
   BenchUut12.estop := TRUE;
   BenchUut12.opeMode := TRUE;
   BenchUut12.valveAStart := FALSE;
   BenchUut12.valveBStart := FALSE;
   BenchUut12.valveCStart := FALSE;
   BenchUut12.valveDStart := FALSE;
   BenchUut12.mixMotorStart := FALSE;
   BenchUut12.autoStart := FALSE;
   BenchUut12.processMode := TRUE;
   BenchUut12.levelSensor := INT#50;
   BenchUut12.mixMotorComplete := FALSE;
   TraceIn_estop[114] := BenchUut12.estop;
   TraceIn_opeMode[114] := BenchUut12.opeMode;
   TraceIn_valveAStart[114] := BenchUut12.valveAStart;
   TraceIn_valveBStart[114] := BenchUut12.valveBStart;
   TraceIn_valveCStart[114] := BenchUut12.valveCStart;
   TraceIn_valveDStart[114] := BenchUut12.valveDStart;
   TraceIn_mixMotorStart[114] := BenchUut12.mixMotorStart;
   TraceIn_autoStart[114] := BenchUut12.autoStart;
   TraceIn_processMode[114] := BenchUut12.processMode;
   TraceIn_levelSensor[114] := BenchUut12.levelSensor;
   TraceIn_mixMotorComplete[114] := BenchUut12.mixMotorComplete;
   BenchUut12();
   TraceOut_valveARun[114] := BenchUut12.valveARun;
   TraceOut_valveBRun[114] := BenchUut12.valveBRun;
   TraceOut_valveCRun[114] := BenchUut12.valveCRun;
   TraceOut_valveDRun[114] := BenchUut12.valveDRun;
   TraceOut_mixMotorRun[114] := BenchUut12.mixMotorRun;
   BenchCalls := BenchCalls + 1;
 115:
   BenchUut12.estop := TRUE;
   BenchUut12.opeMode := TRUE;
   BenchUut12.valveAStart := FALSE;
   BenchUut12.valveBStart := FALSE;
   BenchUut12.valveCStart := FALSE;
   BenchUut12.valveDStart := FALSE;
   BenchUut12.mixMotorStart := FALSE;
   BenchUut12.autoStart := FALSE;
   BenchUut12.processMode := TRUE;
   BenchUut12.levelSensor := INT#80;
   BenchUut12.mixMotorComplete := FALSE;
   TraceIn_estop[115] := BenchUut12.estop;
   TraceIn_opeMode[115] := BenchUut12.opeMode;
   TraceIn_valveAStart[115] := BenchUut12.valveAStart;
   TraceIn_valveBStart[115] := BenchUut12.valveBStart;
   TraceIn_valveCStart[115] := BenchUut12.valveCStart;
   TraceIn_valveDStart[115] := BenchUut12.valveDStart;
   TraceIn_mixMotorStart[115] := BenchUut12.mixMotorStart;
   TraceIn_autoStart[115] := BenchUut12.autoStart;
   TraceIn_processMode[115] := BenchUut12.processMode;
   TraceIn_levelSensor[115] := BenchUut12.levelSensor;
   TraceIn_mixMotorComplete[115] := BenchUut12.mixMotorComplete;
   BenchUut12();
   TraceOut_valveARun[115] := BenchUut12.valveARun;
   TraceOut_valveBRun[115] := BenchUut12.valveBRun;
   TraceOut_valveCRun[115] := BenchUut12.valveCRun;
   TraceOut_valveDRun[115] := BenchUut12.valveDRun;
   TraceOut_mixMotorRun[115] := BenchUut12.mixMotorRun;
   BenchCalls := BenchCalls + 1;
 116:
   BenchUut12.estop := TRUE;
   BenchUut12.opeMode := TRUE;
   BenchUut12.valveAStart := FALSE;
   BenchUut12.valveBStart := FALSE;
   BenchUut12.valveCStart := FALSE;
   BenchUut12.valveDStart := FALSE;
   BenchUut12.mixMotorStart := FALSE;
   BenchUut12.autoStart := FALSE;
   BenchUut12.processMode := TRUE;
   BenchUut12.levelSensor := INT#80;
   BenchUut12.mixMotorComplete := FALSE;
   TraceIn_estop[116] := BenchUut12.estop;
   TraceIn_opeMode[116] := BenchUut12.opeMode;
   TraceIn_valveAStart[116] := BenchUut12.valveAStart;
   TraceIn_valveBStart[116] := BenchUut12.valveBStart;
   TraceIn_valveCStart[116] := BenchUut12.valveCStart;
   TraceIn_valveDStart[116] := BenchUut12.valveDStart;
   TraceIn_mixMotorStart[116] := BenchUut12.mixMotorStart;
   TraceIn_autoStart[116] := BenchUut12.autoStart;
   TraceIn_processMode[116] := BenchUut12.processMode;
   TraceIn_levelSensor[116] := BenchUut12.levelSensor;
   TraceIn_mixMotorComplete[116] := BenchUut12.mixMotorComplete;
   BenchUut12();
   TraceOut_valveARun[116] := BenchUut12.valveARun;
   TraceOut_valveBRun[116] := BenchUut12.valveBRun;
   TraceOut_valveCRun[116] := BenchUut12.valveCRun;
   TraceOut_valveDRun[116] := BenchUut12.valveDRun;
   TraceOut_mixMotorRun[116] := BenchUut12.mixMotorRun;
   BenchCalls := BenchCalls + 1;
 117:
   BenchUut12.estop := TRUE;
   BenchUut12.opeMode := TRUE;
   BenchUut12.valveAStart := FALSE;
   BenchUut12.valveBStart := FALSE;
   BenchUut12.valveCStart := FALSE;
   BenchUut12.valveDStart := FALSE;
   BenchUut12.mixMotorStart := FALSE;
   BenchUut12.autoStart := FALSE;
   BenchUut12.processMode := TRUE;
   BenchUut12.levelSensor := INT#100;
   BenchUut12.mixMotorComplete := FALSE;
   TraceIn_estop[117] := BenchUut12.estop;
   TraceIn_opeMode[117] := BenchUut12.opeMode;
   TraceIn_valveAStart[117] := BenchUut12.valveAStart;
   TraceIn_valveBStart[117] := BenchUut12.valveBStart;
   TraceIn_valveCStart[117] := BenchUut12.valveCStart;
   TraceIn_valveDStart[117] := BenchUut12.valveDStart;
   TraceIn_mixMotorStart[117] := BenchUut12.mixMotorStart;
   TraceIn_autoStart[117] := BenchUut12.autoStart;
   TraceIn_processMode[117] := BenchUut12.processMode;
   TraceIn_levelSensor[117] := BenchUut12.levelSensor;
   TraceIn_mixMotorComplete[117] := BenchUut12.mixMotorComplete;
   BenchUut12();
   TraceOut_valveARun[117] := BenchUut12.valveARun;
   TraceOut_valveBRun[117] := BenchUut12.valveBRun;
   TraceOut_valveCRun[117] := BenchUut12.valveCRun;
   TraceOut_valveDRun[117] := BenchUut12.valveDRun;
   TraceOut_mixMotorRun[117] := BenchUut12.mixMotorRun;
   BenchCalls := BenchCalls + 1;
 118:
   BenchUut12.estop := TRUE;
   BenchUut12.opeMode := TRUE;
   BenchUut12.valveAStart := FALSE;
   BenchUut12.valveBStart := FALSE;
   BenchUut12.valveCStart := FALSE;
   BenchUut12.valveDStart := FALSE;
   BenchUut12.mixMotorStart := FALSE;
   BenchUut12.autoStart := FALSE;
   BenchUut12.processMode := TRUE;
   BenchUut12.levelSensor := INT#100;
   BenchUut12.mixMotorComplete := FALSE;
   TraceIn_estop[118] := BenchUut12.estop;
   TraceIn_opeMode[118] := BenchUut12.opeMode;
   TraceIn_valveAStart[118] := BenchUut12.valveAStart;
   TraceIn_valveBStart[118] := BenchUut12.valveBStart;
   TraceIn_valveCStart[118] := BenchUut12.valveCStart;
   TraceIn_valveDStart[118] := BenchUut12.valveDStart;
   TraceIn_mixMotorStart[118] := BenchUut12.mixMotorStart;
   TraceIn_autoStart[118] := BenchUut12.autoStart;
   TraceIn_processMode[118] := BenchUut12.processMode;
   TraceIn_levelSensor[118] := BenchUut12.levelSensor;
   TraceIn_mixMotorComplete[118] := BenchUut12.mixMotorComplete;
   BenchUut12();
   TraceOut_valveARun[118] := BenchUut12.valveARun;
   TraceOut_valveBRun[118] := BenchUut12.valveBRun;
   TraceOut_valveCRun[118] := BenchUut12.valveCRun;
   TraceOut_valveDRun[118] := BenchUut12.valveDRun;
   TraceOut_mixMotorRun[118] := BenchUut12.mixMotorRun;
   BenchCalls := BenchCalls + 1;
 119:
   BenchUut12.estop := TRUE;
   BenchUut12.opeMode := TRUE;
   BenchUut12.valveAStart := FALSE;
   BenchUut12.valveBStart := FALSE;
   BenchUut12.valveCStart := FALSE;
   BenchUut12.valveDStart := FALSE;
   BenchUut12.mixMotorStart := FALSE;
   BenchUut12.autoStart := FALSE;
   BenchUut12.processMode := TRUE;
   BenchUut12.levelSensor := INT#100;
   BenchUut12.mixMotorComplete := FALSE;
   TraceIn_estop[119] := BenchUut12.estop;
   TraceIn_opeMode[119] := BenchUut12.opeMode;
   TraceIn_valveAStart[119] := BenchUut12.valveAStart;
   TraceIn_valveBStart[119] := BenchUut12.valveBStart;
   TraceIn_valveCStart[119] := BenchUut12.valveCStart;
   TraceIn_valveDStart[119] := BenchUut12.valveDStart;
   TraceIn_mixMotorStart[119] := BenchUut12.mixMotorStart;
   TraceIn_autoStart[119] := BenchUut12.autoStart;
   TraceIn_processMode[119] := BenchUut12.processMode;
   TraceIn_levelSensor[119] := BenchUut12.levelSensor;
   TraceIn_mixMotorComplete[119] := BenchUut12.mixMotorComplete;
   BenchUut12();
   TraceOut_valveARun[119] := BenchUut12.valveARun;
   TraceOut_valveBRun[119] := BenchUut12.valveBRun;
   TraceOut_valveCRun[119] := BenchUut12.valveCRun;
   TraceOut_valveDRun[119] := BenchUut12.valveDRun;
   TraceOut_mixMotorRun[119] := BenchUut12.mixMotorRun;
   BenchCalls := BenchCalls + 1;
 120:
   BenchUut12.estop := TRUE;
   BenchUut12.opeMode := TRUE;
   BenchUut12.valveAStart := FALSE;
   BenchUut12.valveBStart := FALSE;
   BenchUut12.valveCStart := FALSE;
   BenchUut12.valveDStart := FALSE;
   BenchUut12.mixMotorStart := FALSE;
   BenchUut12.autoStart := FALSE;
   BenchUut12.processMode := TRUE;
   BenchUut12.levelSensor := INT#100;
   BenchUut12.mixMotorComplete := TRUE;
   TraceIn_estop[120] := BenchUut12.estop;
   TraceIn_opeMode[120] := BenchUut12.opeMode;
   TraceIn_valveAStart[120] := BenchUut12.valveAStart;
   TraceIn_valveBStart[120] := BenchUut12.valveBStart;
   TraceIn_valveCStart[120] := BenchUut12.valveCStart;
   TraceIn_valveDStart[120] := BenchUut12.valveDStart;
   TraceIn_mixMotorStart[120] := BenchUut12.mixMotorStart;
   TraceIn_autoStart[120] := BenchUut12.autoStart;
   TraceIn_processMode[120] := BenchUut12.processMode;
   TraceIn_levelSensor[120] := BenchUut12.levelSensor;
   TraceIn_mixMotorComplete[120] := BenchUut12.mixMotorComplete;
   BenchUut12();
   TraceOut_valveARun[120] := BenchUut12.valveARun;
   TraceOut_valveBRun[120] := BenchUut12.valveBRun;
   TraceOut_valveCRun[120] := BenchUut12.valveCRun;
   TraceOut_valveDRun[120] := BenchUut12.valveDRun;
   TraceOut_mixMotorRun[120] := BenchUut12.mixMotorRun;
   BenchCalls := BenchCalls + 1;
 121:
   BenchUut12.estop := TRUE;
   BenchUut12.opeMode := TRUE;
   BenchUut12.valveAStart := FALSE;
   BenchUut12.valveBStart := FALSE;
   BenchUut12.valveCStart := FALSE;
   BenchUut12.valveDStart := FALSE;
   BenchUut12.mixMotorStart := FALSE;
   BenchUut12.autoStart := FALSE;
   BenchUut12.processMode := TRUE;
   BenchUut12.levelSensor := INT#100;
   BenchUut12.mixMotorComplete := FALSE;
   TraceIn_estop[121] := BenchUut12.estop;
   TraceIn_opeMode[121] := BenchUut12.opeMode;
   TraceIn_valveAStart[121] := BenchUut12.valveAStart;
   TraceIn_valveBStart[121] := BenchUut12.valveBStart;
   TraceIn_valveCStart[121] := BenchUut12.valveCStart;
   TraceIn_valveDStart[121] := BenchUut12.valveDStart;
   TraceIn_mixMotorStart[121] := BenchUut12.mixMotorStart;
   TraceIn_autoStart[121] := BenchUut12.autoStart;
   TraceIn_processMode[121] := BenchUut12.processMode;
   TraceIn_levelSensor[121] := BenchUut12.levelSensor;
   TraceIn_mixMotorComplete[121] := BenchUut12.mixMotorComplete;
   BenchUut12();
   TraceOut_valveARun[121] := BenchUut12.valveARun;
   TraceOut_valveBRun[121] := BenchUut12.valveBRun;
   TraceOut_valveCRun[121] := BenchUut12.valveCRun;
   TraceOut_valveDRun[121] := BenchUut12.valveDRun;
   TraceOut_mixMotorRun[121] := BenchUut12.mixMotorRun;
   BenchCalls := BenchCalls + 1;
 122:
   BenchUut12.estop := TRUE;
   BenchUut12.opeMode := TRUE;
   BenchUut12.valveAStart := FALSE;
   BenchUut12.valveBStart := FALSE;
   BenchUut12.valveCStart := FALSE;
   BenchUut12.valveDStart := FALSE;
   BenchUut12.mixMotorStart := FALSE;
   BenchUut12.autoStart := FALSE;
   BenchUut12.processMode := TRUE;
   BenchUut12.levelSensor := INT#100;
   BenchUut12.mixMotorComplete := FALSE;
   TraceIn_estop[122] := BenchUut12.estop;
   TraceIn_opeMode[122] := BenchUut12.opeMode;
   TraceIn_valveAStart[122] := BenchUut12.valveAStart;
   TraceIn_valveBStart[122] := BenchUut12.valveBStart;
   TraceIn_valveCStart[122] := BenchUut12.valveCStart;
   TraceIn_valveDStart[122] := BenchUut12.valveDStart;
   TraceIn_mixMotorStart[122] := BenchUut12.mixMotorStart;
   TraceIn_autoStart[122] := BenchUut12.autoStart;
   TraceIn_processMode[122] := BenchUut12.processMode;
   TraceIn_levelSensor[122] := BenchUut12.levelSensor;
   TraceIn_mixMotorComplete[122] := BenchUut12.mixMotorComplete;
   BenchUut12();
   TraceOut_valveARun[122] := BenchUut12.valveARun;
   TraceOut_valveBRun[122] := BenchUut12.valveBRun;
   TraceOut_valveCRun[122] := BenchUut12.valveCRun;
   TraceOut_valveDRun[122] := BenchUut12.valveDRun;
   TraceOut_mixMotorRun[122] := BenchUut12.mixMotorRun;
   BenchCalls := BenchCalls + 1;
 123:
   BenchUut12.estop := TRUE;
   BenchUut12.opeMode := FALSE;
   BenchUut12.valveAStart := FALSE;
   BenchUut12.valveBStart := FALSE;
   BenchUut12.valveCStart := FALSE;
   BenchUut12.valveDStart := FALSE;
   BenchUut12.mixMotorStart := FALSE;
   BenchUut12.autoStart := FALSE;
   BenchUut12.processMode := TRUE;
   BenchUut12.levelSensor := INT#100;
   BenchUut12.mixMotorComplete := FALSE;
   TraceIn_estop[123] := BenchUut12.estop;
   TraceIn_opeMode[123] := BenchUut12.opeMode;
   TraceIn_valveAStart[123] := BenchUut12.valveAStart;
   TraceIn_valveBStart[123] := BenchUut12.valveBStart;
   TraceIn_valveCStart[123] := BenchUut12.valveCStart;
   TraceIn_valveDStart[123] := BenchUut12.valveDStart;
   TraceIn_mixMotorStart[123] := BenchUut12.mixMotorStart;
   TraceIn_autoStart[123] := BenchUut12.autoStart;
   TraceIn_processMode[123] := BenchUut12.processMode;
   TraceIn_levelSensor[123] := BenchUut12.levelSensor;
   TraceIn_mixMotorComplete[123] := BenchUut12.mixMotorComplete;
   BenchUut12();
   TraceOut_valveARun[123] := BenchUut12.valveARun;
   TraceOut_valveBRun[123] := BenchUut12.valveBRun;
   TraceOut_valveCRun[123] := BenchUut12.valveCRun;
   TraceOut_valveDRun[123] := BenchUut12.valveDRun;
   TraceOut_mixMotorRun[123] := BenchUut12.mixMotorRun;
   BenchCalls := BenchCalls + 1;
 124:
   BenchUut12.estop := TRUE;
   BenchUut12.opeMode := TRUE;
   BenchUut12.valveAStart := FALSE;
   BenchUut12.valveBStart := FALSE;
   BenchUut12.valveCStart := FALSE;
   BenchUut12.valveDStart := FALSE;
   BenchUut12.mixMotorStart := FALSE;
   BenchUut12.autoStart := FALSE;
   BenchUut12.processMode := TRUE;
   BenchUut12.levelSensor := INT#0;
   BenchUut12.mixMotorComplete := FALSE;
   TraceIn_estop[124] := BenchUut12.estop;
   TraceIn_opeMode[124] := BenchUut12.opeMode;
   TraceIn_valveAStart[124] := BenchUut12.valveAStart;
   TraceIn_valveBStart[124] := BenchUut12.valveBStart;
   TraceIn_valveCStart[124] := BenchUut12.valveCStart;
   TraceIn_valveDStart[124] := BenchUut12.valveDStart;
   TraceIn_mixMotorStart[124] := BenchUut12.mixMotorStart;
   TraceIn_autoStart[124] := BenchUut12.autoStart;
   TraceIn_processMode[124] := BenchUut12.processMode;
   TraceIn_levelSensor[124] := BenchUut12.levelSensor;
   TraceIn_mixMotorComplete[124] := BenchUut12.mixMotorComplete;
   BenchUut12();
   TraceOut_valveARun[124] := BenchUut12.valveARun;
   TraceOut_valveBRun[124] := BenchUut12.valveBRun;
   TraceOut_valveCRun[124] := BenchUut12.valveCRun;
   TraceOut_valveDRun[124] := BenchUut12.valveDRun;
   TraceOut_mixMotorRun[124] := BenchUut12.mixMotorRun;
   BenchCalls := BenchCalls + 1;
 125:
   BenchUut12.estop := TRUE;
   BenchUut12.opeMode := TRUE;
   BenchUut12.valveAStart := FALSE;
   BenchUut12.valveBStart := FALSE;
   BenchUut12.valveCStart := FALSE;
   BenchUut12.valveDStart := FALSE;
   BenchUut12.mixMotorStart := FALSE;
   BenchUut12.autoStart := TRUE;
   BenchUut12.processMode := TRUE;
   BenchUut12.levelSensor := INT#0;
   BenchUut12.mixMotorComplete := FALSE;
   TraceIn_estop[125] := BenchUut12.estop;
   TraceIn_opeMode[125] := BenchUut12.opeMode;
   TraceIn_valveAStart[125] := BenchUut12.valveAStart;
   TraceIn_valveBStart[125] := BenchUut12.valveBStart;
   TraceIn_valveCStart[125] := BenchUut12.valveCStart;
   TraceIn_valveDStart[125] := BenchUut12.valveDStart;
   TraceIn_mixMotorStart[125] := BenchUut12.mixMotorStart;
   TraceIn_autoStart[125] := BenchUut12.autoStart;
   TraceIn_processMode[125] := BenchUut12.processMode;
   TraceIn_levelSensor[125] := BenchUut12.levelSensor;
   TraceIn_mixMotorComplete[125] := BenchUut12.mixMotorComplete;
   BenchUut12();
   TraceOut_valveARun[125] := BenchUut12.valveARun;
   TraceOut_valveBRun[125] := BenchUut12.valveBRun;
   TraceOut_valveCRun[125] := BenchUut12.valveCRun;
   TraceOut_valveDRun[125] := BenchUut12.valveDRun;
   TraceOut_mixMotorRun[125] := BenchUut12.mixMotorRun;
   BenchCalls := BenchCalls + 1;
 126:
   BenchUut12.estop := TRUE;
   BenchUut12.opeMode := TRUE;
   BenchUut12.valveAStart := FALSE;
   BenchUut12.valveBStart := FALSE;
   BenchUut12.valveCStart := FALSE;
   BenchUut12.valveDStart := FALSE;
   BenchUut12.mixMotorStart := FALSE;
   BenchUut12.autoStart := FALSE;
   BenchUut12.processMode := TRUE;
   BenchUut12.levelSensor := INT#0;
   BenchUut12.mixMotorComplete := FALSE;
   TraceIn_estop[126] := BenchUut12.estop;
   TraceIn_opeMode[126] := BenchUut12.opeMode;
   TraceIn_valveAStart[126] := BenchUut12.valveAStart;
   TraceIn_valveBStart[126] := BenchUut12.valveBStart;
   TraceIn_valveCStart[126] := BenchUut12.valveCStart;
   TraceIn_valveDStart[126] := BenchUut12.valveDStart;
   TraceIn_mixMotorStart[126] := BenchUut12.mixMotorStart;
   TraceIn_autoStart[126] := BenchUut12.autoStart;
   TraceIn_processMode[126] := BenchUut12.processMode;
   TraceIn_levelSensor[126] := BenchUut12.levelSensor;
   TraceIn_mixMotorComplete[126] := BenchUut12.mixMotorComplete;
   BenchUut12();
   TraceOut_valveARun[126] := BenchUut12.valveARun;
   TraceOut_valveBRun[126] := BenchUut12.valveBRun;
   TraceOut_valveCRun[126] := BenchUut12.valveCRun;
   TraceOut_valveDRun[126] := BenchUut12.valveDRun;
   TraceOut_mixMotorRun[126] := BenchUut12.mixMotorRun;
   BenchCalls := BenchCalls + 1;
 END_CASE;
 BenchStep := BenchStep + 1;
 IF BenchStep >= 127 THEN BenchDone := TRUE; END_IF;
END_IF;
END_PROGRAM
